FUNCTION_BLOCK FB_Gr05AutoProcedure
(*

The function block used to generate auto process..

Constructor: 		Patryk Panylo
Company:		E. Riexinger GmbH
Date:			28.04.2015
Version:			1.00

Date:			Revision:		Who:				Comment
dd.mm.yyyy		x.xx			Initials			comment

*)
VAR_INPUT
	(* Input variables / Eingang Variablen *)
	bEnable						:BOOL;						(* Enable FB signal *)
	bExecute					:BOOL;						(* Auto procedure execute *)
	bReleaseNextStep			:BOOL;						(* Auto procedure release next step *)
	bInterrupt					:BOOL;						(* Auto procedure interrupt *)
	SFCInit						:BOOL; 						(* System Flag:: INIT Flag *)
	bFirstTime					:BOOL;
END_VAR
VAR_OUTPUT
	(* Output variables / Ausgang Variablen *)
	bDone						:BOOL;						(* Program done *)
	bInterrupted					:BOOL;						(* Program interrupted *)
	bBusy						:BOOL;						(* Program busy *)
	bError						:BOOL;						(* Program error *)
	udnErrorNo					:UDINT;						(* Error number *)
	SFCError						:BOOL; 						(* System Flag: Timeout in this step *)
END_VAR
VAR_IN_OUT
	(* Input Output variables / Ausgang Variablen *)

END_VAR
VAR
	(* Enummerations *)

	(* Variables *)
	lrClamp1Pos					:LREAL;
	lrClamp1PosCache			:LREAL;
	lrClamp1PosPipeEnd			:LREAL;
	lrClamp2Pos					:LREAL;
	lrActRemoveLength			:LREAL;
	bPipeEndDetected			:BOOL;
	unProcessCounter				:UINT;
	lrActSawingLength				:LREAL;
	lrActSawingAngle				:LREAL;

	lrDistPipeBeginSawBand		:LREAL;

	bSafetyDistEnable			:BOOL; 						(* Safety distance between Clamp1 & 2 increase *)
	bErrorPipeBeginNoDetected	:BOOL;						(* Pipe begin no detected *)
	bErrorPipeEndNoDetected		:BOOL;						(* Pipe end no detected *)
	bErrorCollisionDetected		:BOOL;						(* Collision detected *)
	bWarningPipeBeginNoDetected	:BOOL;						(* Pipe begin no detected *)

	SFCCurrentStep				:STRING;					(* Name des aktiven Schritts *)

	(* References *)

	(* Interfaces *)

	(* Instances *)
	rtPipeBeginIdentify			:R_TRIG;
	rtPipeEndIdentify				:R_TRIG;
END_VAR

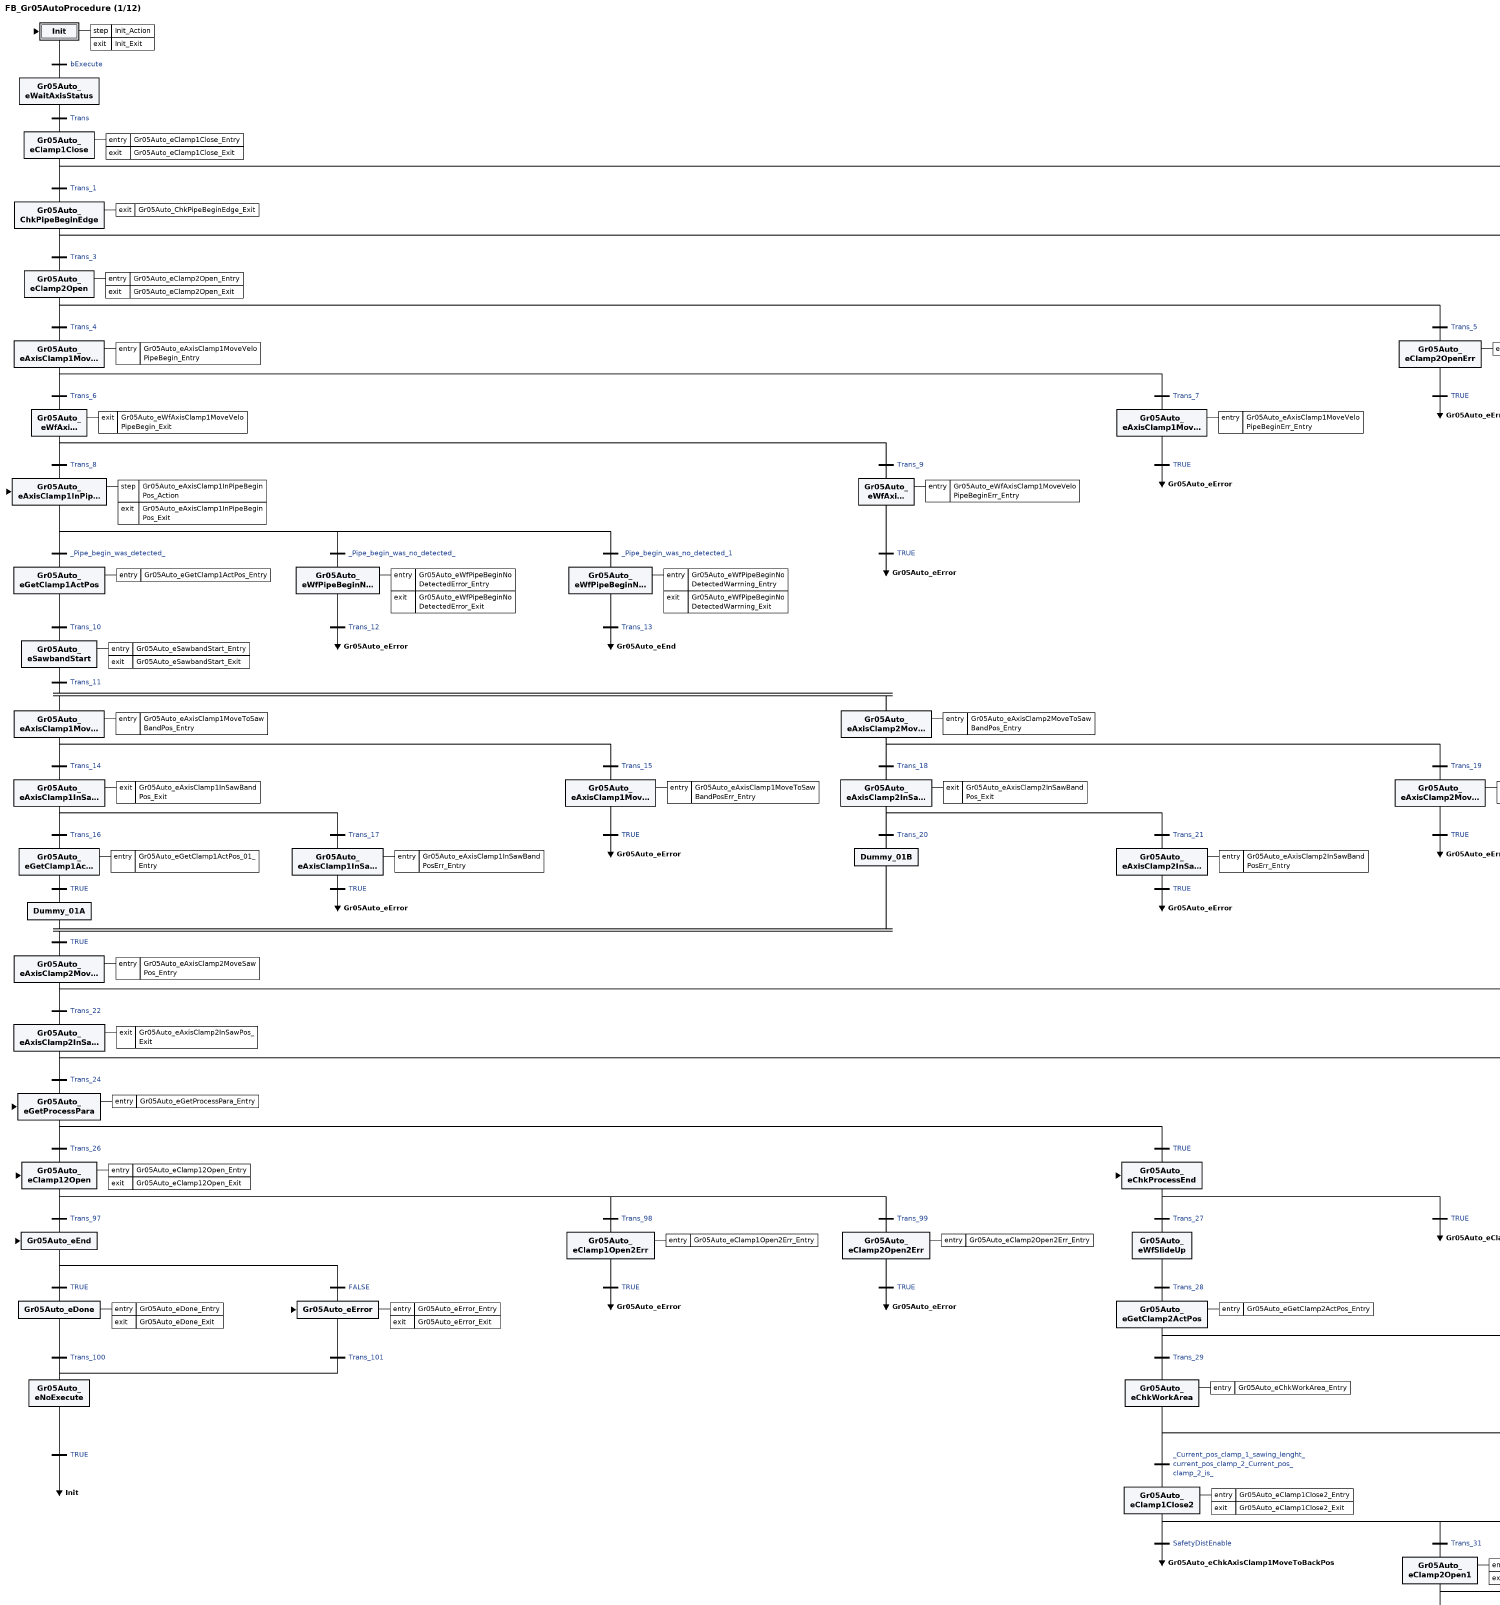
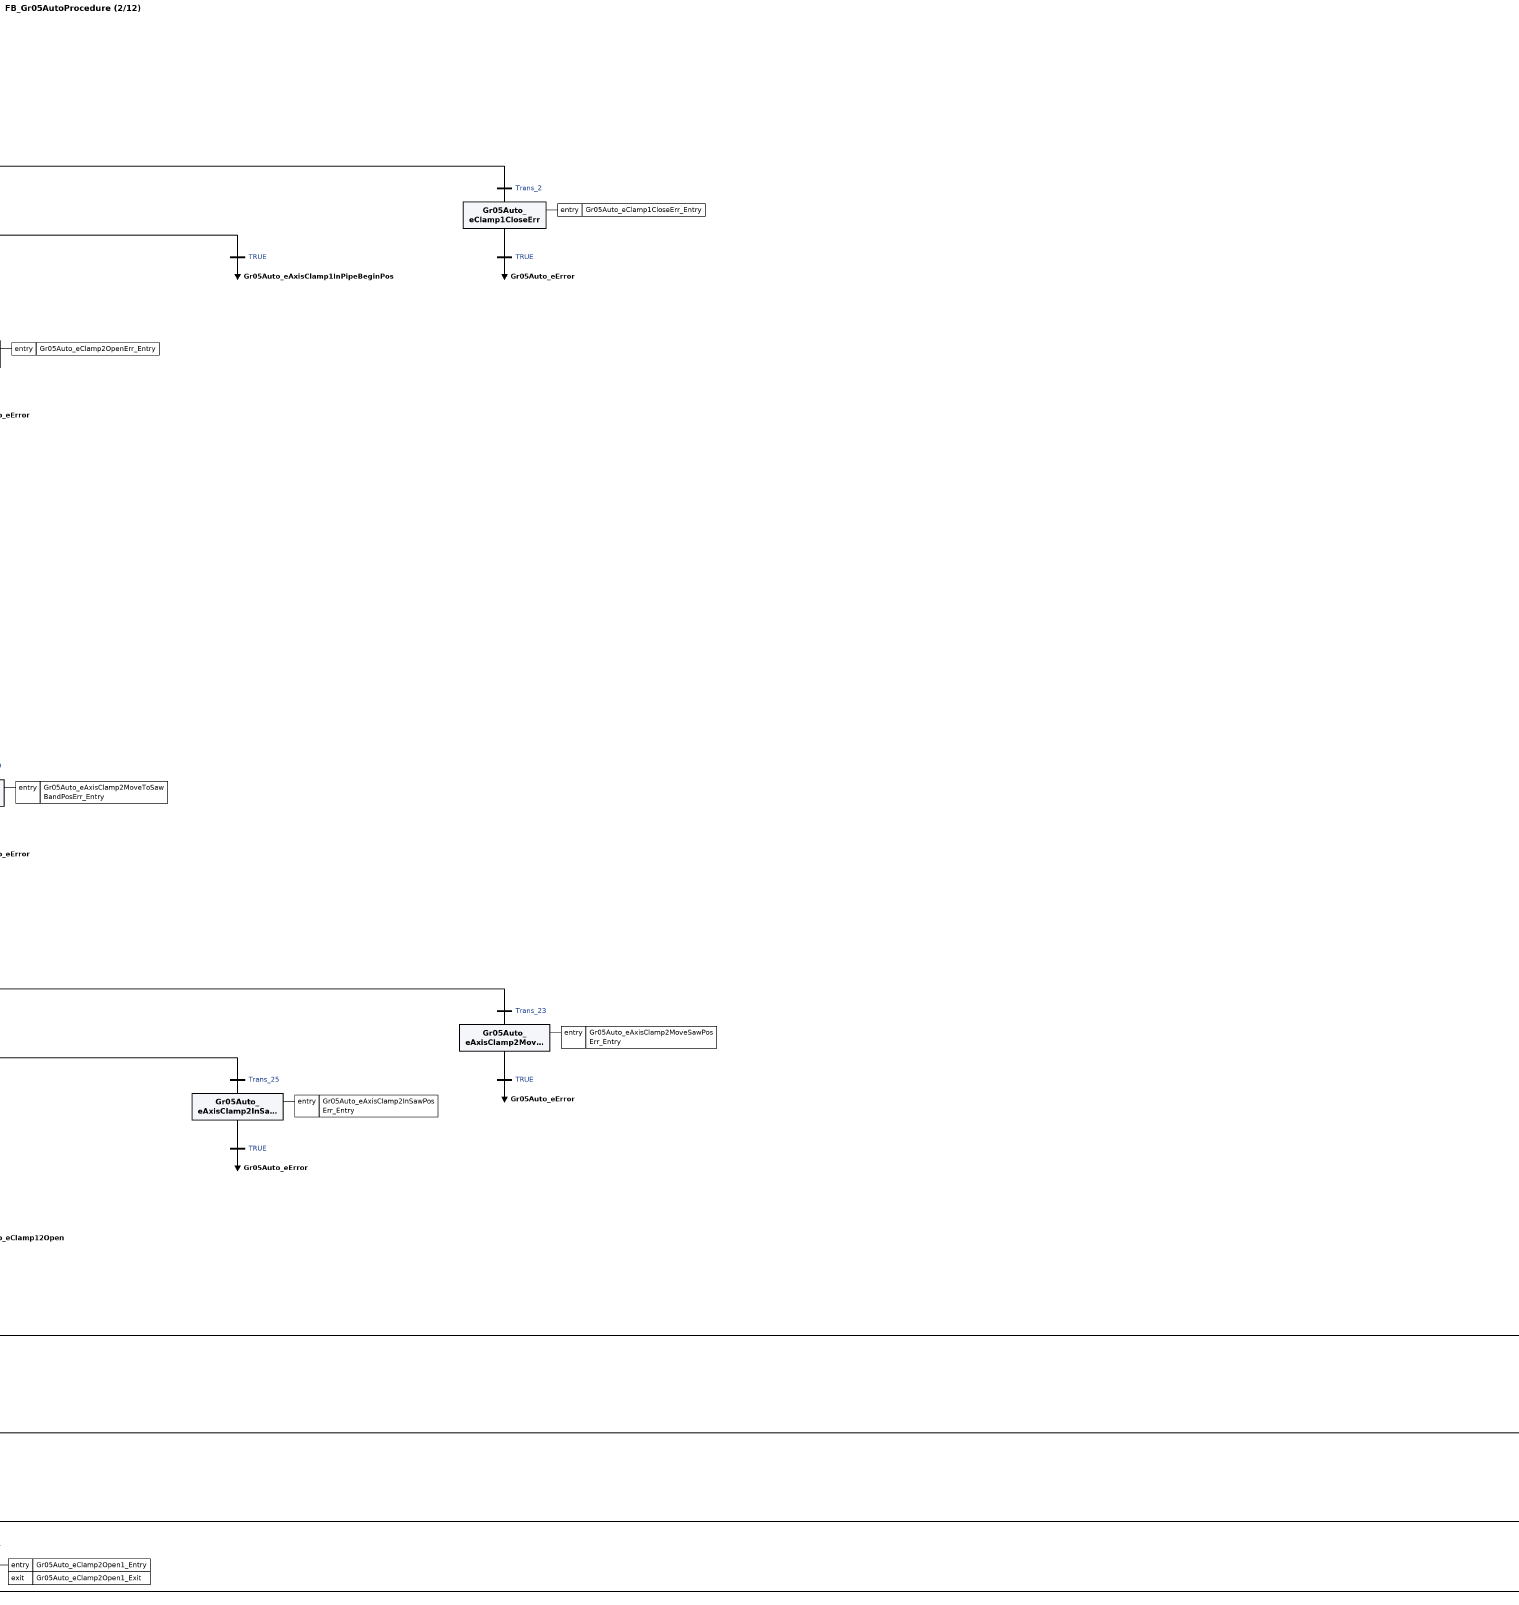
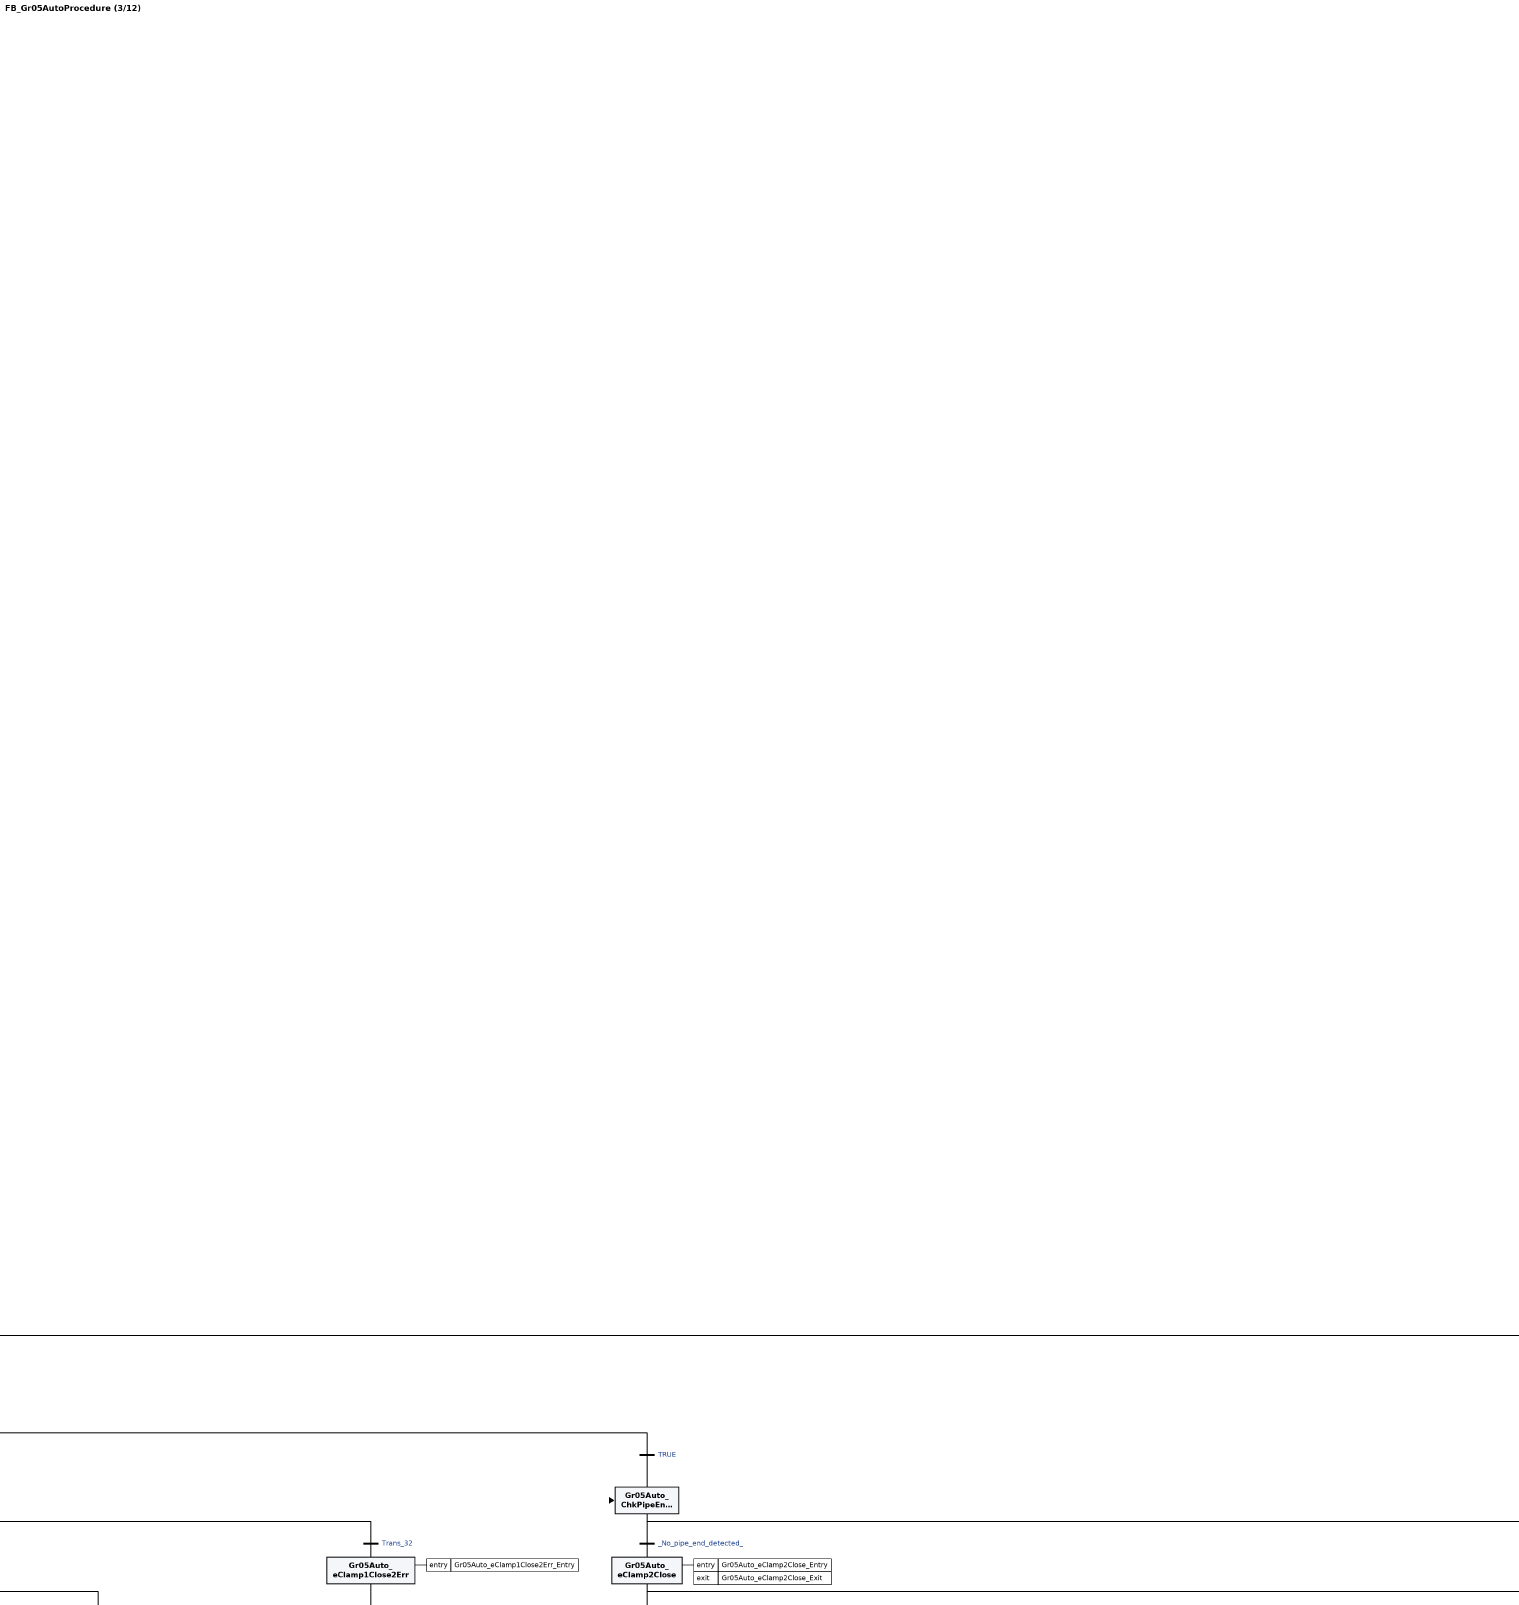
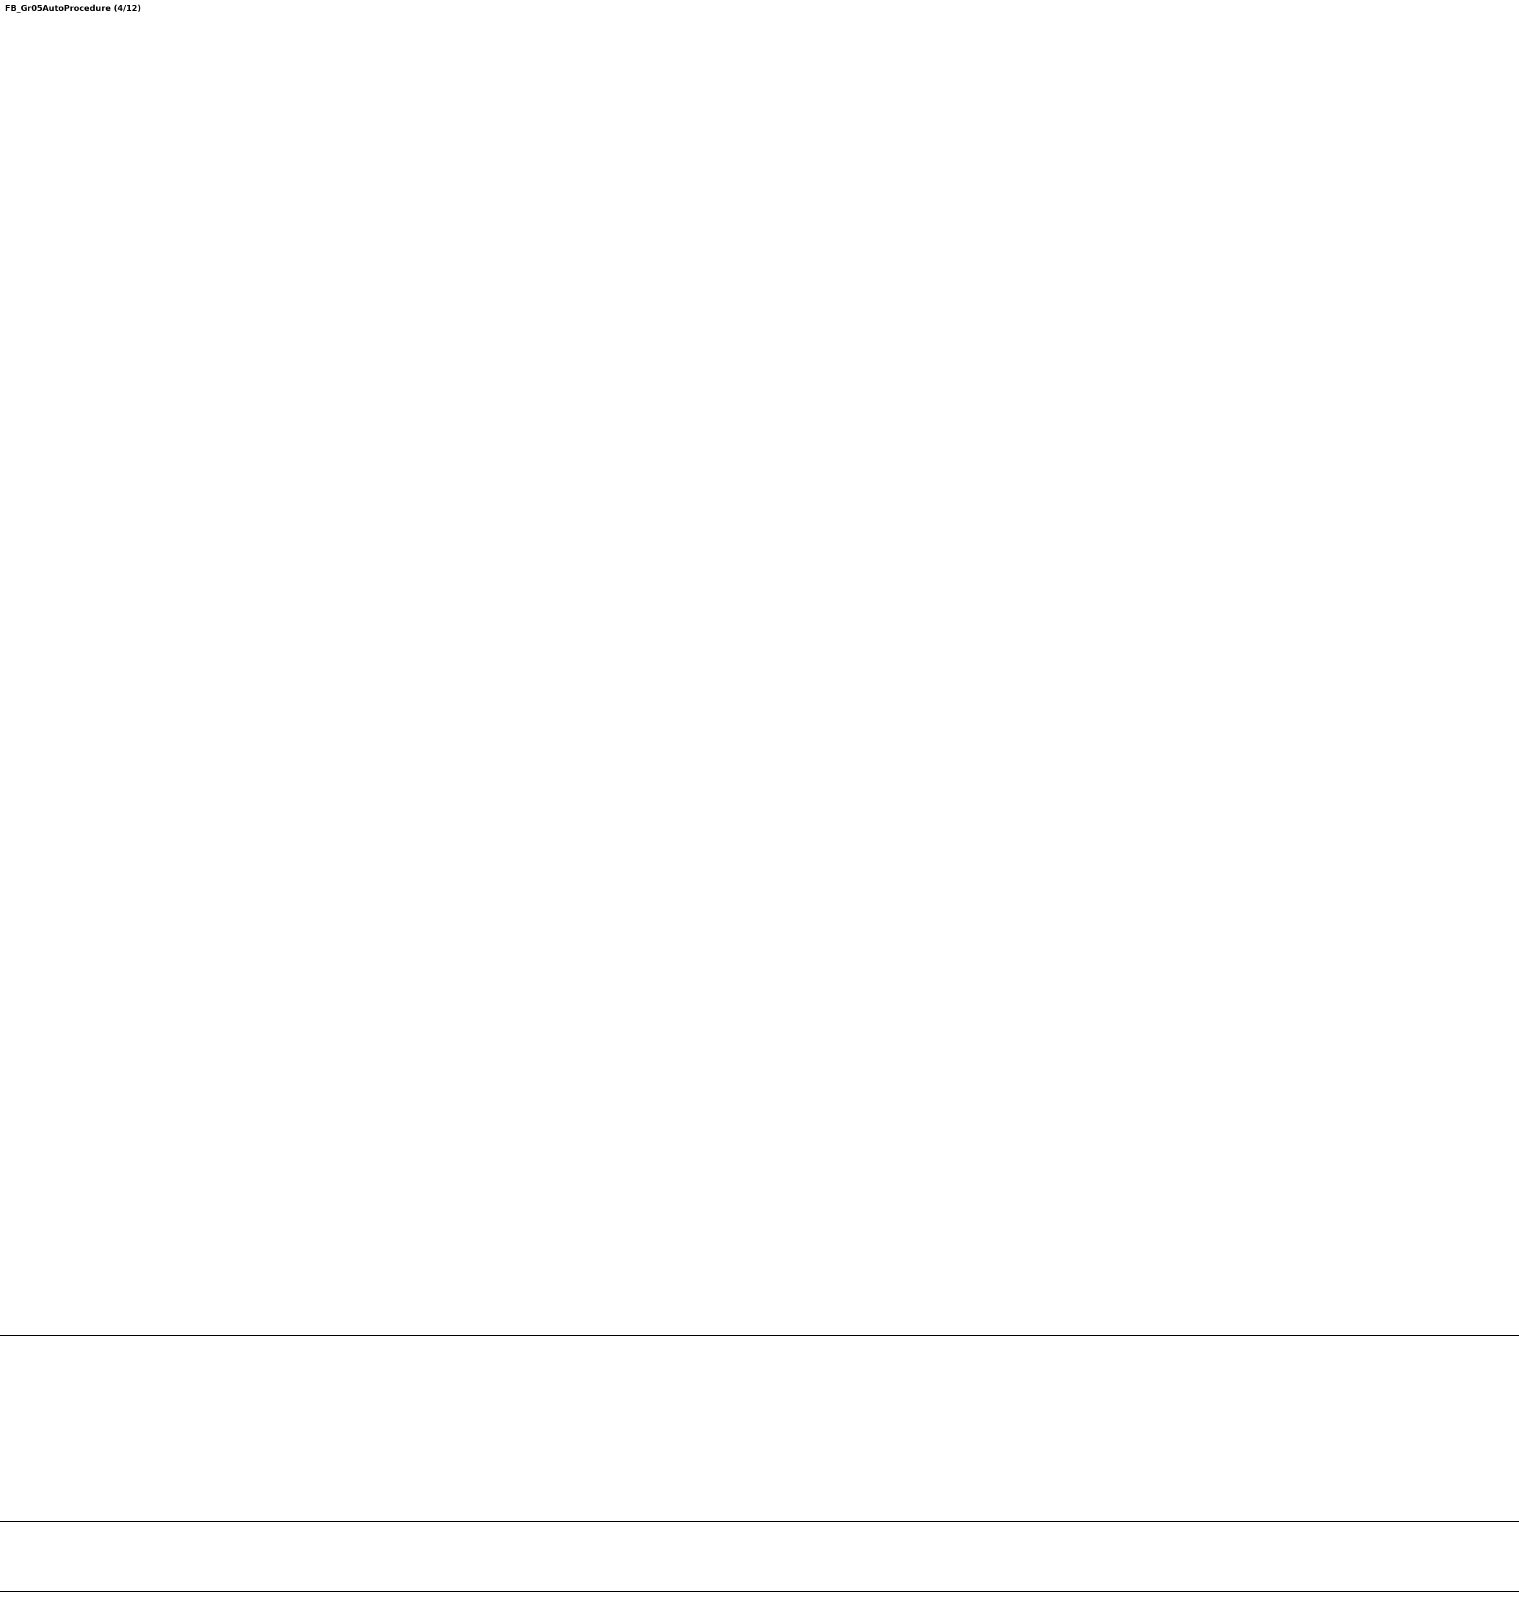
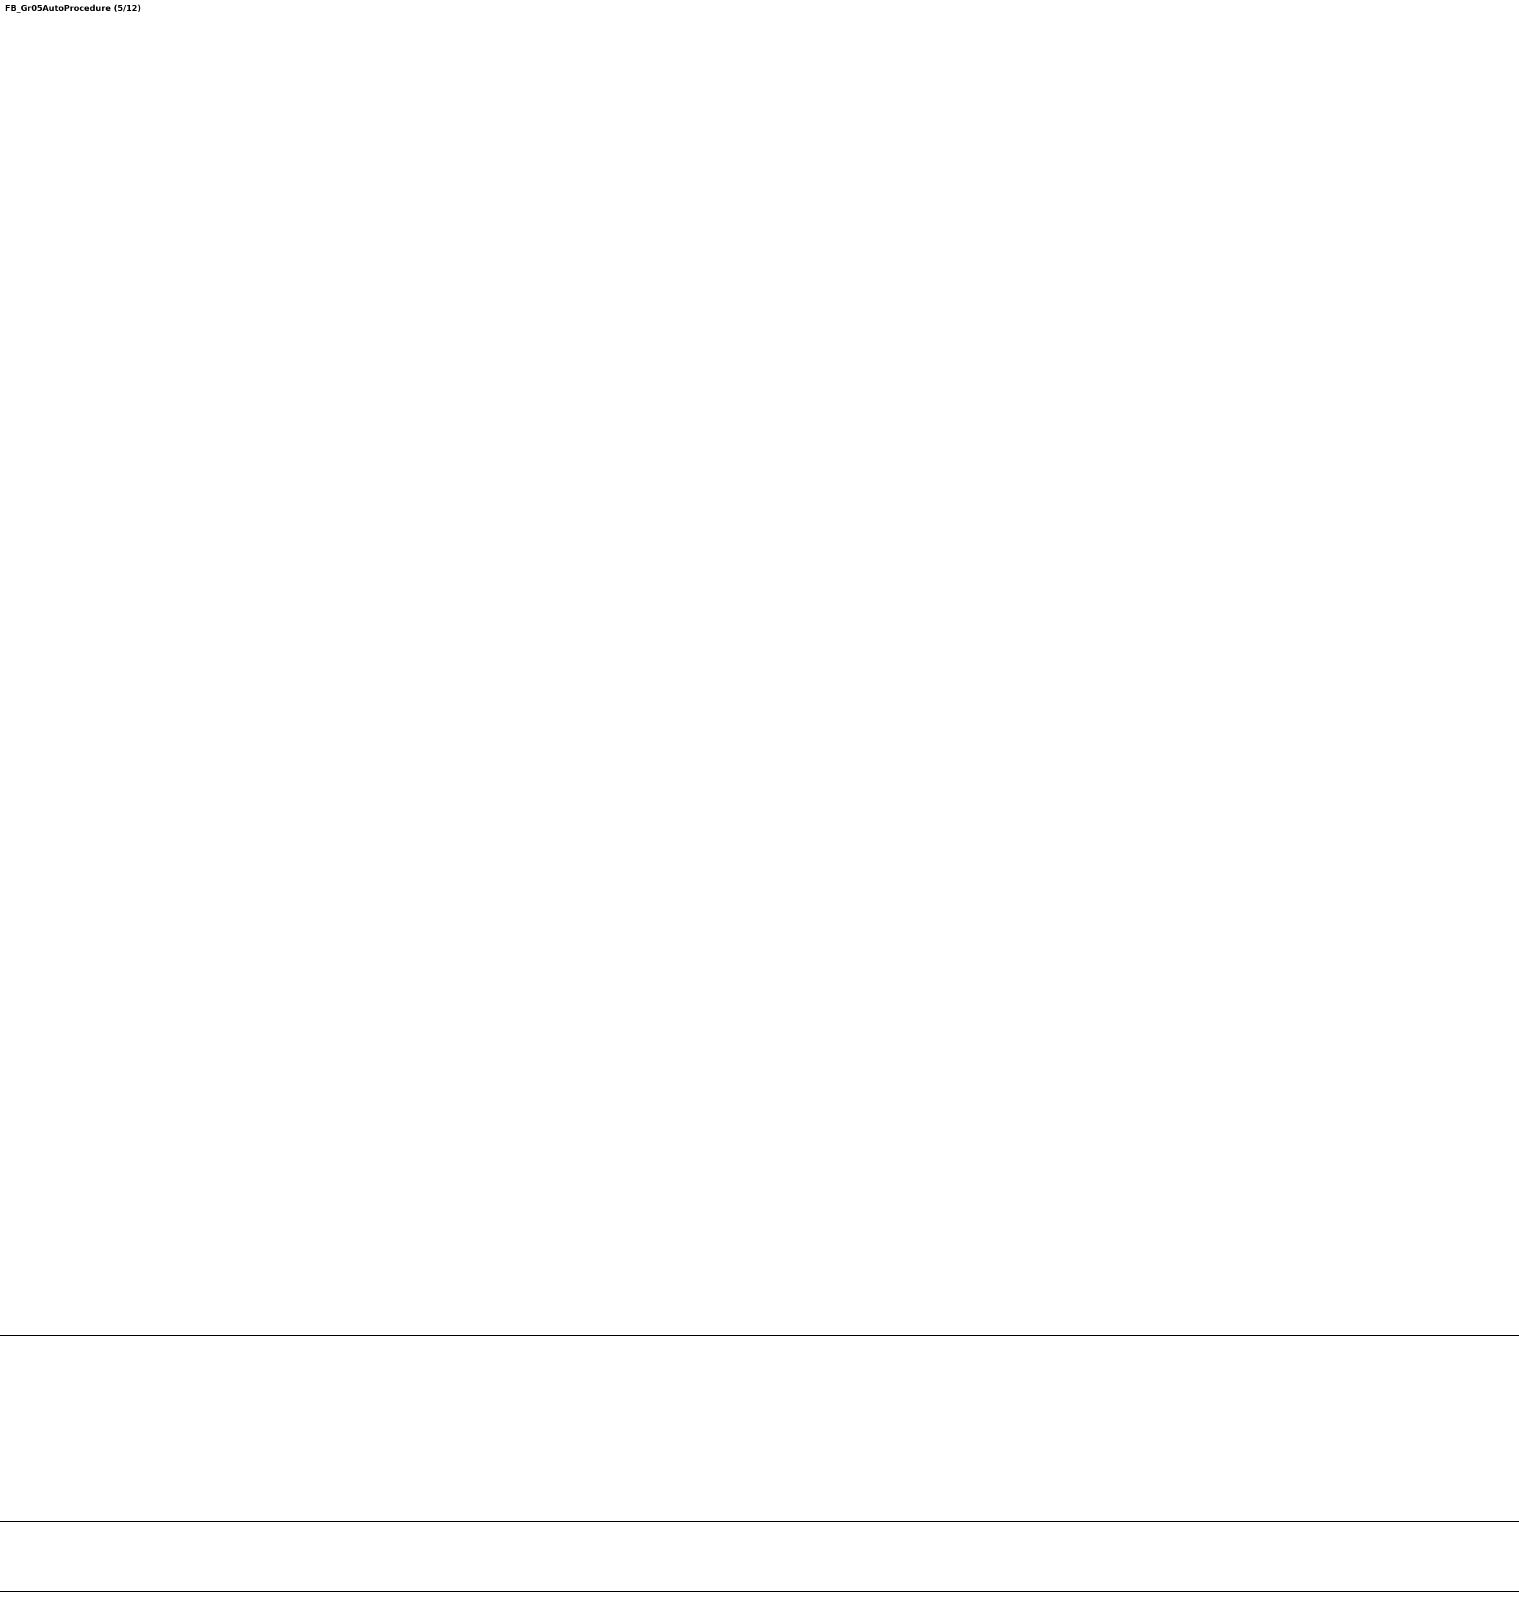
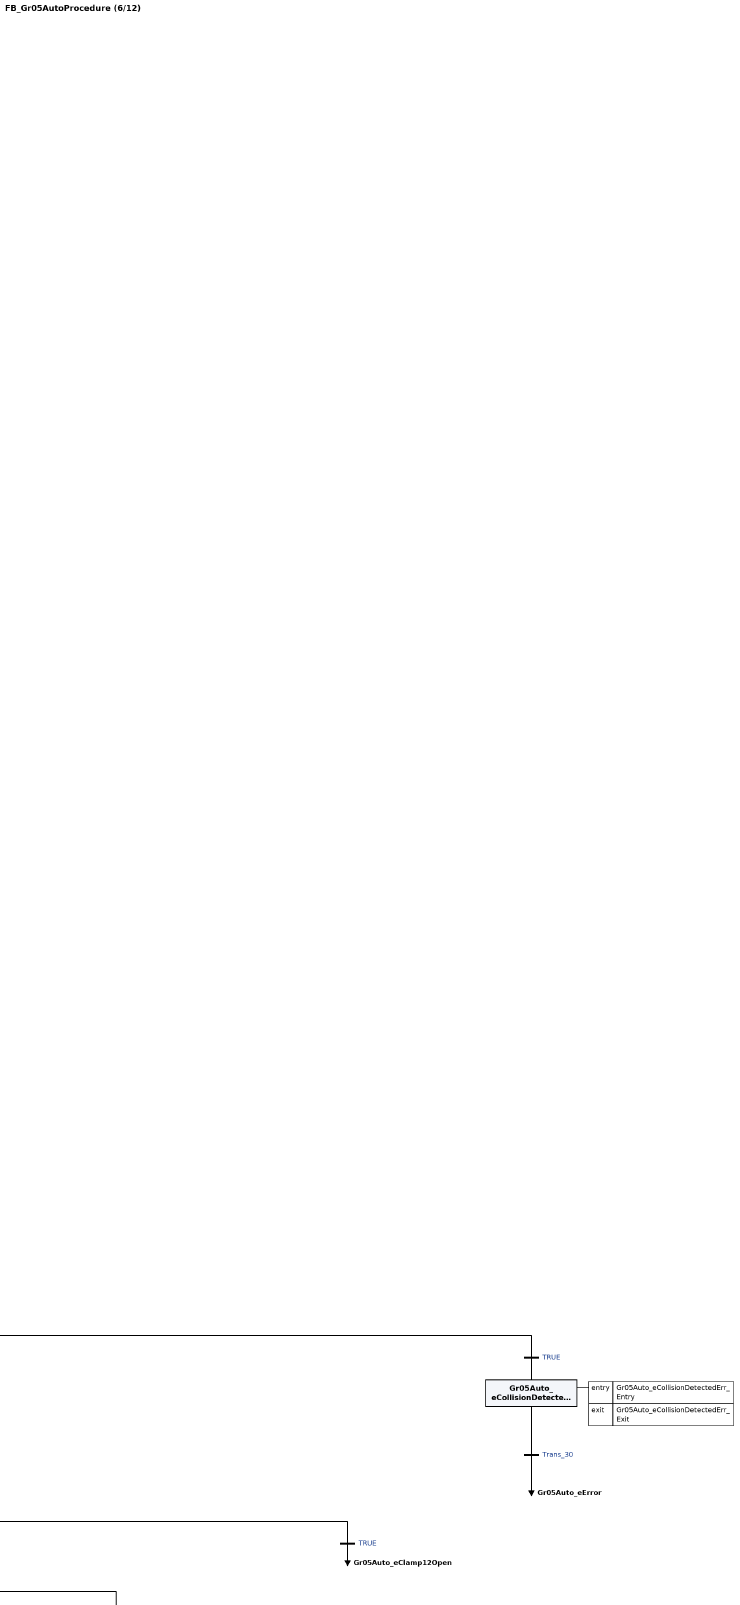
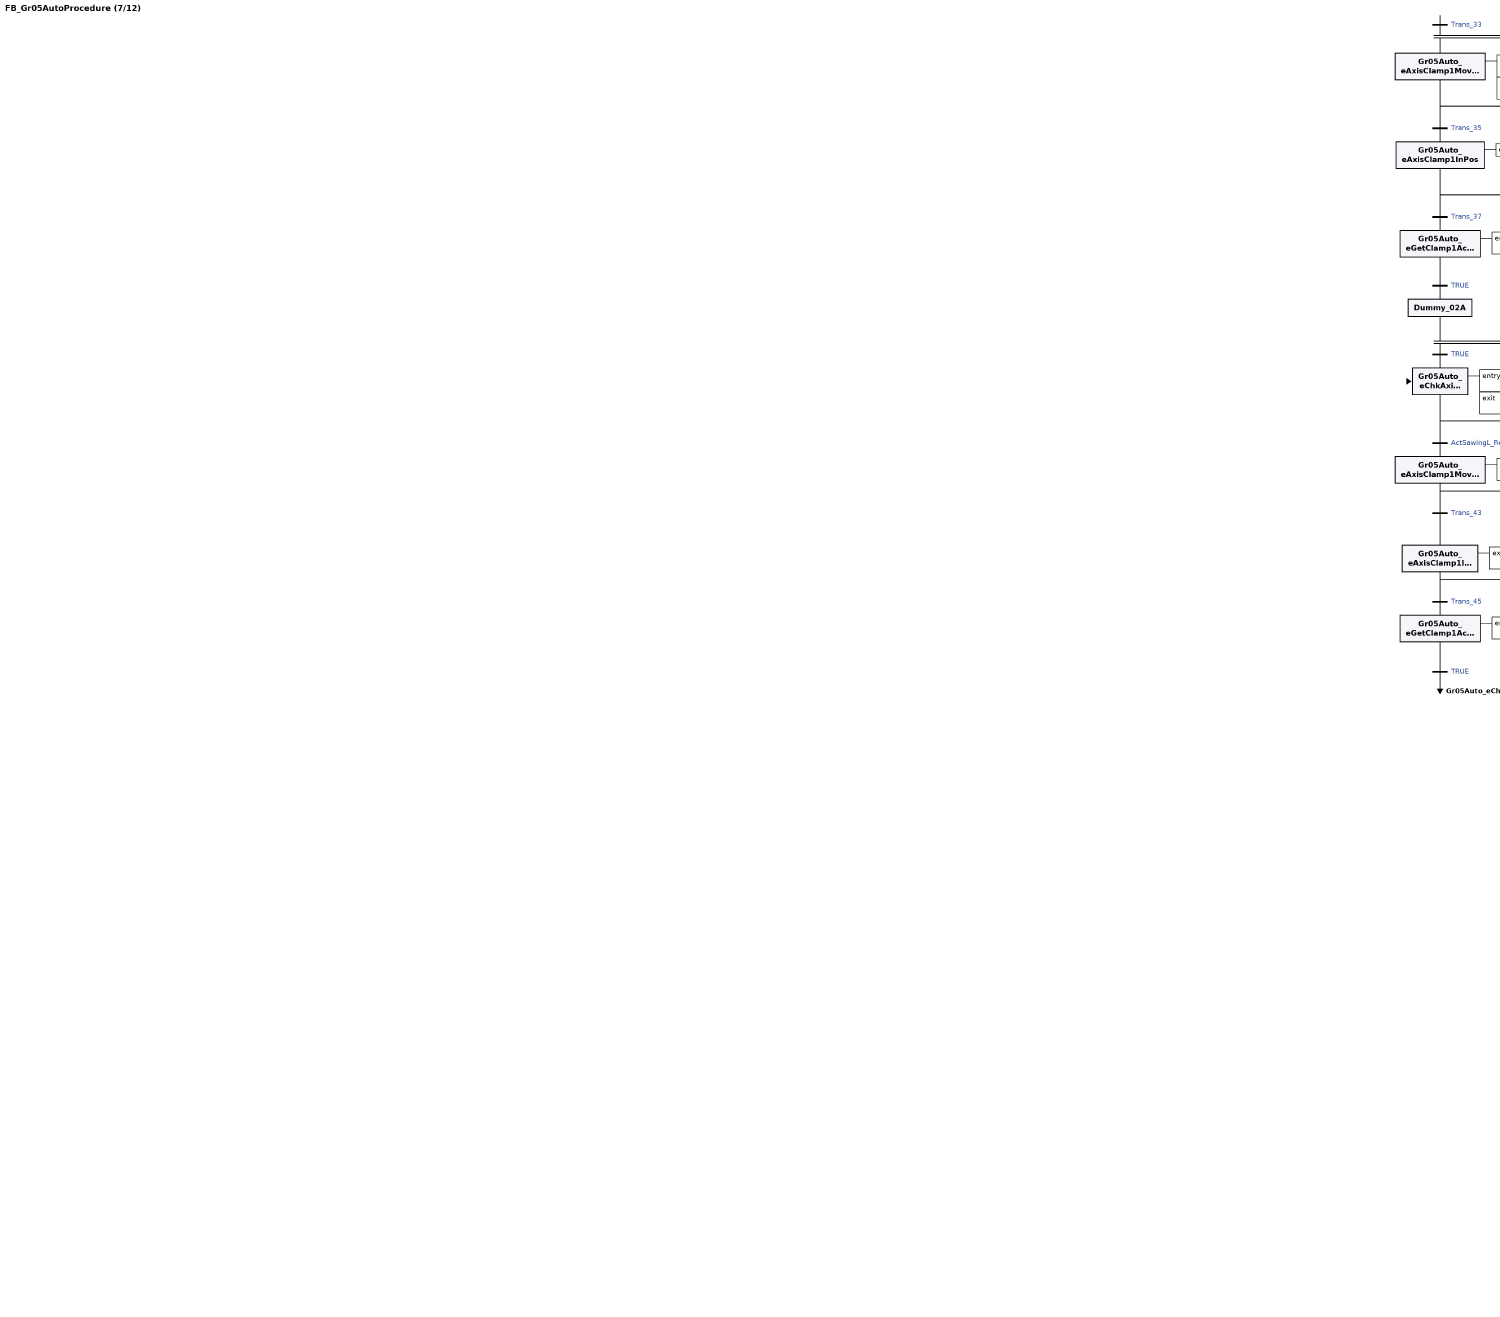
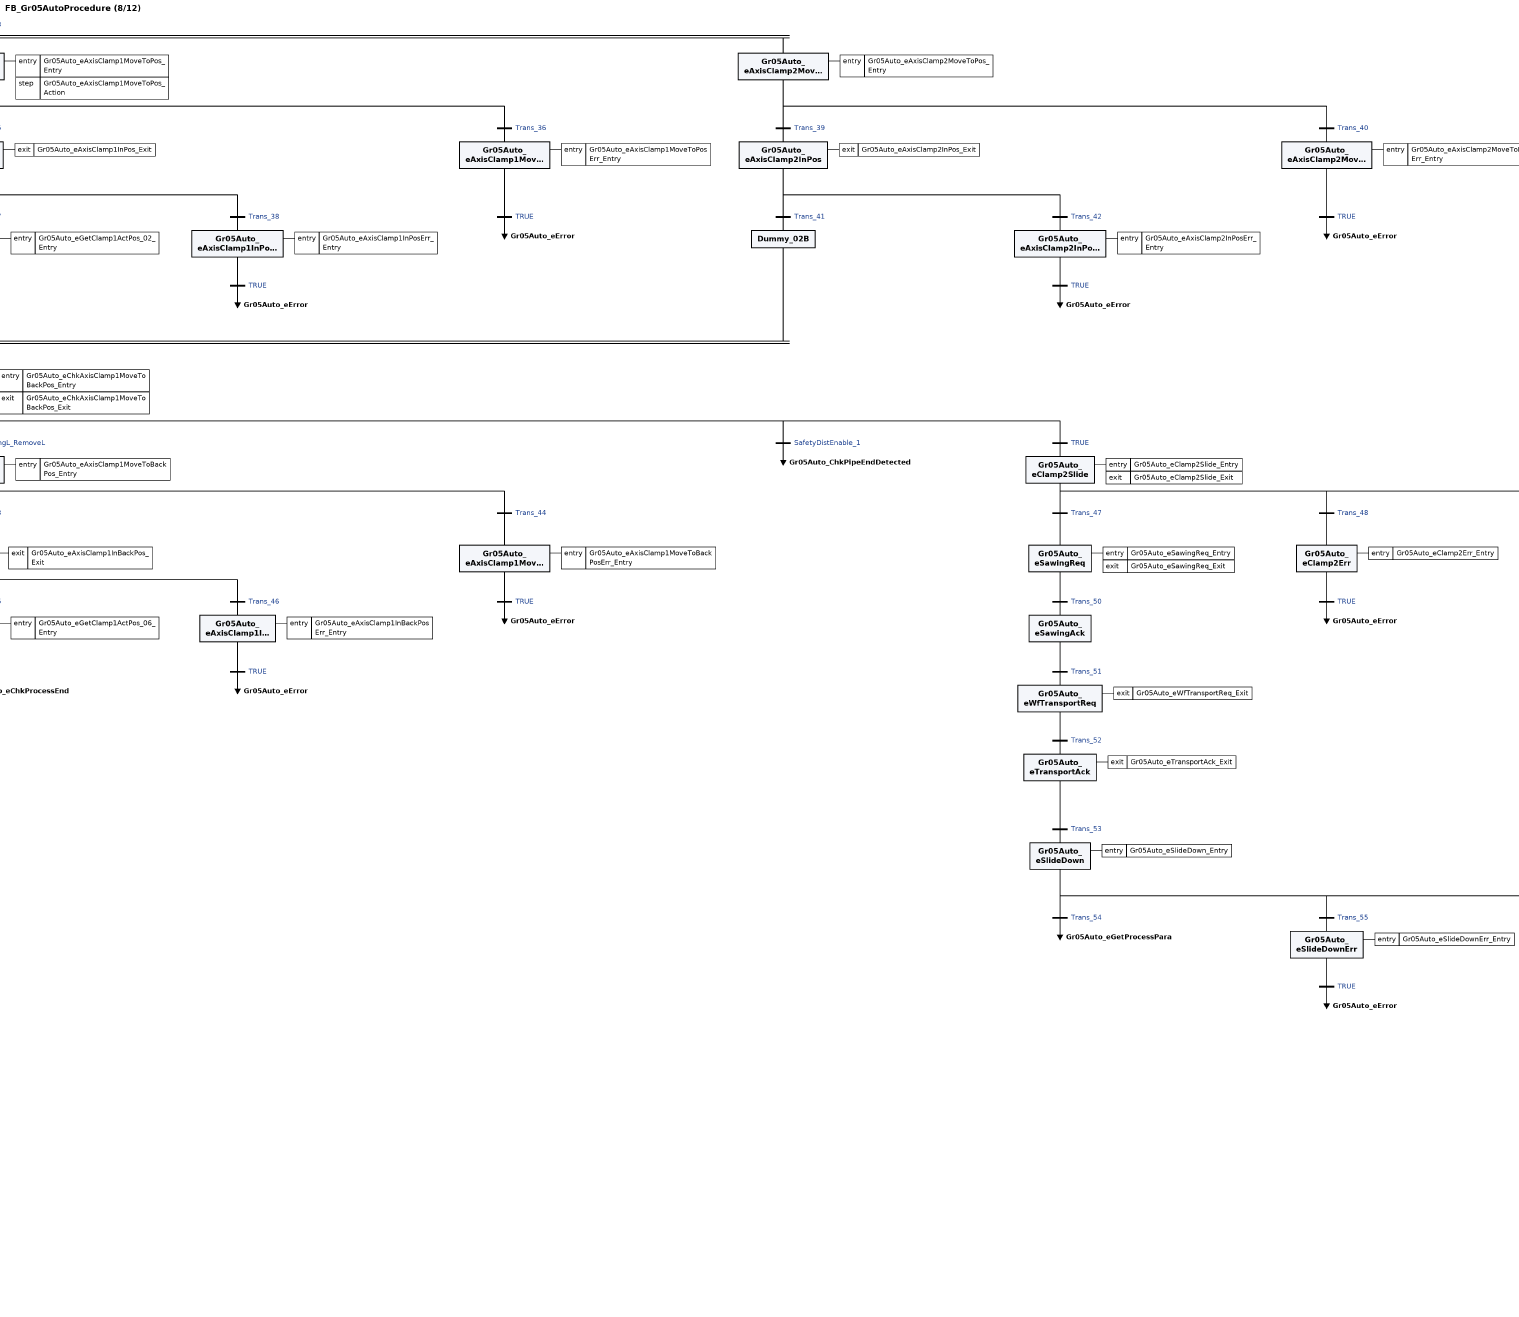
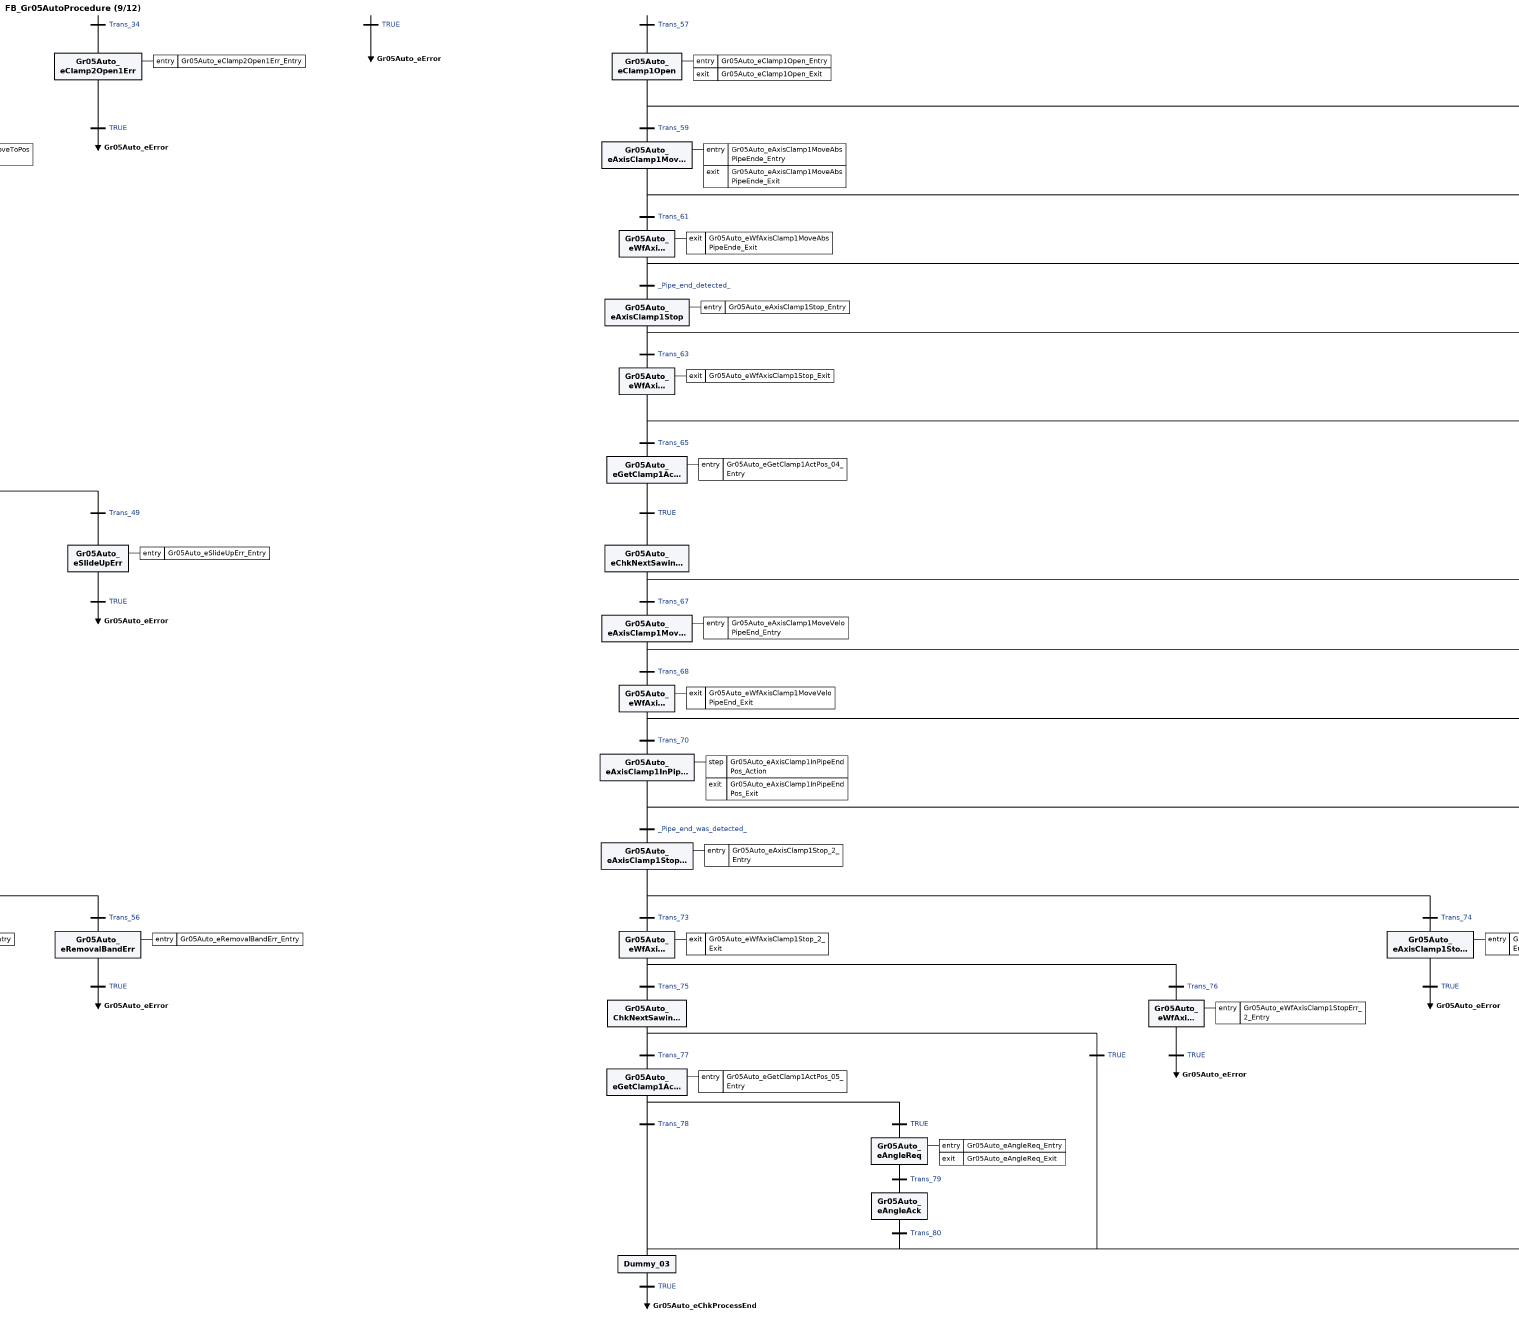
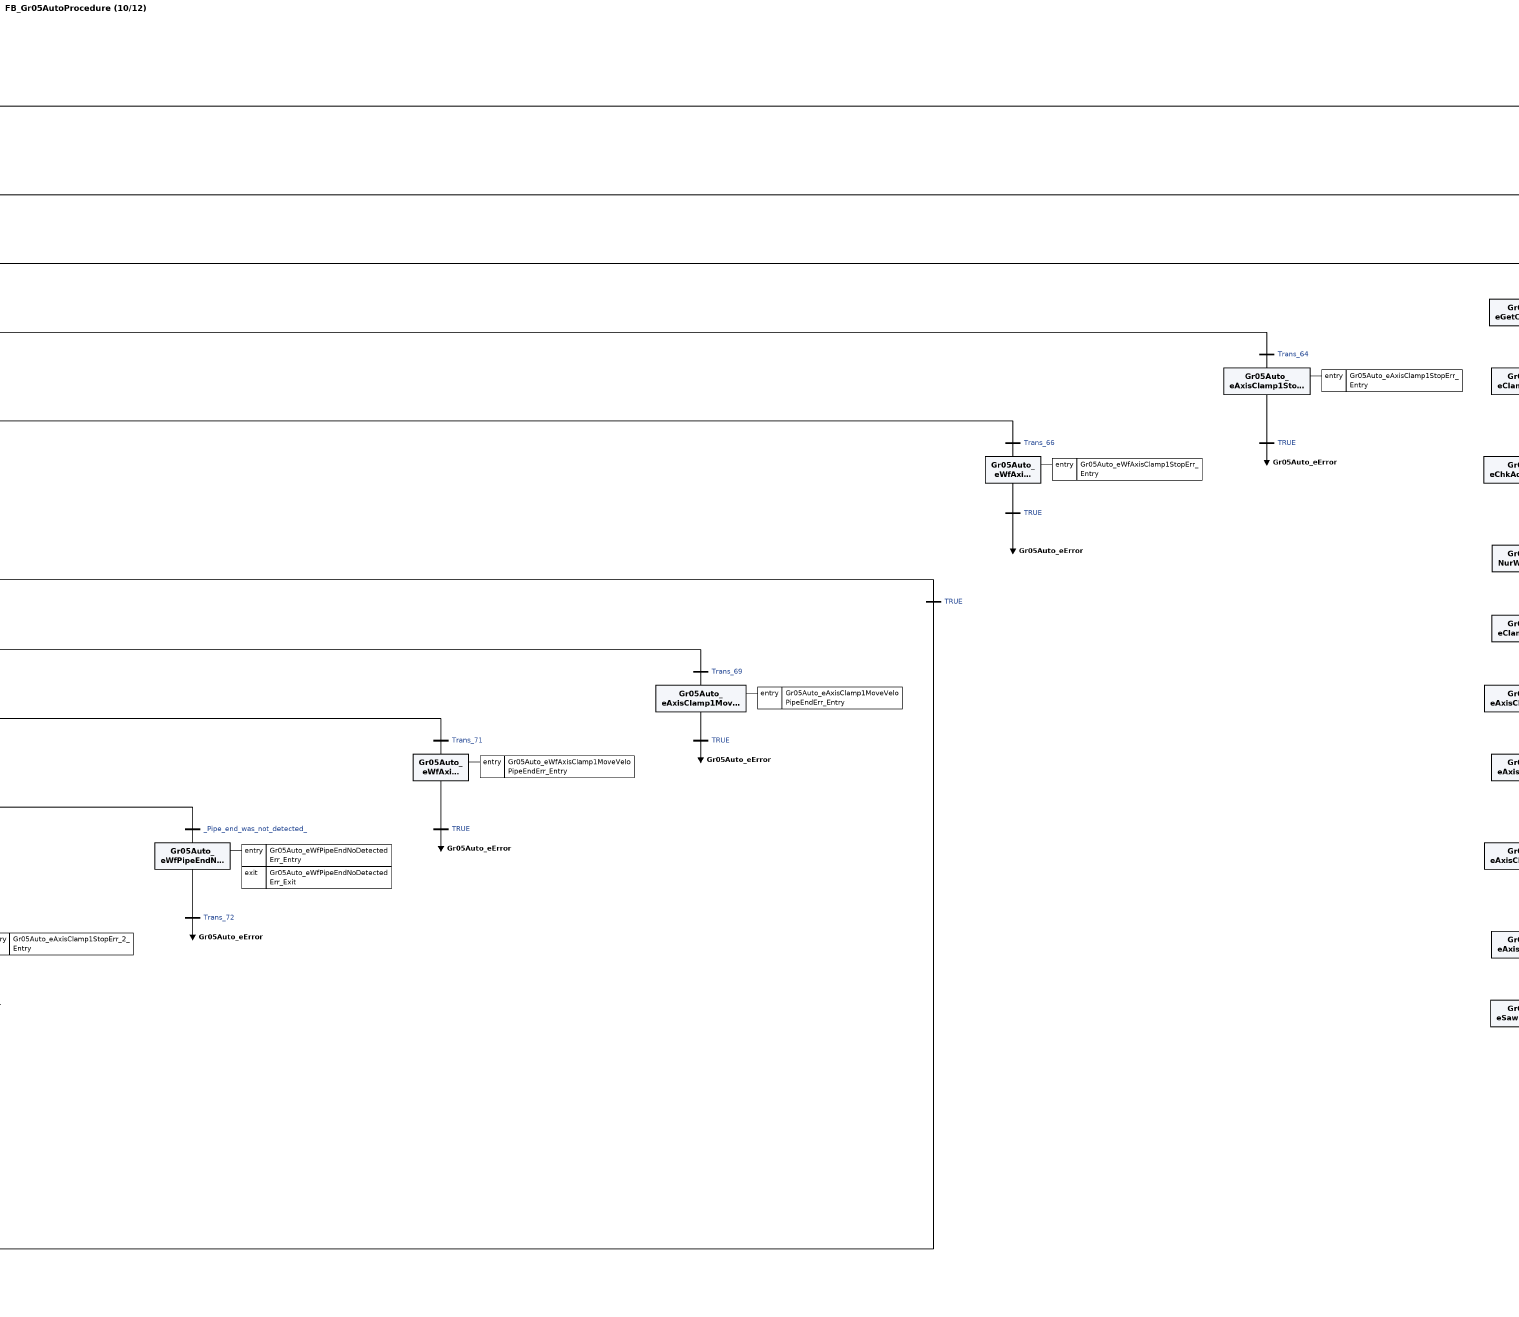
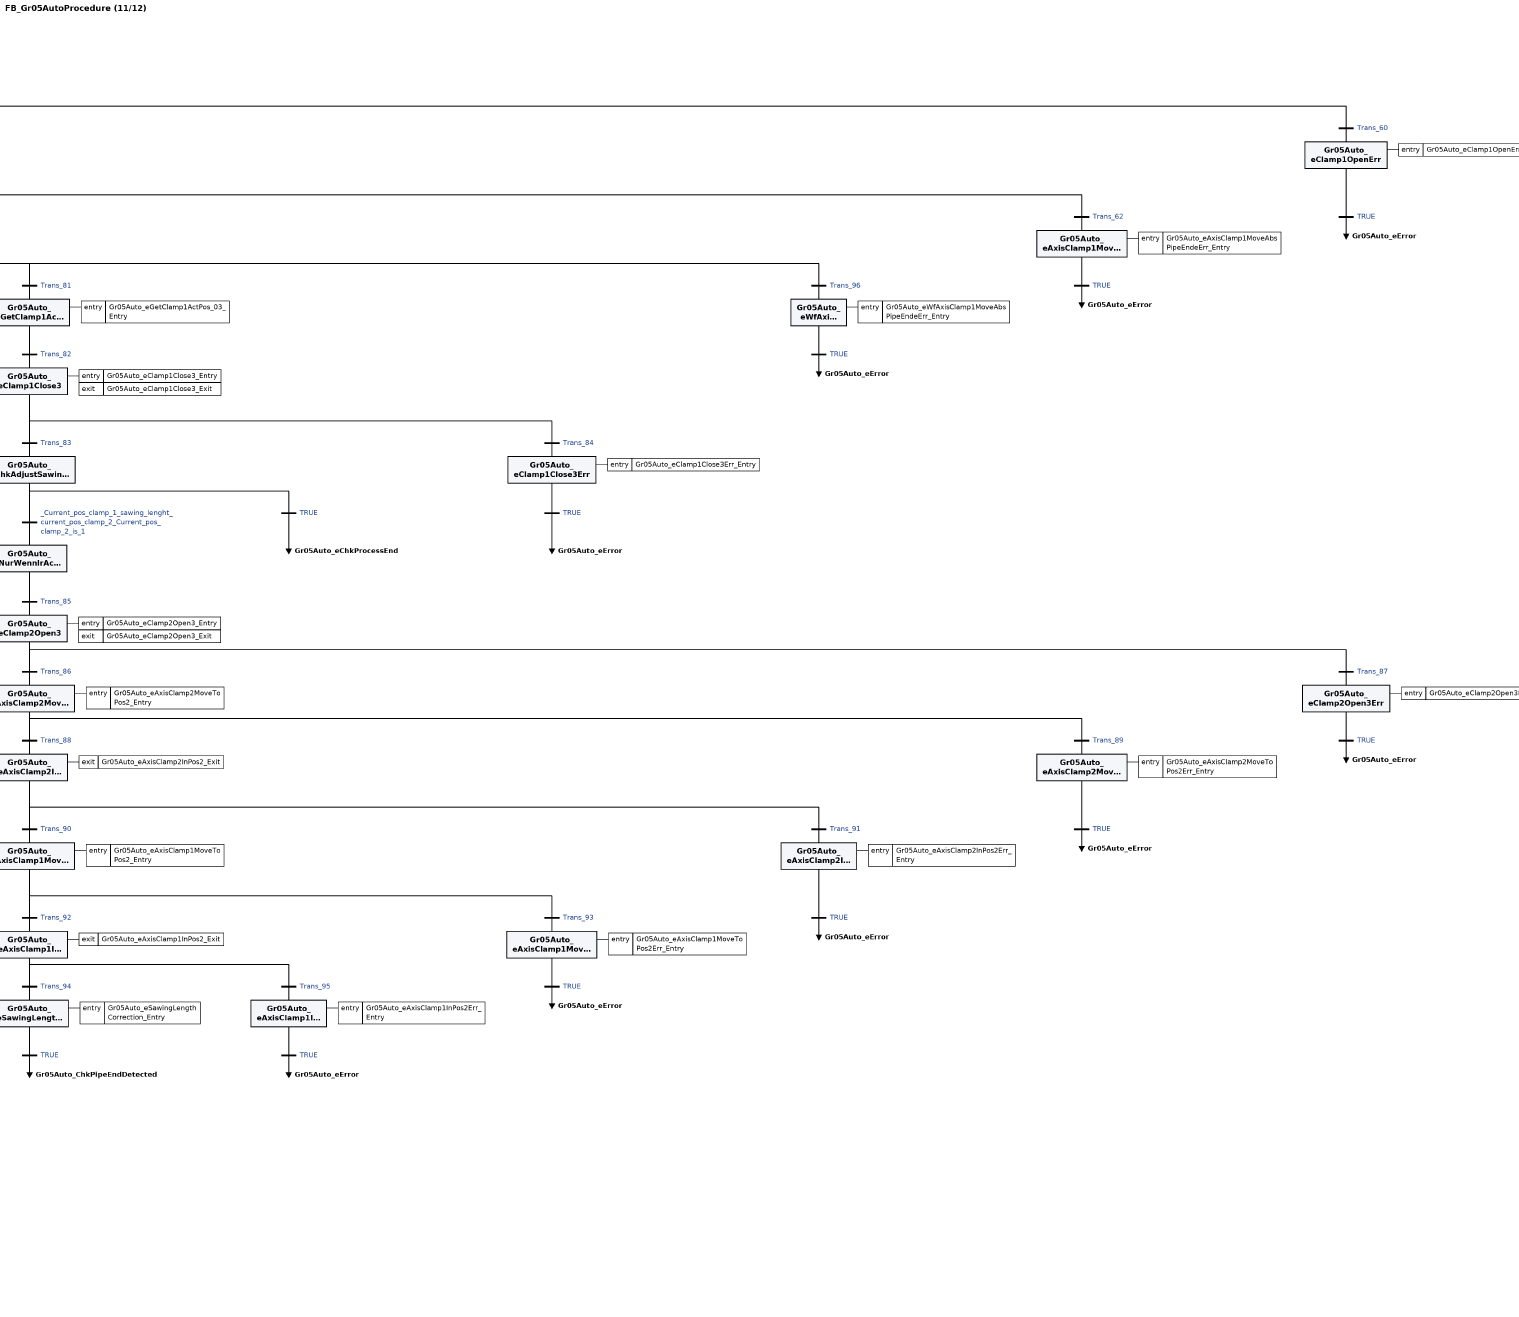
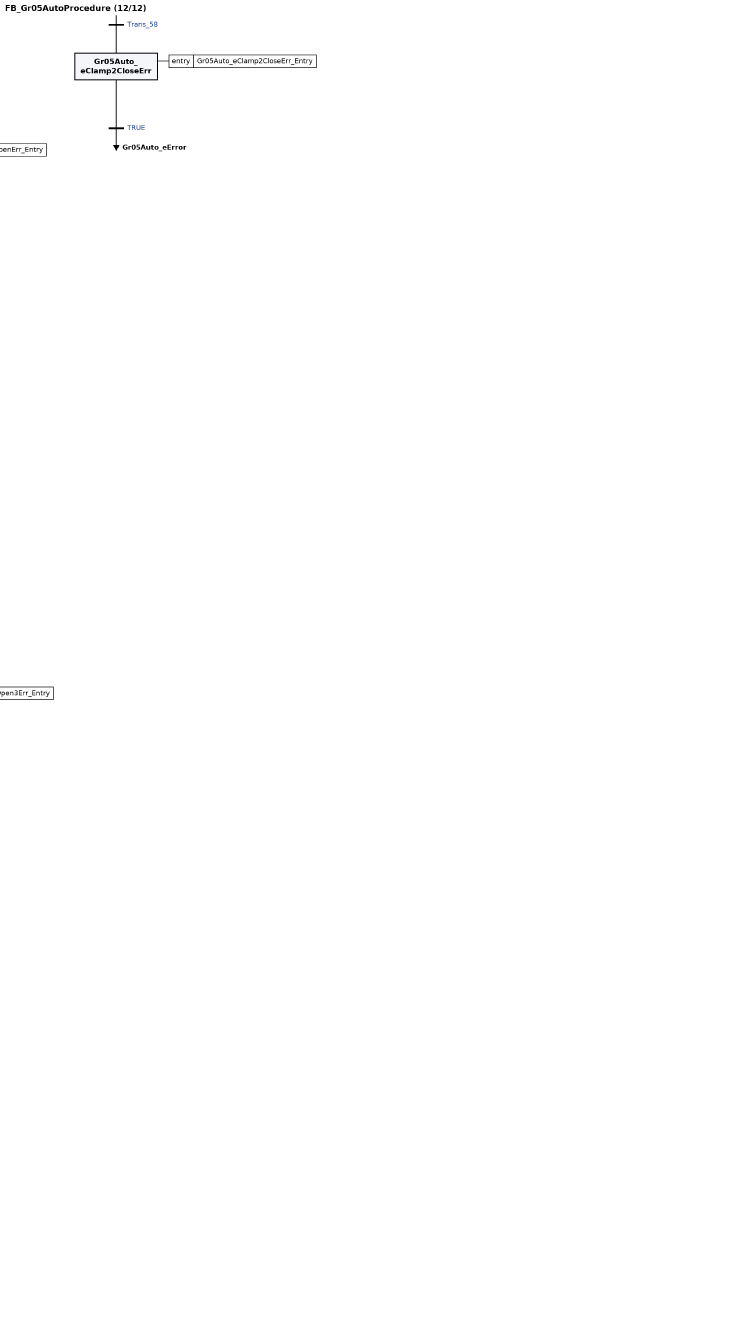
INITIAL_STEP Init:
    Init_Action(N);  // step action
    Init_Exit(P0);  // exit action
END_STEP
TRANSITION FROM Init TO Gr05Auto_eWaitAxisStatus
    := bExecute;
END_TRANSITION
STEP Gr05Auto_eWaitAxisStatus:
END_STEP
TRANSITION FROM Gr05Auto_eWaitAxisStatus TO Gr05Auto_eClamp1Close
    := Trans;
END_TRANSITION
STEP Gr05Auto_eClamp1Close:
    Gr05Auto_eClamp1Close_Entry(P1);  // entry action
    Gr05Auto_eClamp1Close_Exit(P0);  // exit action
END_STEP
TRANSITION FROM Gr05Auto_eClamp1Close TO Gr05Auto_ChkPipeBeginEdge
    := Trans_1;
END_TRANSITION
TRANSITION FROM Gr05Auto_eClamp1Close TO Gr05Auto_eClamp1CloseErr
    := Trans_2;
END_TRANSITION
STEP Gr05Auto_eClamp1CloseErr:
    Gr05Auto_eClamp1CloseErr_Entry(P1);  // entry action
END_STEP
TRANSITION FROM Gr05Auto_eClamp1CloseErr TO Gr05Auto_eError
    := TRUE;
END_TRANSITION
STEP Gr05Auto_ChkPipeBeginEdge:
    Gr05Auto_ChkPipeBeginEdge_Exit(P0);  // exit action
END_STEP
TRANSITION FROM Gr05Auto_ChkPipeBeginEdge TO Gr05Auto_eClamp2Open
    := Trans_3;
END_TRANSITION
TRANSITION FROM Gr05Auto_ChkPipeBeginEdge TO Gr05Auto_eAxisClamp1InPipeBeginPos
    := TRUE;
END_TRANSITION
STEP Gr05Auto_eClamp2Open:
    Gr05Auto_eClamp2Open_Entry(P1);  // entry action
    Gr05Auto_eClamp2Open_Exit(P0);  // exit action
END_STEP
TRANSITION FROM Gr05Auto_eClamp2Open TO Gr05Auto_eAxisClamp1MoveVeloPipeBegin
    := Trans_4;
END_TRANSITION
TRANSITION FROM Gr05Auto_eClamp2Open TO Gr05Auto_eClamp2OpenErr
    := Trans_5;
END_TRANSITION
STEP Gr05Auto_eClamp2OpenErr:
    Gr05Auto_eClamp2OpenErr_Entry(P1);  // entry action
END_STEP
TRANSITION FROM Gr05Auto_eClamp2OpenErr TO Gr05Auto_eError
    := TRUE;
END_TRANSITION
STEP Gr05Auto_eAxisClamp1MoveVeloPipeBegin:
    Gr05Auto_eAxisClamp1MoveVeloPipeBegin_Entry(P1);  // entry action
END_STEP
TRANSITION FROM Gr05Auto_eAxisClamp1MoveVeloPipeBegin TO Gr05Auto_eWfAxisClamp1MoveVeloPipeBegin
    := Trans_6;
END_TRANSITION
TRANSITION FROM Gr05Auto_eAxisClamp1MoveVeloPipeBegin TO Gr05Auto_eAxisClamp1MoveVeloPipeBeginErr
    := Trans_7;
END_TRANSITION
STEP Gr05Auto_eAxisClamp1MoveVeloPipeBeginErr:
    Gr05Auto_eAxisClamp1MoveVeloPipeBeginErr_Entry(P1);  // entry action
END_STEP
TRANSITION FROM Gr05Auto_eAxisClamp1MoveVeloPipeBeginErr TO Gr05Auto_eError
    := TRUE;
END_TRANSITION
STEP Gr05Auto_eWfAxisClamp1MoveVeloPipeBegin:
    Gr05Auto_eWfAxisClamp1MoveVeloPipeBegin_Exit(P0);  // exit action
END_STEP
TRANSITION FROM Gr05Auto_eWfAxisClamp1MoveVeloPipeBegin TO Gr05Auto_eAxisClamp1InPipeBeginPos
    := Trans_8;
END_TRANSITION
TRANSITION FROM Gr05Auto_eWfAxisClamp1MoveVeloPipeBegin TO Gr05Auto_eWfAxisClamp1MoveVeloPipeBeginErr
    := Trans_9;
END_TRANSITION
STEP Gr05Auto_eWfAxisClamp1MoveVeloPipeBeginErr:
    Gr05Auto_eWfAxisClamp1MoveVeloPipeBeginErr_Entry(P1);  // entry action
END_STEP
TRANSITION FROM Gr05Auto_eWfAxisClamp1MoveVeloPipeBeginErr TO Gr05Auto_eError
    := TRUE;
END_TRANSITION
STEP Gr05Auto_eAxisClamp1InPipeBeginPos:
    Gr05Auto_eAxisClamp1InPipeBeginPos_Action(N);  // step action
    Gr05Auto_eAxisClamp1InPipeBeginPos_Exit(P0);  // exit action
END_STEP
TRANSITION FROM Gr05Auto_eAxisClamp1InPipeBeginPos TO Gr05Auto_eGetClamp1ActPos
    := _Pipe_begin_was_detected_;
END_TRANSITION
STEP Gr05Auto_eGetClamp1ActPos:
    Gr05Auto_eGetClamp1ActPos_Entry(P1);  // entry action
END_STEP
TRANSITION FROM Gr05Auto_eGetClamp1ActPos TO Gr05Auto_eSawbandStart
    := Trans_10;
END_TRANSITION
STEP Gr05Auto_eSawbandStart:
    Gr05Auto_eSawbandStart_Entry(P1);  // entry action
    Gr05Auto_eSawbandStart_Exit(P0);  // exit action
END_STEP
TRANSITION FROM Gr05Auto_eSawbandStart TO (Gr05Auto_eAxisClamp1MoveToSawBandPos, Gr05Auto_eAxisClamp2MoveToSawBandPos)
    := Trans_11;
END_TRANSITION
TRANSITION FROM Gr05Auto_eAxisClamp1InPipeBeginPos TO Gr05Auto_eWfPipeBeginNoDetectedError
    := _Pipe_begin_was_no_detected_;
END_TRANSITION
STEP Gr05Auto_eWfPipeBeginNoDetectedError:
    Gr05Auto_eWfPipeBeginNoDetectedError_Entry(P1);  // entry action
    Gr05Auto_eWfPipeBeginNoDetectedError_Exit(P0);  // exit action
END_STEP
TRANSITION FROM Gr05Auto_eWfPipeBeginNoDetectedError TO Gr05Auto_eError
    := Trans_12;
END_TRANSITION
TRANSITION FROM Gr05Auto_eAxisClamp1InPipeBeginPos TO Gr05Auto_eWfPipeBeginNoDetectedWarrning
    := _Pipe_begin_was_no_detected_1;
END_TRANSITION
STEP Gr05Auto_eWfPipeBeginNoDetectedWarrning:
    Gr05Auto_eWfPipeBeginNoDetectedWarrning_Entry(P1);  // entry action
    Gr05Auto_eWfPipeBeginNoDetectedWarrning_Exit(P0);  // exit action
END_STEP
TRANSITION FROM Gr05Auto_eWfPipeBeginNoDetectedWarrning TO Gr05Auto_eEnd
    := Trans_13;
END_TRANSITION
STEP Gr05Auto_eAxisClamp1MoveToSawBandPos:
    Gr05Auto_eAxisClamp1MoveToSawBandPos_Entry(P1);  // entry action
END_STEP
TRANSITION FROM Gr05Auto_eAxisClamp1MoveToSawBandPos TO Gr05Auto_eAxisClamp1InSawBandPos
    := Trans_14;
END_TRANSITION
TRANSITION FROM Gr05Auto_eAxisClamp1MoveToSawBandPos TO Gr05Auto_eAxisClamp1MoveToSawBandPosErr
    := Trans_15;
END_TRANSITION
STEP Gr05Auto_eAxisClamp1MoveToSawBandPosErr:
    Gr05Auto_eAxisClamp1MoveToSawBandPosErr_Entry(P1);  // entry action
END_STEP
TRANSITION FROM Gr05Auto_eAxisClamp1MoveToSawBandPosErr TO Gr05Auto_eError
    := TRUE;
END_TRANSITION
STEP Gr05Auto_eAxisClamp1InSawBandPos:
    Gr05Auto_eAxisClamp1InSawBandPos_Exit(P0);  // exit action
END_STEP
TRANSITION FROM Gr05Auto_eAxisClamp1InSawBandPos TO Gr05Auto_eGetClamp1ActPos_01
    := Trans_16;
END_TRANSITION
STEP Gr05Auto_eGetClamp1ActPos_01:
    Gr05Auto_eGetClamp1ActPos_01_Entry(P1);  // entry action
END_STEP
TRANSITION FROM Gr05Auto_eGetClamp1ActPos_01 TO Dummy_01A
    := TRUE;
END_TRANSITION
TRANSITION FROM Gr05Auto_eAxisClamp1InSawBandPos TO Gr05Auto_eAxisClamp1InSawBandPosErr
    := Trans_17;
END_TRANSITION
STEP Gr05Auto_eAxisClamp1InSawBandPosErr:
    Gr05Auto_eAxisClamp1InSawBandPosErr_Entry(P1);  // entry action
END_STEP
TRANSITION FROM Gr05Auto_eAxisClamp1InSawBandPosErr TO Gr05Auto_eError
    := TRUE;
END_TRANSITION
STEP Dummy_01A:
END_STEP
STEP Gr05Auto_eAxisClamp2MoveToSawBandPos:
    Gr05Auto_eAxisClamp2MoveToSawBandPos_Entry(P1);  // entry action
END_STEP
TRANSITION FROM Gr05Auto_eAxisClamp2MoveToSawBandPos TO Gr05Auto_eAxisClamp2InSawBandPos
    := Trans_18;
END_TRANSITION
TRANSITION FROM Gr05Auto_eAxisClamp2MoveToSawBandPos TO Gr05Auto_eAxisClamp2MoveToSawBandPosErr
    := Trans_19;
END_TRANSITION
STEP Gr05Auto_eAxisClamp2MoveToSawBandPosErr:
    Gr05Auto_eAxisClamp2MoveToSawBandPosErr_Entry(P1);  // entry action
END_STEP
TRANSITION FROM Gr05Auto_eAxisClamp2MoveToSawBandPosErr TO Gr05Auto_eError
    := TRUE;
END_TRANSITION
STEP Gr05Auto_eAxisClamp2InSawBandPos:
    Gr05Auto_eAxisClamp2InSawBandPos_Exit(P0);  // exit action
END_STEP
TRANSITION FROM Gr05Auto_eAxisClamp2InSawBandPos TO Dummy_01B
    := Trans_20;
END_TRANSITION
TRANSITION FROM Gr05Auto_eAxisClamp2InSawBandPos TO Gr05Auto_eAxisClamp2InSawBandPosErr
    := Trans_21;
END_TRANSITION
STEP Gr05Auto_eAxisClamp2InSawBandPosErr:
    Gr05Auto_eAxisClamp2InSawBandPosErr_Entry(P1);  // entry action
END_STEP
TRANSITION FROM Gr05Auto_eAxisClamp2InSawBandPosErr TO Gr05Auto_eError
    := TRUE;
END_TRANSITION
STEP Dummy_01B:
END_STEP
TRANSITION FROM (Dummy_01A, Dummy_01B) TO Gr05Auto_eAxisClamp2MoveSawPos
    := TRUE;
END_TRANSITION
STEP Gr05Auto_eAxisClamp2MoveSawPos:
    Gr05Auto_eAxisClamp2MoveSawPos_Entry(P1);  // entry action
END_STEP
TRANSITION FROM Gr05Auto_eAxisClamp2MoveSawPos TO Gr05Auto_eAxisClamp2InSawPos
    := Trans_22;
END_TRANSITION
TRANSITION FROM Gr05Auto_eAxisClamp2MoveSawPos TO Gr05Auto_eAxisClamp2MoveSawPosErr
    := Trans_23;
END_TRANSITION
STEP Gr05Auto_eAxisClamp2MoveSawPosErr:
    Gr05Auto_eAxisClamp2MoveSawPosErr_Entry(P1);  // entry action
END_STEP
TRANSITION FROM Gr05Auto_eAxisClamp2MoveSawPosErr TO Gr05Auto_eError
    := TRUE;
END_TRANSITION
STEP Gr05Auto_eAxisClamp2InSawPos:
    Gr05Auto_eAxisClamp2InSawPos_Exit(P0);  // exit action
END_STEP
TRANSITION FROM Gr05Auto_eAxisClamp2InSawPos TO Gr05Auto_eGetProcessPara
    := Trans_24;
END_TRANSITION
TRANSITION FROM Gr05Auto_eAxisClamp2InSawPos TO Gr05Auto_eAxisClamp2InSawPosErr
    := Trans_25;
END_TRANSITION
STEP Gr05Auto_eAxisClamp2InSawPosErr:
    Gr05Auto_eAxisClamp2InSawPosErr_Entry(P1);  // entry action
END_STEP
TRANSITION FROM Gr05Auto_eAxisClamp2InSawPosErr TO Gr05Auto_eError
    := TRUE;
END_TRANSITION
STEP Gr05Auto_eGetProcessPara:
    Gr05Auto_eGetProcessPara_Entry(P1);  // entry action
END_STEP
TRANSITION FROM Gr05Auto_eGetProcessPara TO Gr05Auto_eClamp12Open
    := Trans_26;
END_TRANSITION
TRANSITION FROM Gr05Auto_eGetProcessPara TO Gr05Auto_eChkProcessEnd
    := TRUE;
END_TRANSITION
STEP Gr05Auto_eChkProcessEnd:
END_STEP
TRANSITION FROM Gr05Auto_eChkProcessEnd TO Gr05Auto_eWfSlideUp
    := Trans_27;
END_TRANSITION
TRANSITION FROM Gr05Auto_eChkProcessEnd TO Gr05Auto_eClamp12Open
    := TRUE;
END_TRANSITION
STEP Gr05Auto_eWfSlideUp:
END_STEP
TRANSITION FROM Gr05Auto_eWfSlideUp TO Gr05Auto_eGetClamp2ActPos
    := Trans_28;
END_TRANSITION
STEP Gr05Auto_eGetClamp2ActPos:
    Gr05Auto_eGetClamp2ActPos_Entry(P1);  // entry action
END_STEP
TRANSITION FROM Gr05Auto_eGetClamp2ActPos TO Gr05Auto_eChkWorkArea
    := Trans_29;
END_TRANSITION
TRANSITION FROM Gr05Auto_eGetClamp2ActPos TO Gr05Auto_eCollisionDetectedErr
    := TRUE;
END_TRANSITION
STEP Gr05Auto_eCollisionDetectedErr:
    Gr05Auto_eCollisionDetectedErr_Entry(P1);  // entry action
    Gr05Auto_eCollisionDetectedErr_Exit(P0);  // exit action
END_STEP
TRANSITION FROM Gr05Auto_eCollisionDetectedErr TO Gr05Auto_eError
    := Trans_30;
END_TRANSITION
STEP Gr05Auto_eChkWorkArea:
    Gr05Auto_eChkWorkArea_Entry(P1);  // entry action
END_STEP
TRANSITION FROM Gr05Auto_eChkWorkArea TO Gr05Auto_eClamp1Close2
    := _Current_pos_clamp_1_sawing_lenght_current_pos_clamp_2_Current_pos_clamp_2_is_;
END_TRANSITION
STEP Gr05Auto_eClamp1Close2:
    Gr05Auto_eClamp1Close2_Entry(P1);  // entry action
    Gr05Auto_eClamp1Close2_Exit(P0);  // exit action
END_STEP
TRANSITION FROM Gr05Auto_eClamp1Close2 TO Gr05Auto_eChkAxisClamp1MoveToBackPos
    := SafetyDistEnable;
END_TRANSITION
TRANSITION FROM Gr05Auto_eClamp1Close2 TO Gr05Auto_eClamp2Open1
    := Trans_31;
END_TRANSITION
TRANSITION FROM Gr05Auto_eClamp1Close2 TO Gr05Auto_eClamp1Close2Err
    := Trans_32;
END_TRANSITION
STEP Gr05Auto_eClamp1Close2Err:
    Gr05Auto_eClamp1Close2Err_Entry(P1);  // entry action
END_STEP
TRANSITION FROM Gr05Auto_eClamp1Close2Err TO Gr05Auto_eError
    := TRUE;
END_TRANSITION
STEP Gr05Auto_eClamp2Open1:
    Gr05Auto_eClamp2Open1_Entry(P1);  // entry action
    Gr05Auto_eClamp2Open1_Exit(P0);  // exit action
END_STEP
TRANSITION FROM Gr05Auto_eClamp2Open1 TO (Gr05Auto_eAxisClamp1MoveToPos, Gr05Auto_eAxisClamp2MoveToPos)
    := Trans_33;
END_TRANSITION
TRANSITION FROM Gr05Auto_eClamp2Open1 TO Gr05Auto_eClamp2Open1Err
    := Trans_34;
END_TRANSITION
STEP Gr05Auto_eClamp2Open1Err:
    Gr05Auto_eClamp2Open1Err_Entry(P1);  // entry action
END_STEP
TRANSITION FROM Gr05Auto_eClamp2Open1Err TO Gr05Auto_eError
    := TRUE;
END_TRANSITION
STEP Gr05Auto_eAxisClamp1MoveToPos:
    Gr05Auto_eAxisClamp1MoveToPos_Entry(P1);  // entry action
    Gr05Auto_eAxisClamp1MoveToPos_Action(N);  // step action
END_STEP
TRANSITION FROM Gr05Auto_eAxisClamp1MoveToPos TO Gr05Auto_eAxisClamp1InPos
    := Trans_35;
END_TRANSITION
TRANSITION FROM Gr05Auto_eAxisClamp1MoveToPos TO Gr05Auto_eAxisClamp1MoveToPosErr
    := Trans_36;
END_TRANSITION
STEP Gr05Auto_eAxisClamp1MoveToPosErr:
    Gr05Auto_eAxisClamp1MoveToPosErr_Entry(P1);  // entry action
END_STEP
TRANSITION FROM Gr05Auto_eAxisClamp1MoveToPosErr TO Gr05Auto_eError
    := TRUE;
END_TRANSITION
STEP Gr05Auto_eAxisClamp1InPos:
    Gr05Auto_eAxisClamp1InPos_Exit(P0);  // exit action
END_STEP
TRANSITION FROM Gr05Auto_eAxisClamp1InPos TO Gr05Auto_eGetClamp1ActPos_02
    := Trans_37;
END_TRANSITION
STEP Gr05Auto_eGetClamp1ActPos_02:
    Gr05Auto_eGetClamp1ActPos_02_Entry(P1);  // entry action
END_STEP
TRANSITION FROM Gr05Auto_eGetClamp1ActPos_02 TO Dummy_02A
    := TRUE;
END_TRANSITION
TRANSITION FROM Gr05Auto_eAxisClamp1InPos TO Gr05Auto_eAxisClamp1InPosErr
    := Trans_38;
END_TRANSITION
STEP Gr05Auto_eAxisClamp1InPosErr:
    Gr05Auto_eAxisClamp1InPosErr_Entry(P1);  // entry action
END_STEP
TRANSITION FROM Gr05Auto_eAxisClamp1InPosErr TO Gr05Auto_eError
    := TRUE;
END_TRANSITION
STEP Dummy_02A:
END_STEP
STEP Gr05Auto_eAxisClamp2MoveToPos:
    Gr05Auto_eAxisClamp2MoveToPos_Entry(P1);  // entry action
END_STEP
TRANSITION FROM Gr05Auto_eAxisClamp2MoveToPos TO Gr05Auto_eAxisClamp2InPos
    := Trans_39;
END_TRANSITION
TRANSITION FROM Gr05Auto_eAxisClamp2MoveToPos TO Gr05Auto_eAxisClamp2MoveToPosErr
    := Trans_40;
END_TRANSITION
STEP Gr05Auto_eAxisClamp2MoveToPosErr:
    Gr05Auto_eAxisClamp2MoveToPosErr_Entry(P1);  // entry action
END_STEP
TRANSITION FROM Gr05Auto_eAxisClamp2MoveToPosErr TO Gr05Auto_eError
    := TRUE;
END_TRANSITION
STEP Gr05Auto_eAxisClamp2InPos:
    Gr05Auto_eAxisClamp2InPos_Exit(P0);  // exit action
END_STEP
TRANSITION FROM Gr05Auto_eAxisClamp2InPos TO Dummy_02B
    := Trans_41;
END_TRANSITION
TRANSITION FROM Gr05Auto_eAxisClamp2InPos TO Gr05Auto_eAxisClamp2InPosErr
    := Trans_42;
END_TRANSITION
STEP Gr05Auto_eAxisClamp2InPosErr:
    Gr05Auto_eAxisClamp2InPosErr_Entry(P1);  // entry action
END_STEP
TRANSITION FROM Gr05Auto_eAxisClamp2InPosErr TO Gr05Auto_eError
    := TRUE;
END_TRANSITION
STEP Dummy_02B:
END_STEP
TRANSITION FROM (Dummy_02A, Dummy_02B) TO Gr05Auto_eChkAxisClamp1MoveToBackPos
    := TRUE;
END_TRANSITION
STEP Gr05Auto_eChkAxisClamp1MoveToBackPos:
    Gr05Auto_eChkAxisClamp1MoveToBackPos_Entry(P1);  // entry action
    Gr05Auto_eChkAxisClamp1MoveToBackPos_Exit(P0);  // exit action
END_STEP
TRANSITION FROM Gr05Auto_eChkAxisClamp1MoveToBackPos TO Gr05Auto_eAxisClamp1MoveToBackPos
    := ActSawingL_RemoveL;
END_TRANSITION
STEP Gr05Auto_eAxisClamp1MoveToBackPos:
    Gr05Auto_eAxisClamp1MoveToBackPos_Entry(P1);  // entry action
END_STEP
TRANSITION FROM Gr05Auto_eAxisClamp1MoveToBackPos TO Gr05Auto_eAxisClamp1InBackPos
    := Trans_43;
END_TRANSITION
TRANSITION FROM Gr05Auto_eAxisClamp1MoveToBackPos TO Gr05Auto_eAxisClamp1MoveToBackPosErr
    := Trans_44;
END_TRANSITION
STEP Gr05Auto_eAxisClamp1MoveToBackPosErr:
    Gr05Auto_eAxisClamp1MoveToBackPosErr_Entry(P1);  // entry action
END_STEP
TRANSITION FROM Gr05Auto_eAxisClamp1MoveToBackPosErr TO Gr05Auto_eError
    := TRUE;
END_TRANSITION
STEP Gr05Auto_eAxisClamp1InBackPos:
    Gr05Auto_eAxisClamp1InBackPos_Exit(P0);  // exit action
END_STEP
TRANSITION FROM Gr05Auto_eAxisClamp1InBackPos TO Gr05Auto_eGetClamp1ActPos_06
    := Trans_45;
END_TRANSITION
STEP Gr05Auto_eGetClamp1ActPos_06:
    Gr05Auto_eGetClamp1ActPos_06_Entry(P1);  // entry action
END_STEP
TRANSITION FROM Gr05Auto_eGetClamp1ActPos_06 TO Gr05Auto_eChkProcessEnd
    := TRUE;
END_TRANSITION
TRANSITION FROM Gr05Auto_eAxisClamp1InBackPos TO Gr05Auto_eAxisClamp1InBackPosErr
    := Trans_46;
END_TRANSITION
STEP Gr05Auto_eAxisClamp1InBackPosErr:
    Gr05Auto_eAxisClamp1InBackPosErr_Entry(P1);  // entry action
END_STEP
TRANSITION FROM Gr05Auto_eAxisClamp1InBackPosErr TO Gr05Auto_eError
    := TRUE;
END_TRANSITION
TRANSITION FROM Gr05Auto_eChkAxisClamp1MoveToBackPos TO Gr05Auto_ChkPipeEndDetected
    := SafetyDistEnable_1;
END_TRANSITION
TRANSITION FROM Gr05Auto_eChkAxisClamp1MoveToBackPos TO Gr05Auto_eClamp2Slide
    := TRUE;
END_TRANSITION
STEP Gr05Auto_eClamp2Slide:
    Gr05Auto_eClamp2Slide_Entry(P1);  // entry action
    Gr05Auto_eClamp2Slide_Exit(P0);  // exit action
END_STEP
TRANSITION FROM Gr05Auto_eClamp2Slide TO Gr05Auto_eSawingReq
    := Trans_47;
END_TRANSITION
TRANSITION FROM Gr05Auto_eClamp2Slide TO Gr05Auto_eClamp2Err
    := Trans_48;
END_TRANSITION
STEP Gr05Auto_eClamp2Err:
    Gr05Auto_eClamp2Err_Entry(P1);  // entry action
END_STEP
TRANSITION FROM Gr05Auto_eClamp2Err TO Gr05Auto_eError
    := TRUE;
END_TRANSITION
TRANSITION FROM Gr05Auto_eClamp2Slide TO Gr05Auto_eSlideUpErr
    := Trans_49;
END_TRANSITION
STEP Gr05Auto_eSlideUpErr:
    Gr05Auto_eSlideUpErr_Entry(P1);  // entry action
END_STEP
TRANSITION FROM Gr05Auto_eSlideUpErr TO Gr05Auto_eError
    := TRUE;
END_TRANSITION
STEP Gr05Auto_eSawingReq:
    Gr05Auto_eSawingReq_Entry(P1);  // entry action
    Gr05Auto_eSawingReq_Exit(P0);  // exit action
END_STEP
TRANSITION FROM Gr05Auto_eSawingReq TO Gr05Auto_eSawingAck
    := Trans_50;
END_TRANSITION
STEP Gr05Auto_eSawingAck:
END_STEP
TRANSITION FROM Gr05Auto_eSawingAck TO Gr05Auto_eWfTransportReq
    := Trans_51;
END_TRANSITION
STEP Gr05Auto_eWfTransportReq:
    Gr05Auto_eWfTransportReq_Exit(P0);  // exit action
END_STEP
TRANSITION FROM Gr05Auto_eWfTransportReq TO Gr05Auto_eTransportAck
    := Trans_52;
END_TRANSITION
STEP Gr05Auto_eTransportAck:
    Gr05Auto_eTransportAck_Exit(P0);  // exit action
END_STEP
TRANSITION FROM Gr05Auto_eTransportAck TO Gr05Auto_eSlideDown
    := Trans_53;
END_TRANSITION
STEP Gr05Auto_eSlideDown:
    Gr05Auto_eSlideDown_Entry(P1);  // entry action
END_STEP
TRANSITION FROM Gr05Auto_eSlideDown TO Gr05Auto_eGetProcessPara
    := Trans_54;
END_TRANSITION
TRANSITION FROM Gr05Auto_eSlideDown TO Gr05Auto_eSlideDownErr
    := Trans_55;
END_TRANSITION
STEP Gr05Auto_eSlideDownErr:
    Gr05Auto_eSlideDownErr_Entry(P1);  // entry action
END_STEP
TRANSITION FROM Gr05Auto_eSlideDownErr TO Gr05Auto_eError
    := TRUE;
END_TRANSITION
TRANSITION FROM Gr05Auto_eSlideDown TO Gr05Auto_eRemovalBandErr
    := Trans_56;
END_TRANSITION
STEP Gr05Auto_eRemovalBandErr:
    Gr05Auto_eRemovalBandErr_Entry(P1);  // entry action
END_STEP
TRANSITION FROM Gr05Auto_eRemovalBandErr TO Gr05Auto_eError
    := TRUE;
END_TRANSITION
TRANSITION FROM Gr05Auto_eChkWorkArea TO Gr05Auto_ChkPipeEndDetected
    := TRUE;
END_TRANSITION
STEP Gr05Auto_ChkPipeEndDetected:
END_STEP
TRANSITION FROM Gr05Auto_ChkPipeEndDetected TO Gr05Auto_eClamp2Close
    := _No_pipe_end_detected_;
END_TRANSITION
TRANSITION FROM Gr05Auto_ChkPipeEndDetected TO Gr05Auto_eClamp12Open
    := TRUE;
END_TRANSITION
STEP Gr05Auto_eClamp2Close:
    Gr05Auto_eClamp2Close_Entry(P1);  // entry action
    Gr05Auto_eClamp2Close_Exit(P0);  // exit action
END_STEP
TRANSITION FROM Gr05Auto_eClamp2Close TO Gr05Auto_eClamp1Open
    := Trans_57;
END_TRANSITION
TRANSITION FROM Gr05Auto_eClamp2Close TO Gr05Auto_eClamp2CloseErr
    := Trans_58;
END_TRANSITION
STEP Gr05Auto_eClamp2CloseErr:
    Gr05Auto_eClamp2CloseErr_Entry(P1);  // entry action
END_STEP
TRANSITION FROM Gr05Auto_eClamp2CloseErr TO Gr05Auto_eError
    := TRUE;
END_TRANSITION
STEP Gr05Auto_eClamp1Open:
    Gr05Auto_eClamp1Open_Entry(P1);  // entry action
    Gr05Auto_eClamp1Open_Exit(P0);  // exit action
END_STEP
TRANSITION FROM Gr05Auto_eClamp1Open TO Gr05Auto_eAxisClamp1MoveAbsPipeEnde
    := Trans_59;
END_TRANSITION
TRANSITION FROM Gr05Auto_eClamp1Open TO Gr05Auto_eClamp1OpenErr
    := Trans_60;
END_TRANSITION
STEP Gr05Auto_eClamp1OpenErr:
    Gr05Auto_eClamp1OpenErr_Entry(P1);  // entry action
END_STEP
TRANSITION FROM Gr05Auto_eClamp1OpenErr TO Gr05Auto_eError
    := TRUE;
END_TRANSITION
STEP Gr05Auto_eAxisClamp1MoveAbsPipeEnde:
    Gr05Auto_eAxisClamp1MoveAbsPipeEnde_Entry(P1);  // entry action
    Gr05Auto_eAxisClamp1MoveAbsPipeEnde_Exit(P0);  // exit action
END_STEP
TRANSITION FROM Gr05Auto_eAxisClamp1MoveAbsPipeEnde TO Gr05Auto_eWfAxisClamp1MoveAbsPipeEnde
    := Trans_61;
END_TRANSITION
TRANSITION FROM Gr05Auto_eAxisClamp1MoveAbsPipeEnde TO Gr05Auto_eAxisClamp1MoveAbsPipeEndeErr
    := Trans_62;
END_TRANSITION
STEP Gr05Auto_eAxisClamp1MoveAbsPipeEndeErr:
    Gr05Auto_eAxisClamp1MoveAbsPipeEndeErr_Entry(P1);  // entry action
END_STEP
TRANSITION FROM Gr05Auto_eAxisClamp1MoveAbsPipeEndeErr TO Gr05Auto_eError
    := TRUE;
END_TRANSITION
STEP Gr05Auto_eWfAxisClamp1MoveAbsPipeEnde:
    Gr05Auto_eWfAxisClamp1MoveAbsPipeEnde_Exit(P0);  // exit action
END_STEP
TRANSITION FROM Gr05Auto_eWfAxisClamp1MoveAbsPipeEnde TO Gr05Auto_eAxisClamp1Stop
    := _Pipe_end_detected_;
END_TRANSITION
STEP Gr05Auto_eAxisClamp1Stop:
    Gr05Auto_eAxisClamp1Stop_Entry(P1);  // entry action
END_STEP
TRANSITION FROM Gr05Auto_eAxisClamp1Stop TO Gr05Auto_eWfAxisClamp1Stop
    := Trans_63;
END_TRANSITION
TRANSITION FROM Gr05Auto_eAxisClamp1Stop TO Gr05Auto_eAxisClamp1StopErr
    := Trans_64;
END_TRANSITION
STEP Gr05Auto_eAxisClamp1StopErr:
    Gr05Auto_eAxisClamp1StopErr_Entry(P1);  // entry action
END_STEP
TRANSITION FROM Gr05Auto_eAxisClamp1StopErr TO Gr05Auto_eError
    := TRUE;
END_TRANSITION
STEP Gr05Auto_eWfAxisClamp1Stop:
    Gr05Auto_eWfAxisClamp1Stop_Exit(P0);  // exit action
END_STEP
TRANSITION FROM Gr05Auto_eWfAxisClamp1Stop TO Gr05Auto_eGetClamp1ActPos_04
    := Trans_65;
END_TRANSITION
STEP Gr05Auto_eGetClamp1ActPos_04:
    Gr05Auto_eGetClamp1ActPos_04_Entry(P1);  // entry action
END_STEP
TRANSITION FROM Gr05Auto_eGetClamp1ActPos_04 TO Gr05Auto_eChkNextSawingAngle
    := TRUE;
END_TRANSITION
TRANSITION FROM Gr05Auto_eWfAxisClamp1Stop TO Gr05Auto_eWfAxisClamp1StopErr
    := Trans_66;
END_TRANSITION
STEP Gr05Auto_eWfAxisClamp1StopErr:
    Gr05Auto_eWfAxisClamp1StopErr_Entry(P1);  // entry action
END_STEP
TRANSITION FROM Gr05Auto_eWfAxisClamp1StopErr TO Gr05Auto_eError
    := TRUE;
END_TRANSITION
STEP Gr05Auto_eChkNextSawingAngle:
END_STEP
TRANSITION FROM Gr05Auto_eChkNextSawingAngle TO Gr05Auto_eAxisClamp1MoveVeloPipeEnd
    := Trans_67;
END_TRANSITION
STEP Gr05Auto_eAxisClamp1MoveVeloPipeEnd:
    Gr05Auto_eAxisClamp1MoveVeloPipeEnd_Entry(P1);  // entry action
END_STEP
TRANSITION FROM Gr05Auto_eAxisClamp1MoveVeloPipeEnd TO Gr05Auto_eWfAxisClamp1MoveVeloPipeEnd
    := Trans_68;
END_TRANSITION
TRANSITION FROM Gr05Auto_eAxisClamp1MoveVeloPipeEnd TO Gr05Auto_eAxisClamp1MoveVeloPipeEndErr
    := Trans_69;
END_TRANSITION
STEP Gr05Auto_eAxisClamp1MoveVeloPipeEndErr:
    Gr05Auto_eAxisClamp1MoveVeloPipeEndErr_Entry(P1);  // entry action
END_STEP
TRANSITION FROM Gr05Auto_eAxisClamp1MoveVeloPipeEndErr TO Gr05Auto_eError
    := TRUE;
END_TRANSITION
STEP Gr05Auto_eWfAxisClamp1MoveVeloPipeEnd:
    Gr05Auto_eWfAxisClamp1MoveVeloPipeEnd_Exit(P0);  // exit action
END_STEP
TRANSITION FROM Gr05Auto_eWfAxisClamp1MoveVeloPipeEnd TO Gr05Auto_eAxisClamp1InPipeEndPos
    := Trans_70;
END_TRANSITION
TRANSITION FROM Gr05Auto_eWfAxisClamp1MoveVeloPipeEnd TO Gr05Auto_eWfAxisClamp1MoveVeloPipeEndErr
    := Trans_71;
END_TRANSITION
STEP Gr05Auto_eWfAxisClamp1MoveVeloPipeEndErr:
    Gr05Auto_eWfAxisClamp1MoveVeloPipeEndErr_Entry(P1);  // entry action
END_STEP
TRANSITION FROM Gr05Auto_eWfAxisClamp1MoveVeloPipeEndErr TO Gr05Auto_eError
    := TRUE;
END_TRANSITION
STEP Gr05Auto_eAxisClamp1InPipeEndPos:
    Gr05Auto_eAxisClamp1InPipeEndPos_Action(N);  // step action
    Gr05Auto_eAxisClamp1InPipeEndPos_Exit(P0);  // exit action
END_STEP
TRANSITION FROM Gr05Auto_eAxisClamp1InPipeEndPos TO Gr05Auto_eAxisClamp1Stop_2
    := _Pipe_end_was_detected_;
END_TRANSITION
TRANSITION FROM Gr05Auto_eAxisClamp1InPipeEndPos TO Gr05Auto_eWfPipeEndNoDetectedErr
    := _Pipe_end_was_not_detected_;
END_TRANSITION
STEP Gr05Auto_eWfPipeEndNoDetectedErr:
    Gr05Auto_eWfPipeEndNoDetectedErr_Entry(P1);  // entry action
    Gr05Auto_eWfPipeEndNoDetectedErr_Exit(P0);  // exit action
END_STEP
TRANSITION FROM Gr05Auto_eWfPipeEndNoDetectedErr TO Gr05Auto_eError
    := Trans_72;
END_TRANSITION
STEP Gr05Auto_eAxisClamp1Stop_2:
    Gr05Auto_eAxisClamp1Stop_2_Entry(P1);  // entry action
END_STEP
TRANSITION FROM Gr05Auto_eAxisClamp1Stop_2 TO Gr05Auto_eWfAxisClamp1Stop_2
    := Trans_73;
END_TRANSITION
TRANSITION FROM Gr05Auto_eAxisClamp1Stop_2 TO Gr05Auto_eAxisClamp1StopErr_2
    := Trans_74;
END_TRANSITION
STEP Gr05Auto_eAxisClamp1StopErr_2:
    Gr05Auto_eAxisClamp1StopErr_2_Entry(P1);  // entry action
END_STEP
TRANSITION FROM Gr05Auto_eAxisClamp1StopErr_2 TO Gr05Auto_eError
    := TRUE;
END_TRANSITION
STEP Gr05Auto_eWfAxisClamp1Stop_2:
    Gr05Auto_eWfAxisClamp1Stop_2_Exit(P0);  // exit action
END_STEP
TRANSITION FROM Gr05Auto_eWfAxisClamp1Stop_2 TO _Gr05Auto_ChkNextSawingLenght
    := Trans_75;
END_TRANSITION
TRANSITION FROM Gr05Auto_eWfAxisClamp1Stop_2 TO Gr05Auto_eWfAxisClamp1StopErr_2
    := Trans_76;
END_TRANSITION
STEP Gr05Auto_eWfAxisClamp1StopErr_2:
    Gr05Auto_eWfAxisClamp1StopErr_2_Entry(P1);  // entry action
END_STEP
TRANSITION FROM Gr05Auto_eWfAxisClamp1StopErr_2 TO Gr05Auto_eError
    := TRUE;
END_TRANSITION
STEP _Gr05Auto_ChkNextSawingLenght:  // name as stored:  Gr05Auto_ChkNextSawingLenght
END_STEP
TRANSITION FROM _Gr05Auto_ChkNextSawingLenght TO Gr05Auto_eGetClamp1ActPos_05
    := Trans_77;
END_TRANSITION
STEP Gr05Auto_eGetClamp1ActPos_05:
    Gr05Auto_eGetClamp1ActPos_05_Entry(P1);  // entry action
END_STEP
TRANSITION FROM Gr05Auto_eGetClamp1ActPos_05 TO Dummy_03
    := Trans_78;
END_TRANSITION
TRANSITION FROM Gr05Auto_eGetClamp1ActPos_05 TO Gr05Auto_eAngleReq
    := TRUE;
END_TRANSITION
STEP Gr05Auto_eAngleReq:
    Gr05Auto_eAngleReq_Entry(P1);  // entry action
    Gr05Auto_eAngleReq_Exit(P0);  // exit action
END_STEP
TRANSITION FROM Gr05Auto_eAngleReq TO Gr05Auto_eAngleAck
    := Trans_79;
END_TRANSITION
STEP Gr05Auto_eAngleAck:
END_STEP
TRANSITION FROM Gr05Auto_eAngleAck TO Dummy_03
    := Trans_80;
END_TRANSITION
TRANSITION FROM _Gr05Auto_ChkNextSawingLenght TO Dummy_03
    := TRUE;
END_TRANSITION
TRANSITION FROM Gr05Auto_eChkNextSawingAngle TO Dummy_03
    := TRUE;
END_TRANSITION
STEP Dummy_03:
END_STEP
TRANSITION FROM Dummy_03 TO Gr05Auto_eChkProcessEnd
    := TRUE;
END_TRANSITION
TRANSITION FROM Gr05Auto_eWfAxisClamp1MoveAbsPipeEnde TO Gr05Auto_eGetClamp1ActPos_03
    := Trans_81;
END_TRANSITION
STEP Gr05Auto_eGetClamp1ActPos_03:
    Gr05Auto_eGetClamp1ActPos_03_Entry(P1);  // entry action
END_STEP
TRANSITION FROM Gr05Auto_eGetClamp1ActPos_03 TO Gr05Auto_eClamp1Close3
    := Trans_82;
END_TRANSITION
STEP Gr05Auto_eClamp1Close3:
    Gr05Auto_eClamp1Close3_Entry(P1);  // entry action
    Gr05Auto_eClamp1Close3_Exit(P0);  // exit action
END_STEP
TRANSITION FROM Gr05Auto_eClamp1Close3 TO Gr05Auto_eChkAdjustSawingLength
    := Trans_83;
END_TRANSITION
TRANSITION FROM Gr05Auto_eClamp1Close3 TO Gr05Auto_eClamp1Close3Err
    := Trans_84;
END_TRANSITION
STEP Gr05Auto_eClamp1Close3Err:
    Gr05Auto_eClamp1Close3Err_Entry(P1);  // entry action
END_STEP
TRANSITION FROM Gr05Auto_eClamp1Close3Err TO Gr05Auto_eError
    := TRUE;
END_TRANSITION
STEP Gr05Auto_eChkAdjustSawingLength:
END_STEP
TRANSITION FROM Gr05Auto_eChkAdjustSawingLength TO Gr05Auto_NurWennlrActRemoveLength_0
    := _Current_pos_clamp_1_sawing_lenght_current_pos_clamp_2_Current_pos_clamp_2_is_1;
END_TRANSITION
TRANSITION FROM Gr05Auto_eChkAdjustSawingLength TO Gr05Auto_eChkProcessEnd
    := TRUE;
END_TRANSITION
STEP Gr05Auto_NurWennlrActRemoveLength_0:
END_STEP
TRANSITION FROM Gr05Auto_NurWennlrActRemoveLength_0 TO Gr05Auto_eClamp2Open3
    := Trans_85;
END_TRANSITION
STEP Gr05Auto_eClamp2Open3:
    Gr05Auto_eClamp2Open3_Entry(P1);  // entry action
    Gr05Auto_eClamp2Open3_Exit(P0);  // exit action
END_STEP
TRANSITION FROM Gr05Auto_eClamp2Open3 TO Gr05Auto_eAxisClamp2MoveToPos2
    := Trans_86;
END_TRANSITION
TRANSITION FROM Gr05Auto_eClamp2Open3 TO Gr05Auto_eClamp2Open3Err
    := Trans_87;
END_TRANSITION
STEP Gr05Auto_eClamp2Open3Err:
    Gr05Auto_eClamp2Open3Err_Entry(P1);  // entry action
END_STEP
TRANSITION FROM Gr05Auto_eClamp2Open3Err TO Gr05Auto_eError
    := TRUE;
END_TRANSITION
STEP Gr05Auto_eAxisClamp2MoveToPos2:
    Gr05Auto_eAxisClamp2MoveToPos2_Entry(P1);  // entry action
END_STEP
TRANSITION FROM Gr05Auto_eAxisClamp2MoveToPos2 TO Gr05Auto_eAxisClamp2InPos2
    := Trans_88;
END_TRANSITION
TRANSITION FROM Gr05Auto_eAxisClamp2MoveToPos2 TO Gr05Auto_eAxisClamp2MoveToPos2Err
    := Trans_89;
END_TRANSITION
STEP Gr05Auto_eAxisClamp2MoveToPos2Err:
    Gr05Auto_eAxisClamp2MoveToPos2Err_Entry(P1);  // entry action
END_STEP
TRANSITION FROM Gr05Auto_eAxisClamp2MoveToPos2Err TO Gr05Auto_eError
    := TRUE;
END_TRANSITION
STEP Gr05Auto_eAxisClamp2InPos2:
    Gr05Auto_eAxisClamp2InPos2_Exit(P0);  // exit action
END_STEP
TRANSITION FROM Gr05Auto_eAxisClamp2InPos2 TO Gr05Auto_eAxisClamp1MoveToPos2
    := Trans_90;
END_TRANSITION
TRANSITION FROM Gr05Auto_eAxisClamp2InPos2 TO Gr05Auto_eAxisClamp2InPos2Err
    := Trans_91;
END_TRANSITION
STEP Gr05Auto_eAxisClamp2InPos2Err:
    Gr05Auto_eAxisClamp2InPos2Err_Entry(P1);  // entry action
END_STEP
TRANSITION FROM Gr05Auto_eAxisClamp2InPos2Err TO Gr05Auto_eError
    := TRUE;
END_TRANSITION
STEP Gr05Auto_eAxisClamp1MoveToPos2:
    Gr05Auto_eAxisClamp1MoveToPos2_Entry(P1);  // entry action
END_STEP
TRANSITION FROM Gr05Auto_eAxisClamp1MoveToPos2 TO Gr05Auto_eAxisClamp1InPos2
    := Trans_92;
END_TRANSITION
TRANSITION FROM Gr05Auto_eAxisClamp1MoveToPos2 TO Gr05Auto_eAxisClamp1MoveToPos2Err
    := Trans_93;
END_TRANSITION
STEP Gr05Auto_eAxisClamp1MoveToPos2Err:
    Gr05Auto_eAxisClamp1MoveToPos2Err_Entry(P1);  // entry action
END_STEP
TRANSITION FROM Gr05Auto_eAxisClamp1MoveToPos2Err TO Gr05Auto_eError
    := TRUE;
END_TRANSITION
STEP Gr05Auto_eAxisClamp1InPos2:
    Gr05Auto_eAxisClamp1InPos2_Exit(P0);  // exit action
END_STEP
TRANSITION FROM Gr05Auto_eAxisClamp1InPos2 TO Gr05Auto_eSawingLengthCorrection
    := Trans_94;
END_TRANSITION
STEP Gr05Auto_eSawingLengthCorrection:
    Gr05Auto_eSawingLengthCorrection_Entry(P1);  // entry action
END_STEP
TRANSITION FROM Gr05Auto_eSawingLengthCorrection TO Gr05Auto_ChkPipeEndDetected
    := TRUE;
END_TRANSITION
TRANSITION FROM Gr05Auto_eAxisClamp1InPos2 TO Gr05Auto_eAxisClamp1InPos2Err
    := Trans_95;
END_TRANSITION
STEP Gr05Auto_eAxisClamp1InPos2Err:
    Gr05Auto_eAxisClamp1InPos2Err_Entry(P1);  // entry action
END_STEP
TRANSITION FROM Gr05Auto_eAxisClamp1InPos2Err TO Gr05Auto_eError
    := TRUE;
END_TRANSITION
TRANSITION FROM Gr05Auto_eWfAxisClamp1MoveAbsPipeEnde TO Gr05Auto_eWfAxisClamp1MoveAbsPipeEndeErr
    := Trans_96;
END_TRANSITION
STEP Gr05Auto_eWfAxisClamp1MoveAbsPipeEndeErr:
    Gr05Auto_eWfAxisClamp1MoveAbsPipeEndeErr_Entry(P1);  // entry action
END_STEP
TRANSITION FROM Gr05Auto_eWfAxisClamp1MoveAbsPipeEndeErr TO Gr05Auto_eError
    := TRUE;
END_TRANSITION
STEP Gr05Auto_eClamp12Open:
    Gr05Auto_eClamp12Open_Entry(P1);  // entry action
    Gr05Auto_eClamp12Open_Exit(P0);  // exit action
END_STEP
TRANSITION FROM Gr05Auto_eClamp12Open TO Gr05Auto_eEnd
    := Trans_97;
END_TRANSITION
TRANSITION FROM Gr05Auto_eClamp12Open TO Gr05Auto_eClamp1Open2Err
    := Trans_98;
END_TRANSITION
STEP Gr05Auto_eClamp1Open2Err:
    Gr05Auto_eClamp1Open2Err_Entry(P1);  // entry action
END_STEP
TRANSITION FROM Gr05Auto_eClamp1Open2Err TO Gr05Auto_eError
    := TRUE;
END_TRANSITION
TRANSITION FROM Gr05Auto_eClamp12Open TO Gr05Auto_eClamp2Open2Err
    := Trans_99;
END_TRANSITION
STEP Gr05Auto_eClamp2Open2Err:
    Gr05Auto_eClamp2Open2Err_Entry(P1);  // entry action
END_STEP
TRANSITION FROM Gr05Auto_eClamp2Open2Err TO Gr05Auto_eError
    := TRUE;
END_TRANSITION
STEP Gr05Auto_eEnd:
END_STEP
TRANSITION FROM Gr05Auto_eEnd TO Gr05Auto_eDone
    := TRUE;
END_TRANSITION
STEP Gr05Auto_eDone:
    Gr05Auto_eDone_Entry(P1);  // entry action
    Gr05Auto_eDone_Exit(P0);  // exit action
END_STEP
TRANSITION FROM Gr05Auto_eDone TO Gr05Auto_eNoExecute
    := Trans_100;
END_TRANSITION
TRANSITION FROM Gr05Auto_eEnd TO Gr05Auto_eError
    := FALSE;
END_TRANSITION
STEP Gr05Auto_eError:
    Gr05Auto_eError_Entry(P1);  // entry action
    Gr05Auto_eError_Exit(P0);  // exit action
END_STEP
TRANSITION FROM Gr05Auto_eError TO Gr05Auto_eNoExecute
    := Trans_101;
END_TRANSITION
STEP Gr05Auto_eNoExecute:
END_STEP
TRANSITION FROM Gr05Auto_eNoExecute TO Init
    := TRUE;
END_TRANSITION

TRANSITION _Current_pos_clamp_1_sawing_lenght_current_pos_clamp_2_Current_pos_clamp_2_is_:
(*1 Current pos clamp 1 - sawing lenght > current pos clamp 2 (Current pos clamp 2 is " + ") *)
(lrClamp1Pos - MAX(ABS(lrActSawingLength), ABS(lrActRemoveLength)) > (F_GetCylinderPos(
										F_SetCylinderPos(SEL(stgGr05HMI.stHMITOPLC.bCylinderPosActive, Gr05Control.fbCylinderPos.lrActPosition, lrClamp2Pos),
														lrgGr05CylinderPosOffset,
														lrgGr05CylinderPosOriginShiftPos,
														etgGr05CylinderPosDirection,
														usngGr05CylinderPosCodingType),
										lrgGr05CylinderPosOffset,
										lrgGr05CylinderPosOriginShiftPos,
										etgGr05CylinderPosDirection,
										usngGr05CylinderPosCodingType)
									    	+ lrgGr05Clamp2Width (*+ lrgGr05SafetyDistance*)))
AND bReleaseNextStep
END_TRANSITION

TRANSITION _Current_pos_clamp_1_sawing_lenght_current_pos_clamp_2_Current_pos_clamp_2_is_1:
(*2 Current pos clamp 1 - sawing lenght <= current pos clamp 2 (Current pos clamp 2 is " + ") *)
(lrClamp1Pos - MAX(ABS(lrActSawingLength), ABS(lrActRemoveLength)) <= (F_GetCylinderPos(
														F_SetCylinderPos(SEL(stgGr05HMI.stHMITOPLC.bCylinderPosActive, Gr05Control.fbCylinderPos.lrActPosition, lrClamp2Pos),
																		lrgGr05CylinderPosOffset,
																		lrgGr05CylinderPosOriginShiftPos,
																		etgGr05CylinderPosDirection,
																		usngGr05CylinderPosCodingType),
														lrgGr05CylinderPosOffset,
														lrgGr05CylinderPosOriginShiftPos,
														etgGr05CylinderPosDirection,
														usngGr05CylinderPosCodingType)
									   					 + lrgGr05Clamp2Width))
AND bReleaseNextStep
END_TRANSITION

TRANSITION _No_pipe_end_detected_:
NOT bPipeEndDetected
AND bReleaseNextStep
END_TRANSITION

TRANSITION _Pipe_begin_was_detected_:
(* Pipe begin was detected *)
rtPipeBeginIdentify.Q
END_TRANSITION

TRANSITION _Pipe_begin_was_no_detected_:
Gr05Control.fbAxisClamp1.lrActPosition < (lrgGr05Clamp1DistPipeBeginSawBand + 10)
OR Gr05Control.fbAxisClamp1.bHardLimitMinExceeded
OR Gr05Control.fbAxisClamp1.bSoftLimitMinExceeded
END_TRANSITION

TRANSITION _Pipe_begin_was_no_detected_1:
(Gr05Control.fbAxisClamp1.lrActPosition <= lrClamp1Pos - lrgGr05SearchDistPipeBegin
AND Gr05Control.fbAxisClamp1.lrActPosition > (lrgGr05Clamp1DistPipeBeginSawBand + 10))
OR Gr05Control.fbAxisClamp1.bHardLimitMinExceeded
OR Gr05Control.fbAxisClamp1.bSoftLimitMinExceeded
END_TRANSITION

TRANSITION _Pipe_end_detected_:
NOT binGr05PipeEndEdge
AND bReleaseNextStep
END_TRANSITION

TRANSITION _Pipe_end_was_detected_:
(* Pipe end was detected *)
rtPipeEndIdentify.Q
END_TRANSITION

TRANSITION _Pipe_end_was_not_detected_:
Gr05Control.fbAxisClamp1.lrActPosition <= lrClamp1Pos - lrgGr05SearchDistPipeEnd
OR Gr05Control.fbAxisClamp1.bHardLimitMinExceeded
OR Gr05Control.fbAxisClamp1.bSoftLimitMinExceeded
END_TRANSITION

TRANSITION ActSawingL_RemoveL:
ABS(lrActSawingLength) < ABS(lrActRemoveLength)
END_TRANSITION

ACTION Gr05Auto_ChkPipeBeginEdge_Exit:
IF NOT binGr05PipeBeginEdge
THEN
	lrDistPipeBeginSawBand := lrgGr05Clamp1DistPipeBeginSawBand;
ELSE
	lrDistPipeBeginSawBand := 0;
END_IF
END_ACTION

ACTION Gr05Auto_eAngleReq_Entry:
stgGr05HMI.stHMITOPLC.lrActSawingLength := ABS(lrClamp1PosPipeEnd - ABS(stgGr05HMI.stHMITOPLC.lrActSawingLength));
lrActSawingLength := ABS(lrClamp1PosPipeEnd - ABS(lrActSawingLength));									(* Next sawing lenght *)
lrActSawingAngle := arrGr00ProcessPara[unProcessCounter - 1, 1] / 180 * PI;
bgGr05AngleReq := TRUE;
END_ACTION

ACTION Gr05Auto_eAngleReq_Exit:
bgGr05AngleReq := FALSE;
END_ACTION

ACTION Gr05Auto_eAxisClamp1InBackPos_Exit:
Gr05Control.fbAxisClamp1.bExeMoveAbs := FALSE;
END_ACTION

ACTION Gr05Auto_eAxisClamp1InBackPosErr_Entry:
Gr05Control.fbAxisClamp1.bExeMoveAbs := FALSE;
END_ACTION

ACTION Gr05Auto_eAxisClamp1InPipeBeginPos_Action:
rtPipeBeginIdentify(CLK := binGr05PipeBeginEdge);
END_ACTION

ACTION Gr05Auto_eAxisClamp1InPipeBeginPos_Exit:
rtPipeBeginIdentify(CLK := FALSE);
END_ACTION

ACTION Gr05Auto_eAxisClamp1InPipeEndPos_Action:
rtPipeEndIdentify(CLK := binGr05PipeEndEdge );
END_ACTION

ACTION Gr05Auto_eAxisClamp1InPipeEndPos_Exit:
rtPipeEndIdentify(CLK := FALSE);
END_ACTION

ACTION Gr05Auto_eAxisClamp1InPos_Exit:
Gr05Control.fbAxisClamp1.bExeMoveAbs := FALSE;
END_ACTION

ACTION Gr05Auto_eAxisClamp1InPos2_Exit:
Gr05Control.fbAxisClamp1.bExeMoveAbs := FALSE;
END_ACTION

ACTION Gr05Auto_eAxisClamp1InPos2Err_Entry:
Gr05Control.fbAxisClamp1.bExeMoveAbs := FALSE;
END_ACTION

ACTION Gr05Auto_eAxisClamp1InPosErr_Entry:
Gr05Control.fbAxisClamp1.bExeMoveAbs := FALSE;
END_ACTION

ACTION Gr05Auto_eAxisClamp1InSawBandPos_Exit:
Gr05Control.fbAxisClamp1.bExeMoveAbs := FALSE;
END_ACTION

ACTION Gr05Auto_eAxisClamp1InSawBandPosErr_Entry:
Gr05Control.fbAxisClamp1.bExeMoveAbs := FALSE;
END_ACTION

ACTION Gr05Auto_eAxisClamp1MoveAbsPipeEnde_Entry:
Gr05Control.fbAxisClamp1.bExeMoveAbs := binGr05PipeEndEdge;
Gr05Control.fbAxisClamp1.lrTargetPosition := stgGr05HMI.stHMITOPLC.arlrAxisClampSoftLimitMax[1];
Gr05Control.fbAxisClamp1.lrAutoVelocity := stgGr05HMI.stHMITOPLC.arlrAxisClampAutoVelo[1];
END_ACTION

ACTION Gr05Auto_eAxisClamp1MoveAbsPipeEnde_Exit:
IF NOT Gr05Control.fbUtility.bPipeEndPresent
THEN
	Gr05Control.fbAxisClamp1.bExeMoveAbs := FALSE;
END_IF
END_ACTION

ACTION Gr05Auto_eAxisClamp1MoveAbsPipeEndeErr_Entry:
Gr05Control.fbAxisClamp1.bExeMoveAbs := FALSE;
END_ACTION

ACTION Gr05Auto_eAxisClamp1MoveToBackPos_Entry:
Gr05Control.fbAxisClamp1.bExeMoveAbs := TRUE;
Gr05Control.fbAxisClamp1.lrTargetPosition := lrClamp1Pos + ABS(lrActRemoveLength - lrActSawingLength);
Gr05Control.fbAxisClamp1.lrAutoVelocity := stgGr05HMI.stHMITOPLC.arlrAxisClampAutoVelo[1];
lrActSawingLength := 0.0;
END_ACTION

ACTION Gr05Auto_eAxisClamp1MoveToBackPosErr_Entry:
Gr05Control.fbAxisClamp1.bExeMoveAbs := FALSE;
END_ACTION

ACTION Gr05Auto_eAxisClamp1MoveToPos_Action:

Gr05Control.fbAxisClamp1.bExeMoveAbs := lrClamp1Pos - MAX(ABS(lrActSawingLength), ABS(lrActRemoveLength)) > (stgGr05HMI.stPLCTOHMI.arlrAxisClampActPos[2] + lrgGr05Clamp2Width (*+lrgGr05SafetyDistance   	(*ESKG 12032026*)*) );
END_ACTION

ACTION Gr05Auto_eAxisClamp1MoveToPos_Entry:
(*IF lrClamp1Pos + ABS(lrActSawingLength) > stgGr05HMI.stPLCTOHMI.lrAxisClamp1ActPos
THEN
	Gr05Control.fbAxisClamp1.bExeMoveAbs := lrClamp1Pos + ABS(lrActSawingLength) < (stgGr05HMI.stPLCTOHMI.lrAxisClamp2ActPos - lrgGr05Clamp2Width);
ELSE
	Gr05Control.fbAxisClamp1.bExeMoveAbs := TRUE;
END_IF*)
Gr05Control.fbAxisClamp1.lrTargetPosition := lrClamp1Pos - MAX(ABS(lrActSawingLength), ABS(lrActRemoveLength));
Gr05Control.fbAxisClamp1.lrAutoVelocity := stgGr05HMI.stHMITOPLC.arlrAxisClampAutoVelo[1];
END_ACTION

ACTION Gr05Auto_eAxisClamp1MoveToPos2_Entry:
Gr05Control.fbAxisClamp1.bExeMoveAbs := TRUE;
Gr05Control.fbAxisClamp1.lrTargetPosition := lrClamp1Pos -MIN(lrActSawingLength , ABS(Gr05Control.fbAxisClamp1.lrActPosition - Gr05Control.fbCylinderPos.lrActPosition - lrgGr05Clamp2Width)); 	(*ESKG 12032026*)
Gr05Control.fbAxisClamp1.lrAutoVelocity := stgGr05HMI.stHMITOPLC.arlrAxisClampAutoVelo[1];
END_ACTION

ACTION Gr05Auto_eAxisClamp1MoveToPos2Err_Entry:
Gr05Control.fbAxisClamp1.bExeMoveAbs := FALSE;
END_ACTION

ACTION Gr05Auto_eAxisClamp1MoveToPosErr_Entry:
Gr05Control.fbAxisClamp1.bExeMoveAbs := FALSE;
END_ACTION

ACTION Gr05Auto_eAxisClamp1MoveToSawBandPos_Entry:
Gr05Control.fbAxisClamp1.bExeMoveAbs := TRUE;
Gr05Control.fbAxisClamp1.lrTargetPosition := lrClamp1Pos - lrDistPipeBeginSawBand;
Gr05Control.fbAxisClamp1.lrAutoVelocity := stgGr05HMI.stHMITOPLC.arlrAxisClampAutoVelo[1];
END_ACTION

ACTION Gr05Auto_eAxisClamp1MoveToSawBandPosErr_Entry:
Gr05Control.fbAxisClamp1.bExeMoveAbs := FALSE;
END_ACTION

ACTION Gr05Auto_eAxisClamp1MoveVeloPipeBegin_Entry:
Gr05Control.fbAxisClamp1.bExeMoveVelo := TRUE;
Gr05Control.fbAxisClamp1.lrAutoVelocity := -stgGr05HMI.stHMITOPLC.arlrAxisClampAutoVelo[1] / 10;
lrClamp1Pos := Gr05Control.fbAxisClamp1.lrActPosition;
END_ACTION

ACTION Gr05Auto_eAxisClamp1MoveVeloPipeBeginErr_Entry:
Gr05Control.fbAxisClamp1.bExeMoveVelo := FALSE;
END_ACTION

ACTION Gr05Auto_eAxisClamp1MoveVeloPipeEnd_Entry:
Gr05Control.fbAxisClamp1.bExeMoveVelo := TRUE;
Gr05Control.fbAxisClamp1.lrAutoVelocity := -stgGr05HMI.stHMITOPLC.arlrAxisClampAutoVelo[1] / 10;
END_ACTION

ACTION Gr05Auto_eAxisClamp1MoveVeloPipeEndErr_Entry:
Gr05Control.fbAxisClamp1.bExeMoveVelo := FALSE;
END_ACTION

ACTION Gr05Auto_eAxisClamp1Stop_2_Entry:
Gr05Control.fbAxisClamp1.bExeStop := TRUE;
Gr05Control.fbAxisClamp1.lrAutoVelocity := 0.0;
lrClamp1PosPipeEnd := Gr05Control.fbAxisClamp1.lrActPosition + lrgGr05Clamp1PipeSensorOffset;
END_ACTION

ACTION Gr05Auto_eAxisClamp1Stop_Entry:
Gr05Control.fbAxisClamp1.bExeStop := TRUE;
Gr05Control.fbAxisClamp1.lrAutoVelocity := 0.0;
bPipeEndDetected := TRUE;
END_ACTION

ACTION Gr05Auto_eAxisClamp1StopErr_2_Entry:
Gr05Control.fbAxisClamp1.bExeStop := FALSE;
END_ACTION

ACTION Gr05Auto_eAxisClamp1StopErr_Entry:
Gr05Control.fbAxisClamp1.bExeStop := FALSE;
END_ACTION

ACTION Gr05Auto_eAxisClamp2InPos_Exit:
Gr05Control.fbCylinderPos.bExeMoveAbs := FALSE;
END_ACTION

ACTION Gr05Auto_eAxisClamp2InPos2_Exit:
Gr05Control.fbCylinderPos.bExeMoveAbs := FALSE;
END_ACTION

ACTION Gr05Auto_eAxisClamp2InPos2Err_Entry:
Gr05Control.fbCylinderPos.bExeMoveAbs := FALSE;
END_ACTION

ACTION Gr05Auto_eAxisClamp2InPosErr_Entry:
Gr05Control.fbCylinderPos.bExeMoveAbs := FALSE;
END_ACTION

ACTION Gr05Auto_eAxisClamp2InSawBandPos_Exit:
Gr05Control.fbCylinderPos.bExeMoveAbs := FALSE;
END_ACTION

ACTION Gr05Auto_eAxisClamp2InSawBandPosErr_Entry:
Gr05Control.fbCylinderPos.bExeMoveAbs := FALSE;
END_ACTION

ACTION Gr05Auto_eAxisClamp2InSawPos_Exit:
Gr05Control.fbCylinderPos.bExeMoveAbs := FALSE;
END_ACTION

ACTION Gr05Auto_eAxisClamp2InSawPosErr_Entry:
Gr05Control.fbCylinderPos.bExeMoveAbs := FALSE;
END_ACTION

ACTION Gr05Auto_eAxisClamp2MoveSawPos_Entry:
Gr05Control.fbCylinderPos.bExeMoveAbs := TRUE;
Gr05Control.fbCylinderPos.lrTargetPosition := lrgGr05Clamp2SawPos; (* 0.0 *)
END_ACTION

ACTION Gr05Auto_eAxisClamp2MoveSawPosErr_Entry:
Gr05Control.fbCylinderPos.bExeMoveAbs := FALSE;
END_ACTION

ACTION Gr05Auto_eAxisClamp2MoveToPos_Entry:
(*IF (lrClamp2Pos - lrgGr05Clamp2Width) > stgGr05HMI.stPLCTOHMI.lrAxisClamp2ActPos
THEN*)
	Gr05Control.fbCylinderPos.bExeMoveAbs := TRUE;
(*ELSE
	Gr05Control.fbCylinderPos.bExeMoveAbs := stgGr05HMI.stPLCTOHMI.lrAxisClamp1ActPos < (lrClamp2Pos - lrgGr05Clamp2Width);
END_IF*)

Gr05Control.fbCylinderPos.lrTargetPosition := lrClamp2Pos;
END_ACTION

ACTION Gr05Auto_eAxisClamp2MoveToPos2_Entry:
Gr05Control.fbCylinderPos.bExeMoveAbs := TRUE;
IF ABS(lrActSawingLength) < ABS(lrClamp1Pos - lrgGr05Clamp2Width)
THEN
	IF Gr05Control.fbCylinderPos.lrActPosition < (lrClamp1Pos - ABS(lrActSawingLength) - lrgGr05Clamp2Width)
	THEN
		Gr05Control.fbCylinderPos.lrTargetPosition := Gr05Control.fbCylinderPos.lrActPosition;
	ELSE
		Gr05Control.fbCylinderPos.lrTargetPosition := lrClamp1Pos - ABS(lrActSawingLength) - lrgGr05Clamp2Width;
	END_IF
ELSE
	Gr05Control.fbCylinderPos.lrTargetPosition := 0.0;
END_IF
END_ACTION

ACTION Gr05Auto_eAxisClamp2MoveToPos2Err_Entry:
Gr05Control.fbCylinderPos.bExeMoveAbs := FALSE;
END_ACTION

ACTION Gr05Auto_eAxisClamp2MoveToPosErr_Entry:
Gr05Control.fbCylinderPos.bExeMoveAbs := FALSE;
END_ACTION

ACTION Gr05Auto_eAxisClamp2MoveToSawBandPos_Entry:
Gr05Control.fbCylinderPos.bExeMoveAbs := TRUE;
Gr05Control.fbCylinderPos.lrTargetPosition := lrgGr05Clamp2PipeBeginPos;  (*0*)
END_ACTION

ACTION Gr05Auto_eAxisClamp2MoveToSawBandPosErr_Entry:
Gr05Control.fbCylinderPos.bExeMoveAbs := FALSE;
END_ACTION

ACTION Gr05Auto_eChkAxisClamp1MoveToBackPos_Entry:
(*ESKG 12032026*)

IF ABS(lrActSawingLength) >= ABS(lrActRemoveLength)
THEN
	bSafetyDistEnable := ((Gr05Control.fbAxisClamp1.lrActPosition - Gr05Control.fbCylinderPos.lrActPosition - lrgGr05Clamp2Width ) <  lrgGr05SafetyDistance)
						AND Gr05Control.fbUtility.bPipeEndPresent;

	IF bSafetyDistEnable
	THEN
		lrActSawingLength := 0;
		lrActRemoveLength := 0;
	END_IF
END_IF
END_ACTION

ACTION Gr05Auto_eChkAxisClamp1MoveToBackPos_Exit:
Gr05Control.fbAxisClamp1.bExeMoveAbs := FALSE;
END_ACTION

ACTION Gr05Auto_eChkWorkArea_Entry:
lrClamp1PosCache := lrClamp1Pos;
END_ACTION

ACTION Gr05Auto_eClamp12Open_Entry:
Gr05Control.arfbCylinderClamp[1].bAutoOpen := TRUE;					(* Auto open *)
Gr05Control.arfbCylinderClamp[1].bAutoClose := FALSE;					(* Auto close *)
(*Gr05Control.arfbCylinderClamp[2].bAutoOpen := TRUE;				(* Auto open *)
Gr05Control.arfbCylinderClamp[2].bAutoClose := FALSE;					(* Auto close *)*)
END_ACTION

ACTION Gr05Auto_eClamp12Open_Exit:
Gr05Control.arfbCylinderClamp[1].bAutoOpen := FALSE;					(* Auto open *)
Gr05Control.arfbCylinderClamp[1].bAutoClose := FALSE;					(* Auto close *)
Gr05Control.arfbCylinderClamp[2].bAutoOpen := FALSE;					(* Auto open *)
Gr05Control.arfbCylinderClamp[2].bAutoClose := FALSE;					(* Auto close *)
END_ACTION

ACTION Gr05Auto_eClamp1Close_Entry:

Gr05Control.arfbCylinderClamp[1].bAutoOpen := FALSE;										(* Auto open *)
Gr05Control.arfbCylinderClamp[1].bAutoClose := NOT binGr05PipeBeginEdge;					(*ESKG 12032026*)			(* Auto close *)
END_ACTION

ACTION Gr05Auto_eClamp1Close_Exit:
Gr05Control.arfbCylinderClamp[1].bAutoOpen := FALSE;					(* Auto open *)
Gr05Control.arfbCylinderClamp[1].bAutoClose := FALSE;					(* Auto close *)
END_ACTION

ACTION Gr05Auto_eClamp1Close2_Entry:

Gr05Control.arfbCylinderClamp[1].bAutoOpen := FALSE;					(* Auto open *)
Gr05Control.arfbCylinderClamp[1].bAutoClose := TRUE;					(* Auto close *)
END_ACTION

ACTION Gr05Auto_eClamp1Close2_Exit:
Gr05Control.arfbCylinderClamp[1].bAutoOpen := FALSE;					(* Auto open *)
Gr05Control.arfbCylinderClamp[1].bAutoClose := FALSE;					(* Auto close *)
END_ACTION

ACTION Gr05Auto_eClamp1Close2Err_Entry:
Gr05Control.arfbCylinderClamp[1].bAutoOpen := FALSE;					(* Auto open *)
Gr05Control.arfbCylinderClamp[1].bAutoClose := FALSE;					(* Auto close *)
END_ACTION

ACTION Gr05Auto_eClamp1Close3_Entry:
Gr05Control.arfbCylinderClamp[1].bAutoOpen := FALSE;					(* Auto open *)
Gr05Control.arfbCylinderClamp[1].bAutoClose := TRUE;					(* Auto close *)
END_ACTION

ACTION Gr05Auto_eClamp1Close3_Exit:
Gr05Control.arfbCylinderClamp[1].bAutoOpen := FALSE;					(* Auto open *)
Gr05Control.arfbCylinderClamp[1].bAutoClose := FALSE;					(* Auto close *)
END_ACTION

ACTION Gr05Auto_eClamp1Close3Err_Entry:
Gr05Control.arfbCylinderClamp[1].bAutoOpen:= FALSE;					(* Auto open *)
Gr05Control.arfbCylinderClamp[1].bAutoClose := FALSE;					(* Auto close *)
END_ACTION

ACTION Gr05Auto_eClamp1CloseErr_Entry:
Gr05Control.arfbCylinderClamp[1].bAutoOpen := FALSE;					(* Auto open *)
Gr05Control.arfbCylinderClamp[1].bAutoClose := FALSE;					(* Auto close *)
END_ACTION

ACTION Gr05Auto_eClamp1Open_Entry:
Gr05Control.arfbCylinderClamp[1].bAutoOpen := TRUE;					(* Auto open *)
Gr05Control.arfbCylinderClamp[1].bAutoClose := FALSE;					(* Auto close *)
END_ACTION

ACTION Gr05Auto_eClamp1Open_Exit:
Gr05Control.arfbCylinderClamp[1].bAutoOpen := FALSE;					(* Auto open *)
Gr05Control.arfbCylinderClamp[1].bAutoClose := FALSE;					(* Auto close *)
END_ACTION

ACTION Gr05Auto_eClamp1Open2Err_Entry:
Gr05Control.arfbCylinderClamp[1].bAutoOpen := FALSE;					(* Auto open *)
Gr05Control.arfbCylinderClamp[1].bAutoClose := FALSE;					(* Auto close *)
END_ACTION

ACTION Gr05Auto_eClamp1OpenErr_Entry:
Gr05Control.arfbCylinderClamp[1].bAutoOpen := FALSE;					(* Auto open *)
Gr05Control.arfbCylinderClamp[1].bAutoClose := FALSE;					(* Auto close *)
END_ACTION

ACTION Gr05Auto_eClamp2Close_Entry:
Gr05Control.arfbCylinderClamp[2].bAutoOpen := FALSE;					(* Auto open *)
Gr05Control.arfbCylinderClamp[2].bAutoClose := TRUE;					(* Auto close *)
END_ACTION

ACTION Gr05Auto_eClamp2Close_Exit:
Gr05Control.arfbCylinderClamp[2].bAutoOpen := FALSE;					(* Auto open *)
Gr05Control.arfbCylinderClamp[2].bAutoClose := FALSE;					(* Auto close *)
END_ACTION

ACTION Gr05Auto_eClamp2CloseErr_Entry:
Gr05Control.arfbCylinderClamp[2].bAutoOpen := FALSE;					(* Auto open *)
Gr05Control.arfbCylinderClamp[2].bAutoClose := FALSE;					(* Auto close *)
END_ACTION

ACTION Gr05Auto_eClamp2Err_Entry:
Gr05Control.arfbCylinderClamp[2].bAutoOpen := FALSE;					(* Auto open *)
Gr05Control.arfbCylinderClamp[2].bAutoClose := FALSE;					(* Auto close *)
END_ACTION

ACTION Gr05Auto_eClamp2Open_Entry:
Gr05Control.arfbCylinderClamp[2].bAutoOpen := TRUE;					(* Auto open *)
Gr05Control.arfbCylinderClamp[2].bAutoClose := FALSE;					(* Auto close *)
END_ACTION

ACTION Gr05Auto_eClamp2Open_Exit:
Gr05Control.arfbCylinderClamp[2].bAutoOpen := FALSE;					(* Auto open *)
Gr05Control.arfbCylinderClamp[2].bAutoClose := FALSE;					(* Auto close *)
END_ACTION

ACTION Gr05Auto_eClamp2Open1_Entry:
Gr05Control.arfbCylinderClamp[2].bAutoOpen :=	(Gr05Control.fbCylinderPos.lrActPosition <> lrClamp2Pos )   	(*ESKG 12032026*)
											OR	lrClamp1PosCache <> (lrClamp1Pos - MAX(ABS(lrActSawingLength), ABS(lrActRemoveLength)));					(* Auto open *)
Gr05Control.arfbCylinderClamp[2].bAutoClose := FALSE;					(* Auto close *)
END_ACTION

ACTION Gr05Auto_eClamp2Open1_Exit:
Gr05Control.arfbCylinderClamp[2].bAutoOpen := FALSE;					(* Auto open *)
Gr05Control.arfbCylinderClamp[2].bAutoClose := FALSE;					(* Auto close *)
END_ACTION

ACTION Gr05Auto_eClamp2Open1Err_Entry:
Gr05Control.arfbCylinderClamp[2].bAutoOpen := FALSE;					(* Auto open *)
Gr05Control.arfbCylinderClamp[2].bAutoClose := FALSE;					(* Auto close *)
END_ACTION

ACTION Gr05Auto_eClamp2Open2Err_Entry:
Gr05Control.arfbCylinderClamp[2].bAutoOpen := FALSE;					(* Auto open *)
Gr05Control.arfbCylinderClamp[2].bAutoClose := FALSE;					(* Auto close *)
END_ACTION

ACTION Gr05Auto_eClamp2Open3_Entry:
Gr05Control.arfbCylinderClamp[2].bAutoOpen := TRUE;					(* Auto open *)
Gr05Control.arfbCylinderClamp[2].bAutoClose := FALSE;					(* Auto close *)
END_ACTION

ACTION Gr05Auto_eClamp2Open3_Exit:
Gr05Control.arfbCylinderClamp[2].bAutoOpen := FALSE;					(* Auto open *)
Gr05Control.arfbCylinderClamp[2].bAutoClose := FALSE;					(* Auto close *)
END_ACTION

ACTION Gr05Auto_eClamp2Open3Err_Entry:
Gr05Control.arfbCylinderClamp[2].bAutoOpen := FALSE;					(* Auto open *)
Gr05Control.arfbCylinderClamp[2].bAutoClose := FALSE;					(* Auto close *)
END_ACTION

ACTION Gr05Auto_eClamp2OpenErr_Entry:
Gr05Control.arfbCylinderClamp[2].bAutoOpen := FALSE;					(* Auto open *)
Gr05Control.arfbCylinderClamp[2].bAutoClose := FALSE;					(* Auto close *)
END_ACTION

ACTION Gr05Auto_eClamp2Slide_Entry:
Gr05Control.arfbCylinderClamp[2].bAutoOpen := FALSE;					(* Auto open *)
Gr05Control.arfbCylinderClamp[2].bAutoClose := TRUE;					(* Auto close *)
Gr05Control.fbSlide.bAutoMoveToBase := TRUE;						(* Auto move to base *)
Gr05Control.fbSlide.bAutoMoveToWork := FALSE;						(* Auto move to work *)

Gr05Control.fbRemovalBand.arbAutoMoveToMinus[2] := FALSE;			(* Auto move to minus *)

(*ESKG 12032026*)
bSafetyDistEnable:= FALSE;
END_ACTION

ACTION Gr05Auto_eClamp2Slide_Exit:
Gr05Control.arfbCylinderClamp[2].bAutoOpen := FALSE;					(* Auto open *)
Gr05Control.arfbCylinderClamp[2].bAutoClose := FALSE;					(* Auto close *)
Gr05Control.fbSlide.bAutoMoveToBase := FALSE;				(* Auto move to base *)
Gr05Control.fbSlide.bAutoMoveToWork := FALSE;				(* Auto move to work *)
END_ACTION

ACTION Gr05Auto_eCollisionDetectedErr_Entry:
bErrorCollisionDetected := TRUE;
END_ACTION

ACTION Gr05Auto_eCollisionDetectedErr_Exit:
bErrorCollisionDetected := FALSE;
udnErrorNo := 3;
END_ACTION

ACTION Gr05Auto_eDone_Entry:
bDone := TRUE;                                      		(* Program done, in position *)
bBusy := FALSE;                                     		(* Program not busy *)
END_ACTION

ACTION Gr05Auto_eDone_Exit:
bDone := FALSE;                                 	(* Program done *)
bBusy := FALSE;                                 	(* Program not busy *)
bError := FALSE;                                		(* Program not error *)
END_ACTION

ACTION Gr05Auto_eError_Entry:
bDone := FALSE;                                    	 	(* Program done, in position *)
bError := TRUE;                                     		(* Program error *)
bBusy := FALSE;                                     		(* Program not busy *)
END_ACTION

ACTION Gr05Auto_eError_Exit:
bDone := FALSE;                                 	(* Program done *)
bBusy := FALSE;                                 	(* Program not busy *)
bError := FALSE;                                		(* Program not error *)
END_ACTION

ACTION Gr05Auto_eGetClamp1ActPos_01_Entry:
lrClamp1Pos := Gr05Control.fbAxisClamp1.lrActPosition;
END_ACTION

ACTION Gr05Auto_eGetClamp1ActPos_02_Entry:
lrClamp1Pos := Gr05Control.fbAxisClamp1.lrActPosition;
END_ACTION

ACTION Gr05Auto_eGetClamp1ActPos_03_Entry:
lrClamp1Pos := Gr05Control.fbAxisClamp1.lrActPosition;
END_ACTION

ACTION Gr05Auto_eGetClamp1ActPos_04_Entry:
lrClamp1Pos := Gr05Control.fbAxisClamp1.lrActPosition;
END_ACTION

ACTION Gr05Auto_eGetClamp1ActPos_05_Entry:
lrClamp1Pos := Gr05Control.fbAxisClamp1.lrActPosition;
END_ACTION

ACTION Gr05Auto_eGetClamp1ActPos_06_Entry:
lrActRemoveLength := 0.0;
lrClamp1Pos := Gr05Control.fbAxisClamp1.lrActPosition;
END_ACTION

ACTION Gr05Auto_eGetClamp1ActPos_Entry:
lrClamp1Pos := Gr05Control.fbAxisClamp1.lrActPosition;
END_ACTION

ACTION Gr05Auto_eGetClamp2ActPos_Entry:

lrClamp2Pos := F_AxisClamp2Pos(
					bEnable := TRUE,
					lrActClamp2Pos := Gr05Control.fbCylinderPos.lrActPosition,
					lrAngle := lrActSawingAngle,
					lrRadius := stgGr01HMI.stHMITOPLC.rPipeDiameter / 2.0,
					lrPipeClampWidth := lrgGr05PipeClampWidth,
					lrSawbandGuideWidth := lrgGr05SawbandGuideWidth
				);
END_ACTION

ACTION Gr05Auto_eGetProcessPara_Entry:
IF unProcessCounter <= usnFileArrayMaxDimR
THEN
	unProcessCounter := unProcessCounter + 1;

	IF unProcessCounter > 1
	THEN
		lrActRemoveLength := lrgGr05RemovalBandSawBand;
	ELSE
		lrActRemoveLength := 0.0;
	END_IF

	stgGr05HMI.stHMITOPLC.lrActSawingLength := REAL_TO_LREAL(ABS(arrGr00ProcessPara[unProcessCounter,0]));
	lrActSawingLength := SEL(
							stgGr05HMI.stHMITOPLC.lrActSawingLength > 0,
						    	0.0,
						    	REAL_TO_LREAL(ABS(arrGr00ProcessPara[unProcessCounter,0]) +
							(stgGr01HMI.stHMITOPLC.lrSawBandThickness * (1/COS(ABS(arrGr00ProcessPara[unProcessCounter, 1] / 180 * PI)))))
						     );
	(*lrActSawingLength := ABS(arrGr00ProcessPara[unProcessCounter,0]) + (stgGr01HMI.stHMITOPLC.lrSawBandThickness * 1);*)
	lrActSawingAngle := REAL_TO_LREAL(arrGr00ProcessPara[unProcessCounter, 1] / 180 * PI);

	(*ESKG 12032026*)
	IF lrActSawingLength>=lrActRemoveLength
	THEN
		lrActRemoveLength := 0.0;
	END_IF

END_IF
END_ACTION

ACTION Gr05Auto_eRemovalBandErr_Entry:
Gr05Control.fbRemovalBand.arbAutoMoveToMinus[2] := FALSE;				(* Auto move to minus *)
END_ACTION

ACTION Gr05Auto_eSawbandStart_Entry:
Gr01Control.fbSawband.bExeMoveVelo:= TRUE;
Gr01Control.fbSawband.lrAutoVelocity := stgGr01HMI.stHMITOPLC.rSawbandAutoSpeed / 3.28084;
END_ACTION

ACTION Gr05Auto_eSawbandStart_Exit:
Gr01Control.fbSawband.bExeMoveVelo:= FALSE;
END_ACTION

ACTION Gr05Auto_eSawingLengthCorrection_Entry:
stgGr05HMI.stHMITOPLC.lrActSawingLength := MAX(0, ABS(stgGr05HMI.stHMITOPLC.lrActSawingLength) - ABS(lrClamp1Pos - Gr05Control.fbAxisClamp1.lrActPosition));
lrActSawingLength := MAX(0, ABS(lrActSawingLength) - ABS(lrClamp1Pos - Gr05Control.fbAxisClamp1.lrActPosition));
END_ACTION

ACTION Gr05Auto_eSawingReq_Entry:
bgGr05SawingReq := TRUE;
END_ACTION

ACTION Gr05Auto_eSawingReq_Exit:
bgGr05SawingReq := FALSE;
END_ACTION

ACTION Gr05Auto_eSlideDown_Entry:
Gr05Control.fbSlide.bAutoMoveToBase := FALSE;					(* Auto move to base *)
Gr05Control.fbSlide.bAutoMoveToWork := stgGr05HMI.stHMITOPLC.bSlideActive;					(* Auto move to work *)

Gr05Control.fbRemovalBand.arbAutoMoveToMinus[2] := TRUE;				(* Auto move to minus *)
END_ACTION

ACTION Gr05Auto_eSlideDownErr_Entry:
Gr05Control.fbSlide.bAutoMoveToBase := FALSE;				(* Auto move to base *)
Gr05Control.fbSlide.bAutoMoveToWork := FALSE;				(* Auto move to work *)
END_ACTION

ACTION Gr05Auto_eSlideUpErr_Entry:
Gr05Control.fbSlide.bAutoMoveToBase := FALSE;				(* Auto move to base *)
Gr05Control.fbSlide.bAutoMoveToWork := FALSE;				(* Auto move to work *)
END_ACTION

ACTION Gr05Auto_eTransportAck_Exit:
bgGr05TransportAck := FALSE;
END_ACTION

ACTION Gr05Auto_eWfAxisClamp1MoveAbsPipeEnde_Exit:
Gr05Control.fbAxisClamp1.bExeMoveAbs := FALSE;
END_ACTION

ACTION Gr05Auto_eWfAxisClamp1MoveAbsPipeEndeErr_Entry:
Gr05Control.fbAxisClamp1.bExeMoveAbs := FALSE;
END_ACTION

ACTION Gr05Auto_eWfAxisClamp1MoveVeloPipeBegin_Exit:
Gr05Control.fbAxisClamp1.bExeMoveVelo := FALSE;
END_ACTION

ACTION Gr05Auto_eWfAxisClamp1MoveVeloPipeBeginErr_Entry:
Gr05Control.fbAxisClamp1.bExeMoveVelo := FALSE;
END_ACTION

ACTION Gr05Auto_eWfAxisClamp1MoveVeloPipeEnd_Exit:
Gr05Control.fbAxisClamp1.bExeMoveVelo := FALSE;
END_ACTION

ACTION Gr05Auto_eWfAxisClamp1MoveVeloPipeEndErr_Entry:
Gr05Control.fbAxisClamp1.bExeMoveVelo := FALSE;
END_ACTION

ACTION Gr05Auto_eWfAxisClamp1Stop_2_Exit:
Gr05Control.fbAxisClamp1.bExeStop := FALSE;
END_ACTION

ACTION Gr05Auto_eWfAxisClamp1Stop_Exit:
Gr05Control.fbAxisClamp1.bExeStop := FALSE;
END_ACTION

ACTION Gr05Auto_eWfAxisClamp1StopErr_2_Entry:
Gr05Control.fbAxisClamp1.bExeStop := FALSE;
END_ACTION

ACTION Gr05Auto_eWfAxisClamp1StopErr_Entry:
Gr05Control.fbAxisClamp1.bExeStop := FALSE;
END_ACTION

ACTION Gr05Auto_eWfPipeBeginNoDetectedError_Entry:
bErrorPipeBeginNoDetected := TRUE;
END_ACTION

ACTION Gr05Auto_eWfPipeBeginNoDetectedError_Exit:
bErrorPipeBeginNoDetected := FALSE;
END_ACTION

ACTION Gr05Auto_eWfPipeBeginNoDetectedWarrning_Entry:
bWarningPipeBeginNoDetected := TRUE;
END_ACTION

ACTION Gr05Auto_eWfPipeBeginNoDetectedWarrning_Exit:
bWarningPipeBeginNoDetected := FALSE;
END_ACTION

ACTION Gr05Auto_eWfPipeEndNoDetectedErr_Entry:
bErrorPipeEndNoDetected := TRUE;
END_ACTION

ACTION Gr05Auto_eWfPipeEndNoDetectedErr_Exit:
bErrorPipeEndNoDetected := FALSE;
udnErrorNo := 2;
END_ACTION

ACTION Gr05Auto_eWfTransportReq_Exit:
bgGr05TransportAck := TRUE;
END_ACTION

ACTION Init_Action:
IF NOT bFirstTime
THEN
	SFCCurrentStep:= 'Init';

	bDone := FALSE;                                 	(* Program done *)
	bBusy := FALSE;                                  	(* Program not busy *)
	bError := FALSE;                                 	(* Program not error *)
	udnErrorNo := 0;                                		(* Error number *)
	
	(* Internal flags *)
	bgGr05SawingReq := FALSE;
	bgGr05AngleReq := FALSE;
	bgGr05TransportAck := FALSE;
	unProcessCounter	 := 0;

	bErrorPipeBeginNoDetected := FALSE;
	bErrorPipeEndNoDetected := FALSE;
	bWarningPipeBeginNoDetected := FALSE;
	(*ESKG 12032026*)
	bSafetyDistEnable := FALSE;

	bFirstTime := TRUE;
END_IF
END_ACTION

ACTION Init_Exit:
(* Set status *)
bDone := FALSE;                                 	(* Program done *)
bBusy := FALSE;                                  	(* Program not busy *)
bError := FALSE;                                 	(* Program not error *)
udnErrorNo := 0;                                		(* Error number *)

(* Internal flags *)
bgGr05SawingReq := FALSE;
bgGr05AngleReq := FALSE;
bgGr05TransportAck := FALSE;
unProcessCounter	 := 0;
bPipeEndDetected := FALSE;
rtPipeBeginIdentify(CLK := FALSE);
rtPipeEndIdentify(CLK := FALSE);

bErrorPipeBeginNoDetected := FALSE;
bErrorPipeEndNoDetected := FALSE;
bWarningPipeBeginNoDetected := FALSE;

(*ESKG 12032026*)
bSafetyDistEnable:= FALSE;
END_ACTION

TRANSITION SafetyDistEnable:
bSafetyDistEnable  	(*ESKG 12032026*)
AND Gr05Control.arfbCylinderClamp[1].fbCylinder.bEndWork
AND bReleaseNextStep
END_TRANSITION

TRANSITION SafetyDistEnable_1:
	(*ESKG 12032026*)
(*(Gr05Control.fbAxisClamp1.lrActPosition - Gr05Control.fbCylinderPos.lrActPosition - lrgGr05Clamp2Width ) <  lrgGr05SafetyDistance*)
bSafetyDistEnable
END_TRANSITION

TRANSITION Trans:
Gr05Control.bAllAxisCtrlEnabled
END_TRANSITION

TRANSITION Trans_1:
(Gr05Control.arfbCylinderClamp[1].fbCylinder.bEndWork OR  binGr05PipeBeginEdge)
AND bReleaseNextStep
END_TRANSITION

TRANSITION Trans_10:
bReleaseNextStep
END_TRANSITION

TRANSITION Trans_100:
NOT bExecute
END_TRANSITION

TRANSITION Trans_101:
NOT bExecute
END_TRANSITION

TRANSITION Trans_11:
Gr01Control.fbSawband.fbMoveAuto.fbMCMoveVelo.Busy
END_TRANSITION

TRANSITION Trans_12:
stgGr05Alarm.stAuto.arbError[0].bActive
END_TRANSITION

TRANSITION Trans_13:
stgGr05Alarm.stAuto.arbWarning[0].bActive
END_TRANSITION

TRANSITION Trans_14:
Gr05Control.fbAxisClamp1.fbMoveAuto.fbMCMoveAbs.Busy
END_TRANSITION

TRANSITION Trans_15:
Gr05Control.fbAxisClamp1.fbMoveAuto.fbMCMoveAbs.Error
END_TRANSITION

TRANSITION Trans_16:
Gr05Control.fbAxisClamp1.fbMoveAuto.bInPosition
AND bReleaseNextStep
END_TRANSITION

TRANSITION Trans_17:
Gr05Control.fbAxisClamp1.fbMoveAuto.fbMCMoveAbs.Error
END_TRANSITION

TRANSITION Trans_18:
Gr05Control.fbCylinderPos.fbMoveAbs.bBusy
END_TRANSITION

TRANSITION Trans_19:
Gr05Control.fbCylinderPos.fbMoveAbs.bError
END_TRANSITION

TRANSITION Trans_2:
Gr05Control.arfbCylinderClamp[1].bErrorClose
END_TRANSITION

TRANSITION Trans_20:
Gr05Control.fbCylinderPos.fbMoveAbs.bDone
AND bReleaseNextStep
END_TRANSITION

TRANSITION Trans_21:
Gr05Control.fbCylinderPos.fbMoveAbs.bError
END_TRANSITION

TRANSITION Trans_22:
Gr05Control.fbCylinderPos.fbMoveAbs.bBusy
END_TRANSITION

TRANSITION Trans_23:
Gr05Control.fbCylinderPos.fbMoveAbs.bError
END_TRANSITION

TRANSITION Trans_24:
Gr05Control.fbCylinderPos.fbMoveAbs.bDone
AND bReleaseNextStep
END_TRANSITION

TRANSITION Trans_25:
Gr05Control.fbCylinderPos.fbMoveAbs.bError
END_TRANSITION

TRANSITION Trans_26:
unProcessCounter >= usnFileArrayMaxDimR
AND bReleaseNextStep
END_TRANSITION

TRANSITION Trans_27:
arrGr00ProcessPara[unProcessCounter, 0] > 0.0
OR arrGr00ProcessPara[unProcessCounter, 1] <> 0.0
END_TRANSITION

TRANSITION Trans_28:
(Gr05Control.fbSlide.fbCylinder.bEndBase
OR NOT Gr05Control.fbSlide.bEnable)
AND bReleaseNextStep
END_TRANSITION

TRANSITION Trans_29:
(stgGr05HMI.stHMITOPLC.bCylinderPosActive
OR lrClamp2Pos <= Gr05Control.fbCylinderPos.lrActPosition)
AND bReleaseNextStep
END_TRANSITION

TRANSITION Trans_3:
NOT binGr05PipeBeginEdge
AND bReleaseNextStep
END_TRANSITION

TRANSITION Trans_30:
stgGr05Alarm.stAuto.arbError[2].bActive
END_TRANSITION

TRANSITION Trans_31:
Gr05Control.arfbCylinderClamp[1].fbCylinder.bEndWork
AND bReleaseNextStep
END_TRANSITION

TRANSITION Trans_32:
Gr05Control.arfbCylinderClamp[1].bErrorClose
END_TRANSITION

TRANSITION Trans_33:
((Gr05Control.arfbCylinderClamp[2].fbCylinder.bEndBase OR NOT Gr05Control.arfbCylinderClamp[2].bAutoOpen )
OR ( lrClamp1PosCache = (lrClamp1Pos - MAX(ABS(lrActSawingLength), ABS(lrActRemoveLength))+0.2)
))

AND bReleaseNextStep

(* +0.2 this is just an offset works in this case as a delay until the EndBase comes *)
END_TRANSITION

TRANSITION Trans_34:
Gr05Control.arfbCylinderClamp[2].bErrorOpen
END_TRANSITION

TRANSITION Trans_35:
Gr05Control.fbAxisClamp1.fbMoveAuto.fbMCMoveAbs.Busy
END_TRANSITION

TRANSITION Trans_36:
Gr05Control.fbAxisClamp1.fbMoveAuto.fbMCMoveAbs.Error
END_TRANSITION

TRANSITION Trans_37:
Gr05Control.fbAxisClamp1.fbMoveAuto.bInPosition
AND bReleaseNextStep
END_TRANSITION

TRANSITION Trans_38:
Gr05Control.fbAxisClamp1.fbMoveAuto.fbMCMoveAbs.Error
END_TRANSITION

TRANSITION Trans_39:
Gr05Control.fbCylinderPos.fbMoveAbs.bBusy
END_TRANSITION

TRANSITION Trans_4:
Gr05Control.arfbCylinderClamp[2].fbCylinder.bEndBase
AND bReleaseNextStep
END_TRANSITION

TRANSITION Trans_40:
Gr05Control.fbCylinderPos.fbMoveAbs.bError
END_TRANSITION

TRANSITION Trans_41:
Gr05Control.fbCylinderPos.fbMoveAbs.bDone
AND bReleaseNextStep
END_TRANSITION

TRANSITION Trans_42:
Gr05Control.fbCylinderPos.fbMoveAbs.bError
END_TRANSITION

TRANSITION Trans_43:
Gr05Control.fbAxisClamp1.fbMoveAuto.fbMCMoveAbs.Busy
END_TRANSITION

TRANSITION Trans_44:
Gr05Control.fbAxisClamp1.fbMoveAuto.fbMCMoveAbs.Error
END_TRANSITION

TRANSITION Trans_45:
Gr05Control.fbAxisClamp1.fbMoveAuto.bInPosition
AND bReleaseNextStep
END_TRANSITION

TRANSITION Trans_46:
Gr05Control.fbAxisClamp1.fbMoveAuto.fbMCMoveAbs.Error
END_TRANSITION

TRANSITION Trans_47:
Gr05Control.arfbCylinderClamp[2].fbCylinder.bEndWork
AND (Gr05Control.fbSlide.fbCylinder.bEndBase OR NOT Gr05Control.fbSlide.bEnable)
AND bReleaseNextStep
END_TRANSITION

TRANSITION Trans_48:
Gr05Control.arfbCylinderClamp[2].bErrorOpen
END_TRANSITION

TRANSITION Trans_49:
Gr05Control.fbSlide.bErrorMoveToBase
END_TRANSITION

TRANSITION Trans_5:
Gr05Control.arfbCylinderClamp[2].bErrorOpen
END_TRANSITION

TRANSITION Trans_50:
bgGr01SawingAck
AND bReleaseNextStep
END_TRANSITION

TRANSITION Trans_51:
NOT bgGr01SawingAck
AND bReleaseNextStep
END_TRANSITION

TRANSITION Trans_52:
bgGr01TransportReq
AND bReleaseNextStep
END_TRANSITION

TRANSITION Trans_53:
NOT bgGr01TransportReq
AND bReleaseNextStep
END_TRANSITION

TRANSITION Trans_54:
(NOT Gr05Control.fbSlide.fbCylinder.bEndBase
OR NOT Gr05Control.fbSlide.bEnable)
AND bReleaseNextStep
END_TRANSITION

TRANSITION Trans_55:
Gr05Control.fbSlide.bErrorMoveToWork
END_TRANSITION

TRANSITION Trans_56:
Gr05Control.fbRemovalBand.bErrorMoveToMinus
OR Gr05Control.fbRemovalBand.bErrorMoveToPlus
END_TRANSITION

TRANSITION Trans_57:
Gr05Control.arfbCylinderClamp[2].fbCylinder.bEndWork
AND bReleaseNextStep
END_TRANSITION

TRANSITION Trans_58:
Gr05Control.arfbCylinderClamp[2].bErrorClose
END_TRANSITION

TRANSITION Trans_59:
Gr05Control.arfbCylinderClamp[1].fbCylinder.bEndBase
AND bReleaseNextStep
END_TRANSITION

TRANSITION Trans_6:
Gr05Control.fbAxisClamp1.fbMoveAuto.fbMCMoveVelo.Busy
END_TRANSITION

TRANSITION Trans_60:
Gr05Control.arfbCylinderClamp[1].bErrorOpen
END_TRANSITION

TRANSITION Trans_61:
NOT binGr05PipeEndEdge
OR Gr05Control.fbAxisClamp1.fbMoveAuto.fbMCMoveAbs.Busy
END_TRANSITION

TRANSITION Trans_62:
Gr05Control.fbAxisClamp1.fbMoveAuto.fbMCMoveAbs.Error
END_TRANSITION

TRANSITION Trans_63:
Gr05Control.fbAxisClamp1.fbMoveAuto.fbMCStop.Busy
END_TRANSITION

TRANSITION Trans_64:
Gr05Control.fbAxisClamp1.fbMoveAuto.fbMCStop.Error
END_TRANSITION

TRANSITION Trans_65:
Gr05Control.fbAxisClamp1.fbMoveAuto.bStopped
AND Gr05Control.fbAxisClamp1.lrActVelocity = 0.0
AND bReleaseNextStep
END_TRANSITION

TRANSITION Trans_66:
Gr05Control.fbAxisClamp1.fbMoveAuto.fbMCStop.Error
END_TRANSITION

TRANSITION Trans_67:
unProcessCounter > 1
AND arrGr00ProcessPara[unProcessCounter, 1] / 180 * PI = 0.0								(* Check next sawing angle *)
AND bReleaseNextStep
END_TRANSITION

TRANSITION Trans_68:
Gr05Control.fbAxisClamp1.fbMoveAuto.fbMCMoveVelo.Busy
END_TRANSITION

TRANSITION Trans_69:
Gr05Control.fbAxisClamp1.fbMoveAuto.fbMCMoveVelo.Error
END_TRANSITION

TRANSITION Trans_7:
Gr05Control.fbAxisClamp1.fbMoveAuto.fbMCMoveVelo.Error
END_TRANSITION

TRANSITION Trans_70:
Gr05Control.fbAxisClamp1.fbMoveAuto.bInVelocity
AND bReleaseNextStep
END_TRANSITION

TRANSITION Trans_71:
Gr05Control.fbAxisClamp1.fbMoveAuto.fbMCMoveVelo.Error
END_TRANSITION

TRANSITION Trans_72:
stgGr05Alarm.stAuto.arbError[1].bActive
END_TRANSITION

TRANSITION Trans_73:
Gr05Control.fbAxisClamp1.fbMoveAuto.fbMCStop.Busy
END_TRANSITION

TRANSITION Trans_74:
Gr05Control.fbAxisClamp1.fbMoveAuto.fbMCStop.Error
END_TRANSITION

TRANSITION Trans_75:
Gr05Control.fbAxisClamp1.fbMoveAuto.bStopped
AND Gr05Control.fbAxisClamp1.lrActVelocity = 0.0
AND bReleaseNextStep
END_TRANSITION

TRANSITION Trans_76:
Gr05Control.fbAxisClamp1.fbMoveAuto.fbMCStop.Error
END_TRANSITION

TRANSITION Trans_77:
(*lrClamp1PosPipeEnd > ABS(arrGr00ProcessPara[unProcessCounter, 0])					(* Check next sawing lenght *)*)
lrClamp1PosPipeEnd > MAX(ABS(lrActSawingLength), ABS(lrActRemoveLength))				(* Check next sawing lenght *)
END_TRANSITION

TRANSITION Trans_78:
(* Current pos clamp 1 - sawing lenght > current pos clamp 2 (Current pos clamp 2 is " + ") *)
(lrClamp1Pos - MAX(ABS(lrActSawingLength), ABS(lrActRemoveLength)) > (F_GetCylinderPos(
														F_SetCylinderPos(SEL(stgGr05HMI.stHMITOPLC.bCylinderPosActive, Gr05Control.fbCylinderPos.lrActPosition, lrClamp2Pos),
																		lrgGr05CylinderPosOffset,
																		lrgGr05CylinderPosOriginShiftPos,
																		etgGr05CylinderPosDirection,
																		usngGr05CylinderPosCodingType),
														lrgGr05CylinderPosOffset,
														lrgGr05CylinderPosOriginShiftPos,
														etgGr05CylinderPosDirection,
														usngGr05CylinderPosCodingType)
									    + lrgGr05Clamp2Width))
AND bReleaseNextStep
END_TRANSITION

TRANSITION Trans_79:
bgGr01AngleAck
AND bReleaseNextStep
END_TRANSITION

TRANSITION Trans_8:
Gr05Control.fbAxisClamp1.fbMoveAuto.bInVelocity
AND bReleaseNextStep
END_TRANSITION

TRANSITION Trans_80:
NOT bgGr01AngleAck
AND bReleaseNextStep
END_TRANSITION

TRANSITION Trans_81:
Gr05Control.fbAxisClamp1.fbMoveAuto.bInPosition
END_TRANSITION

TRANSITION Trans_82:
bReleaseNextStep
END_TRANSITION

TRANSITION Trans_83:
Gr05Control.arfbCylinderClamp[1].fbCylinder.bEndWork
AND bReleaseNextStep
END_TRANSITION

TRANSITION Trans_84:
Gr05Control.arfbCylinderClamp[1].bErrorClose
END_TRANSITION

TRANSITION Trans_85:
lrActRemoveLength = 0.0
END_TRANSITION

TRANSITION Trans_86:
Gr05Control.arfbCylinderClamp[2].fbCylinder.bEndBase
AND bReleaseNextStep
END_TRANSITION

TRANSITION Trans_87:
Gr05Control.arfbCylinderClamp[2].bErrorOpen
END_TRANSITION

TRANSITION Trans_88:
Gr05Control.fbCylinderPos.fbMoveAbs.bBusy
END_TRANSITION

TRANSITION Trans_89:
Gr05Control.fbCylinderPos.fbMoveAbs.bError
END_TRANSITION

TRANSITION Trans_9:
Gr05Control.fbAxisClamp1.fbMoveAuto.fbMCMoveVelo.Error
END_TRANSITION

TRANSITION Trans_90:
Gr05Control.fbCylinderPos.fbMoveAbs.bDone
AND bReleaseNextStep
END_TRANSITION

TRANSITION Trans_91:
Gr05Control.fbCylinderPos.fbMoveAbs.bError
END_TRANSITION

TRANSITION Trans_92:
Gr05Control.fbAxisClamp1.fbMoveAuto.fbMCMoveAbs.Busy
END_TRANSITION

TRANSITION Trans_93:
Gr05Control.fbAxisClamp1.fbMoveAuto.fbMCMoveAbs.Error
END_TRANSITION

TRANSITION Trans_94:
Gr05Control.fbAxisClamp1.fbMoveAuto.bInPosition
AND bReleaseNextStep
END_TRANSITION

TRANSITION Trans_95:
Gr05Control.fbAxisClamp1.fbMoveAuto.fbMCMoveAbs.Error
END_TRANSITION

TRANSITION Trans_96:
Gr05Control.fbAxisClamp1.fbMoveAuto.fbMCMoveAbs.Error
END_TRANSITION

TRANSITION Trans_97:
Gr05Control.arfbCylinderClamp[1].fbCylinder.bEndBase
(*AND Gr05Control.arfbCylinderClamp[2].fbCylinder.bEndBase*)
AND bReleaseNextStep
END_TRANSITION

TRANSITION Trans_98:
Gr05Control.arfbCylinderClamp[1].bErrorOpen
END_TRANSITION

TRANSITION Trans_99:
Gr05Control.arfbCylinderClamp[2].bErrorOpen
END_TRANSITION

END_FUNCTION_BLOCK

(* stored: Version 1.1.0.1, ProductVersion 3.1.4024.15
   POU FB_Gr05AutoProcedure: Id {c006d6a3-c91a-4fe7-8398-424f5924b193}, SpecialFunc None
   Transition _Current_pos_clamp_1_sawing_lenght_current_pos_clamp_2_Current_pos_clamp_2_is_: Id {6481c542-76c8-4b43-9684-46d763f37665}
   Transition _Current_pos_clamp_1_sawing_lenght_current_pos_clamp_2_Current_pos_clamp_2_is_1: Id {c65fc21f-bb3b-4cd4-9e8a-6c45a80448ee}
   Transition _No_pipe_end_detected_: Id {91338bbf-53d1-4184-bed6-d73023aafab0}
   Transition _Pipe_begin_was_detected_: Id {f2b07088-bb37-471a-801e-c6ecbaf7a004}
   Transition _Pipe_begin_was_no_detected_: Id {8db41f5e-4a0f-443a-a780-380d1f41a938}
   Transition _Pipe_begin_was_no_detected_1: Id {1e069f00-c6b8-490d-a87a-b080814a921c}
   Transition _Pipe_end_detected_: Id {9e7cd500-a92b-4ee3-a79b-95b5c25ca170}
   Transition _Pipe_end_was_detected_: Id {c5fd9dc7-71cd-428d-bfbf-95b4b388e900}
   Transition _Pipe_end_was_not_detected_: Id {2c869067-fd6f-4c9e-9e22-8aadf3bbb1e4}
   Transition ActSawingL_RemoveL: Id {fe49722e-35f7-4a17-a97f-217c16edbb81}
   Action Gr05Auto_ChkPipeBeginEdge_Exit: Id {7d1101a2-06f3-4b58-bdba-abb1531224e7}
   Action Gr05Auto_eAngleReq_Entry: Id {1d389b3c-9699-4362-b889-d016f35d9696}
   Action Gr05Auto_eAngleReq_Exit: Id {534527a1-8315-4c66-9664-36794cbaf616}
   Action Gr05Auto_eAxisClamp1InBackPos_Exit: Id {82f27437-61a9-45f9-8bc8-d1d22b9b4029}
   Action Gr05Auto_eAxisClamp1InBackPosErr_Entry: Id {c587c135-40d7-4d96-97bc-9cad6350b39d}
   Action Gr05Auto_eAxisClamp1InPipeBeginPos_Action: Id {818575f0-a336-4413-9f5c-e9f2037814b7}
   Action Gr05Auto_eAxisClamp1InPipeBeginPos_Exit: Id {d8b00fc7-8f08-47d7-89cb-baa3f7a1f272}
   Action Gr05Auto_eAxisClamp1InPipeEndPos_Action: Id {02437d06-368c-46ab-b97e-751dd7ee46d1}
   Action Gr05Auto_eAxisClamp1InPipeEndPos_Exit: Id {010e0099-2b89-4bbf-a561-caf5a0e95b21}
   Action Gr05Auto_eAxisClamp1InPos_Exit: Id {d5857da8-10ea-4615-acb6-caa53af139cc}
   Action Gr05Auto_eAxisClamp1InPos2_Exit: Id {447f4946-7b9d-47b6-8988-b094f8f70f11}
   Action Gr05Auto_eAxisClamp1InPos2Err_Entry: Id {67a7eb8f-cc21-4a2a-958e-094230f470c6}
   Action Gr05Auto_eAxisClamp1InPosErr_Entry: Id {1f8f0153-e9b0-480c-a34d-00c2505183a0}
   Action Gr05Auto_eAxisClamp1InSawBandPos_Exit: Id {a1ce9bc2-95ab-4922-9439-6b141e3588f7}
   Action Gr05Auto_eAxisClamp1InSawBandPosErr_Entry: Id {21f85646-0df1-460d-be10-4ec4635e9559}
   Action Gr05Auto_eAxisClamp1MoveAbsPipeEnde_Entry: Id {a0101a6c-31a1-43c3-a722-76f0baeda599}
   Action Gr05Auto_eAxisClamp1MoveAbsPipeEnde_Exit: Id {ec425a8e-f2a1-44e3-8922-f107615160fb}
   Action Gr05Auto_eAxisClamp1MoveAbsPipeEndeErr_Entry: Id {21853957-6bde-4e98-b330-6d97e5247b95}
   Action Gr05Auto_eAxisClamp1MoveToBackPos_Entry: Id {e265f354-3adf-4b1b-a593-e700b87d49f9}
   Action Gr05Auto_eAxisClamp1MoveToBackPosErr_Entry: Id {676edf1c-3706-4631-914d-22510e6f13d7}
   Action Gr05Auto_eAxisClamp1MoveToPos_Action: Id {a26a0dce-c76a-4711-be64-a08c8aa22c56}
   Action Gr05Auto_eAxisClamp1MoveToPos_Entry: Id {ecc447ef-c0f8-470d-ac82-be64f50fa825}
   Action Gr05Auto_eAxisClamp1MoveToPos2_Entry: Id {a86c68ce-4588-492a-b688-fd2f40e0f9a9}
   Action Gr05Auto_eAxisClamp1MoveToPos2Err_Entry: Id {e9c77a3a-e884-499f-8e39-ffaab5eeaccf}
   Action Gr05Auto_eAxisClamp1MoveToPosErr_Entry: Id {ca8224d6-1b22-4e4c-8c8e-2294d0d8c087}
   Action Gr05Auto_eAxisClamp1MoveToSawBandPos_Entry: Id {2eef4d10-19d2-42cf-93b6-58293ec388af}
   Action Gr05Auto_eAxisClamp1MoveToSawBandPosErr_Entry: Id {ba50b007-a133-476c-b3ab-5fc9f431f3ca}
   Action Gr05Auto_eAxisClamp1MoveVeloPipeBegin_Entry: Id {e699aee6-0300-4c07-a2a6-49007f5a09ad}
   Action Gr05Auto_eAxisClamp1MoveVeloPipeBeginErr_Entry: Id {78790b27-2540-4b02-964c-8637b813a519}
   Action Gr05Auto_eAxisClamp1MoveVeloPipeEnd_Entry: Id {32c1370d-4185-4d69-b7cf-d77dcbdff087}
   Action Gr05Auto_eAxisClamp1MoveVeloPipeEndErr_Entry: Id {ab0564e6-3d4a-42bf-aef7-cdf399171da7}
   Action Gr05Auto_eAxisClamp1Stop_2_Entry: Id {4788458a-91dc-49dd-85e9-1a28e841f245}
   Action Gr05Auto_eAxisClamp1Stop_Entry: Id {2c316997-9a2d-47bc-a0cb-e4d4dc5c0044}
   Action Gr05Auto_eAxisClamp1StopErr_2_Entry: Id {03905c0e-891e-4242-bf65-f20e95932e92}
   Action Gr05Auto_eAxisClamp1StopErr_Entry: Id {07788e5a-f1c9-405c-8725-191e9ad33104}
   Action Gr05Auto_eAxisClamp2InPos_Exit: Id {d585134b-7419-4d8f-8668-f5c98c079cc5}
   Action Gr05Auto_eAxisClamp2InPos2_Exit: Id {8d051bda-26ed-4bef-93ed-dd5497a7903f}
   Action Gr05Auto_eAxisClamp2InPos2Err_Entry: Id {a16c5bc0-785f-43cd-891a-6f89e3d9952d}
   Action Gr05Auto_eAxisClamp2InPosErr_Entry: Id {df1ecd55-6106-4267-ad38-f95bb237d40b}
   Action Gr05Auto_eAxisClamp2InSawBandPos_Exit: Id {d4345afb-4634-4cfb-903b-c43df2f9863b}
   Action Gr05Auto_eAxisClamp2InSawBandPosErr_Entry: Id {c7991712-0773-4cf5-8758-d968077fc7d5}
   Action Gr05Auto_eAxisClamp2InSawPos_Exit: Id {3698282c-eb3b-4737-a95a-d25262388aa3}
   Action Gr05Auto_eAxisClamp2InSawPosErr_Entry: Id {91e6d10d-d2b2-445c-8a56-efc64929a08b}
   Action Gr05Auto_eAxisClamp2MoveSawPos_Entry: Id {2f51a821-8757-48c8-befb-2e15b0a9c27e}
   Action Gr05Auto_eAxisClamp2MoveSawPosErr_Entry: Id {d01e3b9b-39fb-4019-bfa7-8b24ed2512ac}
   Action Gr05Auto_eAxisClamp2MoveToPos_Entry: Id {564b843a-143b-4f2c-b16d-cf8e822d734b}
   Action Gr05Auto_eAxisClamp2MoveToPos2_Entry: Id {dee9280e-ac7e-48cd-a916-68ade5b1e999}
   Action Gr05Auto_eAxisClamp2MoveToPos2Err_Entry: Id {6595b859-6d9e-4a6d-9a76-9ea032ca9493}
   Action Gr05Auto_eAxisClamp2MoveToPosErr_Entry: Id {d3bf44ef-5107-4021-b4c3-6a2ddbc1c78f}
   Action Gr05Auto_eAxisClamp2MoveToSawBandPos_Entry: Id {e8610859-81ea-414b-b5c1-121b70fe0966}
   Action Gr05Auto_eAxisClamp2MoveToSawBandPosErr_Entry: Id {74b45e41-57db-4495-a1b9-1e7285bc0811}
   Action Gr05Auto_eChkAxisClamp1MoveToBackPos_Entry: Id {c15f677a-24fd-4755-8ab3-a5e3d41c95d0}
   Action Gr05Auto_eChkAxisClamp1MoveToBackPos_Exit: Id {e48deca1-f7b0-41b7-a2f3-60835af9fee8}
   Action Gr05Auto_eChkWorkArea_Entry: Id {33352e18-62da-49c8-8740-f93b31518d88}
   Action Gr05Auto_eClamp12Open_Entry: Id {25d99cf5-deef-4ef3-9012-b97b1be136f2}
   Action Gr05Auto_eClamp12Open_Exit: Id {bd9f8848-ce7f-4722-9a4c-b0b4d9ee2d4d}
   Action Gr05Auto_eClamp1Close_Entry: Id {72183c9e-dc9e-49b7-a69a-54fe28f1f6ec}
   Action Gr05Auto_eClamp1Close_Exit: Id {4b28f930-a1bb-42e8-913e-508ce8030708}
   Action Gr05Auto_eClamp1Close2_Entry: Id {528de016-69e2-426f-9bc1-8460d76e5a4c}
   Action Gr05Auto_eClamp1Close2_Exit: Id {ea079475-ff0a-4b2c-9f0a-7abc9d24e173}
   Action Gr05Auto_eClamp1Close2Err_Entry: Id {243046a1-4045-43c9-a4e2-ae5d218699c3}
   Action Gr05Auto_eClamp1Close3_Entry: Id {6729ea2c-9bf8-4346-a6b8-d8a99a5f6745}
   Action Gr05Auto_eClamp1Close3_Exit: Id {32a706df-f003-4226-a5c6-ad22f46eba73}
   Action Gr05Auto_eClamp1Close3Err_Entry: Id {ed0eb64f-b294-4bb5-8737-5fff4ee47b35}
   Action Gr05Auto_eClamp1CloseErr_Entry: Id {c4adbdf8-0350-421a-bf0a-8f022d3d4796}
   Action Gr05Auto_eClamp1Open_Entry: Id {89beb1bd-91ad-426b-884e-c750ed7ec7d3}
   Action Gr05Auto_eClamp1Open_Exit: Id {47f7eb34-7693-4b6a-bbd2-0aee97a8cde2}
   Action Gr05Auto_eClamp1Open2Err_Entry: Id {62a50412-8b9e-4667-b82c-d270259cbb16}
   Action Gr05Auto_eClamp1OpenErr_Entry: Id {9a731d93-6a99-4964-a7d3-3a93b297f220}
   Action Gr05Auto_eClamp2Close_Entry: Id {aadb4727-179a-47ae-a454-f444ca84ff5b}
   Action Gr05Auto_eClamp2Close_Exit: Id {7f93481f-14ba-4f9f-b8bd-34ce4266271e}
   Action Gr05Auto_eClamp2CloseErr_Entry: Id {97146f8b-2272-4f68-9758-bf4784ee4e72}
   Action Gr05Auto_eClamp2Err_Entry: Id {6a952772-b017-4ee7-bc33-1da17f483437}
   Action Gr05Auto_eClamp2Open_Entry: Id {e69eb5ea-9054-4a61-afc6-2e880d34a3b8}
   Action Gr05Auto_eClamp2Open_Exit: Id {6a61fe58-b92f-4428-b287-0dfa6509d2aa}
   Action Gr05Auto_eClamp2Open1_Entry: Id {d329d572-6934-4333-9c51-90f499b42085}
   Action Gr05Auto_eClamp2Open1_Exit: Id {35cf07fb-2f81-4b27-9f0e-edc0603fe2b7}
   Action Gr05Auto_eClamp2Open1Err_Entry: Id {d1e99eda-1446-4ef3-8560-d0d529c24baf}
   Action Gr05Auto_eClamp2Open2Err_Entry: Id {a8fc3ca8-a504-4154-bb40-5e4c23464b4e}
   Action Gr05Auto_eClamp2Open3_Entry: Id {e0cd2334-91c9-4838-b0d5-84d8dca1c8d2}
   Action Gr05Auto_eClamp2Open3_Exit: Id {a8ebbeb3-57d6-4f2f-8f8f-c0c53991025e}
   Action Gr05Auto_eClamp2Open3Err_Entry: Id {7fd9181b-424e-47ff-9b7a-f19a378090c1}
   Action Gr05Auto_eClamp2OpenErr_Entry: Id {91e23f9e-13d2-4baa-8f47-37da7eb28d04}
   Action Gr05Auto_eClamp2Slide_Entry: Id {1b509614-5c8f-4072-92f1-f9c1f7248f9e}
   Action Gr05Auto_eClamp2Slide_Exit: Id {4c541fdc-aaa8-4bf3-8748-213803fbb427}
   Action Gr05Auto_eCollisionDetectedErr_Entry: Id {4d44d703-5490-422c-8fa4-937cd67571c1}
   Action Gr05Auto_eCollisionDetectedErr_Exit: Id {968e4e1a-0728-4257-8ad5-ca47403f9ccf}
   Action Gr05Auto_eDone_Entry: Id {1c745913-da3c-4f44-829a-3cf26310d759}
   Action Gr05Auto_eDone_Exit: Id {7ab109ae-4201-4fc3-b6f9-c5034bbf4897}
   Action Gr05Auto_eError_Entry: Id {8ff6a727-cb1f-40d8-9399-c0a1f0edc994}
   Action Gr05Auto_eError_Exit: Id {d5f44c68-5af0-41b9-824d-baf54a1fb0b2}
   Action Gr05Auto_eGetClamp1ActPos_01_Entry: Id {94c0fcbb-e02d-4852-9da7-5ea490b3f11d}
   Action Gr05Auto_eGetClamp1ActPos_02_Entry: Id {def876cc-eecb-4aa5-9dc6-ca3227bcfc02}
   Action Gr05Auto_eGetClamp1ActPos_03_Entry: Id {64795166-20bb-4a1c-9c63-6cd05bae47ae}
   Action Gr05Auto_eGetClamp1ActPos_04_Entry: Id {f500f5c2-f162-4e2c-a6f2-ac3316910f9a}
   Action Gr05Auto_eGetClamp1ActPos_05_Entry: Id {6ac5818d-c157-4f43-adb0-ca0be23cb02b}
   Action Gr05Auto_eGetClamp1ActPos_06_Entry: Id {10e52d9c-0a10-4f33-852d-f75074e4270b}
   Action Gr05Auto_eGetClamp1ActPos_Entry: Id {3729689b-c43c-49cb-823e-b8a98e2f0273}
   Action Gr05Auto_eGetClamp2ActPos_Entry: Id {8f51bb36-e3aa-4108-b809-c75d7ad21bb0}
   Action Gr05Auto_eGetProcessPara_Entry: Id {22f4a980-7d39-48f7-b450-d1793048e058}
   Action Gr05Auto_eRemovalBandErr_Entry: Id {cbb27a62-3f2f-4868-991f-db92473c6f01}
   Action Gr05Auto_eSawbandStart_Entry: Id {020eb7db-6d27-4c83-9b2b-f5583953e4b6}
   Action Gr05Auto_eSawbandStart_Exit: Id {57ff5e58-fe83-4b98-95e5-a6936022fb58}
   Action Gr05Auto_eSawingLengthCorrection_Entry: Id {9c418063-f092-4e75-95d0-e602933e46bc}
   Action Gr05Auto_eSawingReq_Entry: Id {c426ed76-57e2-452f-9d36-e766017cfdd0}
   Action Gr05Auto_eSawingReq_Exit: Id {76d1889a-60fc-4fd2-b5ea-13bf0109cf3c}
   Action Gr05Auto_eSlideDown_Entry: Id {a44d763e-9492-4915-b7f5-140352186076}
   Action Gr05Auto_eSlideDownErr_Entry: Id {475aa099-df50-4844-8f0f-e6e5ee771ed8}
   Action Gr05Auto_eSlideUpErr_Entry: Id {82559d77-26fa-4ea5-a94e-2275adaf32e9}
   Action Gr05Auto_eTransportAck_Exit: Id {78aeef6f-07e6-4252-bcb1-58d6013bc1e7}
   Action Gr05Auto_eWfAxisClamp1MoveAbsPipeEnde_Exit: Id {4dab6c74-788e-403c-b963-cf04d4fbec81}
   Action Gr05Auto_eWfAxisClamp1MoveAbsPipeEndeErr_Entry: Id {f4fc9039-2dad-4ea1-945e-a28a4c7d83c3}
   Action Gr05Auto_eWfAxisClamp1MoveVeloPipeBegin_Exit: Id {170e38a7-3c2d-44a5-bbcb-696debfd69af}
   Action Gr05Auto_eWfAxisClamp1MoveVeloPipeBeginErr_Entry: Id {cd8cf5d5-7040-4bce-8fce-f1e806a9d4f6}
   Action Gr05Auto_eWfAxisClamp1MoveVeloPipeEnd_Exit: Id {d7b933c6-c2c7-4454-a675-bd10502400ab}
   Action Gr05Auto_eWfAxisClamp1MoveVeloPipeEndErr_Entry: Id {7f8750b2-eb21-4071-95e5-afae5d1c54c2}
   Action Gr05Auto_eWfAxisClamp1Stop_2_Exit: Id {37bedc03-1a5d-47d6-acdd-9d4526947790}
   Action Gr05Auto_eWfAxisClamp1Stop_Exit: Id {edaeb31f-2806-4e16-b9d3-0173a80d8f61}
   Action Gr05Auto_eWfAxisClamp1StopErr_2_Entry: Id {6f857205-34a8-4dfc-b879-93376445566c}
   Action Gr05Auto_eWfAxisClamp1StopErr_Entry: Id {8c9784ac-8c69-47be-9db5-f9ce3998c119}
   Action Gr05Auto_eWfPipeBeginNoDetectedError_Entry: Id {59aa8b79-44d2-4253-97ff-cec75c460835}
   Action Gr05Auto_eWfPipeBeginNoDetectedError_Exit: Id {60842bba-c9e9-40b8-af45-960cd0009ccc}
   Action Gr05Auto_eWfPipeBeginNoDetectedWarrning_Entry: Id {3b44d596-f122-4735-8f47-e49b74d78f45}
   Action Gr05Auto_eWfPipeBeginNoDetectedWarrning_Exit: Id {a66a2d82-b8b4-4733-8b01-d00f61bda4bc}
   Action Gr05Auto_eWfPipeEndNoDetectedErr_Entry: Id {8011e142-bd4c-41e8-a55c-7e877bdf0b9f}
   Action Gr05Auto_eWfPipeEndNoDetectedErr_Exit: Id {46b0ed65-6d3a-4b14-9012-9ca07481e536}
   Action Gr05Auto_eWfTransportReq_Exit: Id {07162ad3-42cb-4c70-8ff4-8a4787adb266}
   Action Init_Action: Id {73020b56-24e3-4ee9-bad5-4ae590e36ed2}
   Action Init_Exit: Id {85d4513c-b205-4f2e-89c9-544ae04dd426}
   Transition SafetyDistEnable: Id {d0ec5b99-d67e-4fe1-8932-a0722f74e568}
   Transition SafetyDistEnable_1: Id {b1fda3e7-c5fa-48d9-8a77-5c2022df07d4}
   Transition Trans: Id {3ddce4b7-11c1-4ed2-80c1-5f760c49db1d}
   Transition Trans_1: Id {05cc9c8b-bd71-4e38-b12e-5fde4340a0b8}
   Transition Trans_10: Id {17f506b3-00a9-476b-8d71-4695e39f48d7}
   Transition Trans_100: Id {dac33c7f-d08f-42ba-96d3-17a32f722bfb}
   Transition Trans_101: Id {3644a6e6-a052-4fdc-821d-4fb05e9e1b2f}
   Transition Trans_11: Id {9acd7d56-70f4-41e3-8fac-4f2fa8f8fd83}
   Transition Trans_12: Id {b29ccfdc-a253-4455-b478-8a89802d1ed4}
   Transition Trans_13: Id {4ef7619e-fc0d-46d1-9f72-6ba00625f868}
   Transition Trans_14: Id {6b3b904d-609e-4f74-887e-c4a332baa76c}
   Transition Trans_15: Id {aa107144-0995-48c2-b1be-5f0931f705ba}
   Transition Trans_16: Id {8a47e3a0-2dcc-4eaf-96ec-06ec88024399}
   Transition Trans_17: Id {23d1c92a-a5fb-41d3-a543-090ffeaf9f25}
   Transition Trans_18: Id {d2263dee-a359-4264-a422-9a229513cfbb}
   Transition Trans_19: Id {fee0b0bd-475f-496b-885b-7880f3b10418}
   Transition Trans_2: Id {51af1fe4-769d-4e24-8970-e888a7f42fee}
   Transition Trans_20: Id {9c2d4755-9e3d-4562-91e0-fafa709f22f6}
   Transition Trans_21: Id {2f365ad8-931c-4a9d-b293-e29bb5bec034}
   Transition Trans_22: Id {9d0dfb6f-c662-436b-b601-c07d13765bd8}
   Transition Trans_23: Id {14a4469b-942c-419f-a123-cfc462a58e06}
   Transition Trans_24: Id {f534d3b3-f15c-436b-8ba5-1dd49a3a8adf}
   Transition Trans_25: Id {29fd3c2b-3925-412d-91e0-c147f8661701}
   Transition Trans_26: Id {300aff37-1920-46e8-bfc4-a457e570384e}
   Transition Trans_27: Id {954dae76-5937-4d76-8740-8643c3f66dc7}
   Transition Trans_28: Id {75213184-ede9-427f-ba25-c168bd6f0566}
   Transition Trans_29: Id {d6bee61e-8eda-4ffe-83a7-860a90cb9ab6}
   Transition Trans_3: Id {f2832df7-ceb3-4aee-b1db-bd2e990a9715}
   Transition Trans_30: Id {dae48976-0e1f-4321-a07a-745529641746}
   Transition Trans_31: Id {6a1fa657-8587-40fa-8370-d6eeb93975ed}
   Transition Trans_32: Id {362dd6ce-6a41-47cf-8073-0062f6f7fc4c}
   Transition Trans_33: Id {80223384-cc75-4628-a1ca-27aa74a27ceb}
   Transition Trans_34: Id {1bb3413f-3a0f-4a58-a7aa-cbcb580e8c73}
   Transition Trans_35: Id {15510543-586d-461b-88e1-866a042414c6}
   Transition Trans_36: Id {78b535a0-759b-43d3-b1b9-94b532d28884}
   Transition Trans_37: Id {8cc0a4fa-9ee1-45c5-8585-0612d52508a5}
   Transition Trans_38: Id {b53eee66-2713-4295-ae54-c97af9237b0a}
   Transition Trans_39: Id {e9c255fb-5086-4480-bdac-63238da542d3}
   Transition Trans_4: Id {e99af99f-1de7-4a99-b049-2549e48732a4}
   Transition Trans_40: Id {afbf47f0-b10b-472c-bddd-a3fd6463fc71}
   Transition Trans_41: Id {864bfcfa-a754-46a1-b9fb-3b50f74807cc}
   Transition Trans_42: Id {8ceb7b10-6f0c-472e-83f2-fbe351a9cd01}
   Transition Trans_43: Id {37644647-fb0b-4d46-a4c2-5d95b541800d}
   Transition Trans_44: Id {bf6b613f-7154-4b3f-bf51-324b4f1f262c}
   Transition Trans_45: Id {0ab1eddb-7c04-4f68-a470-72fcef43ae7c}
   Transition Trans_46: Id {e1e3b099-39ab-48eb-ae4b-1ad5759431d9}
   Transition Trans_47: Id {9476b89a-8f35-4799-83d4-03e82138e902}
   Transition Trans_48: Id {d89d8a4e-c6c4-4409-ba7b-7e5c9429613e}
   Transition Trans_49: Id {6dbbcb69-cb96-4fc1-98a6-2bb80ae8d84c}
   Transition Trans_5: Id {e47b9578-df07-4e12-8306-26aaa0a6ecf0}
   Transition Trans_50: Id {76ceeb70-4452-4a40-9c42-b601ef241637}
   Transition Trans_51: Id {f35dacd5-e0d1-4451-bfd5-086652e73351}
   Transition Trans_52: Id {6e75a62e-8497-4508-8ef5-08e25c99fe6b}
   Transition Trans_53: Id {869e56c1-6eb5-4878-9e66-7cb560c5fcb3}
   Transition Trans_54: Id {cae10fe3-e081-4350-b242-745fd4227805}
   Transition Trans_55: Id {08ac33b2-5e1f-4639-a09a-883298509093}
   Transition Trans_56: Id {71ca1fcf-2265-417d-aa2a-27d911069c78}
   Transition Trans_57: Id {b06078fa-6b6f-48c2-bd1c-8a764f46e477}
   Transition Trans_58: Id {c1bdcb17-a11e-4f98-9e5b-c240bf65e069}
   Transition Trans_59: Id {011ce394-7eda-4a73-9816-2ca7149ee80a}
   Transition Trans_6: Id {8e5b9af4-6320-4af4-967d-8615b8e6dabc}
   Transition Trans_60: Id {971986f1-afa8-4631-a150-12b43643526c}
   Transition Trans_61: Id {049c2c78-8b06-48b1-86b1-659bce566ca4}
   Transition Trans_62: Id {ab1c7d03-d8ce-4c4f-bc2a-2f89b17fe068}
   Transition Trans_63: Id {e4cef4bf-9afd-4fe2-a6b4-5e76e2d98e3b}
   Transition Trans_64: Id {2cc9c9e4-4837-49d4-b31d-2f987d2761b6}
   Transition Trans_65: Id {1fd3af44-cc34-4fe9-a3fe-0651e24799b9}
   Transition Trans_66: Id {dd2ddf4b-0db4-4fb6-88ac-aa712741aa0d}
   Transition Trans_67: Id {0b733374-9c56-4a18-9450-8350918fb205}
   Transition Trans_68: Id {c95cf03b-e98e-4821-828f-a4723c836fda}
   Transition Trans_69: Id {02611326-3bf6-4659-a5f1-06d69a7f86ca}
   Transition Trans_7: Id {d2cc99d2-2baa-4c66-8c61-1574092b01d9}
   Transition Trans_70: Id {147e7842-75d8-4982-99be-4acd026e049c}
   Transition Trans_71: Id {b5494e10-3c0d-4c65-8350-5ad04d31aa3c}
   Transition Trans_72: Id {b01024d1-36ef-4dfc-a55e-ff07b835c43c}
   Transition Trans_73: Id {24f62e30-d7db-4e81-9a6a-702321be4f16}
   Transition Trans_74: Id {007a540b-c73f-4993-9237-b79ca7773d1e}
   Transition Trans_75: Id {87cd0eb4-ee69-4d2f-b286-111fa5b31793}
   Transition Trans_76: Id {00915d48-24a0-46d3-ab6a-a85c3ee66421}
   Transition Trans_77: Id {966a3c91-99ab-4190-b151-9b0d5b19940d}
   Transition Trans_78: Id {ac882a59-53a7-426b-92b0-75861867283b}
   Transition Trans_79: Id {190c7633-18eb-4ce8-8931-f7432173c920}
   Transition Trans_8: Id {26204b5a-f781-4ed1-8b43-32f9c984f456}
   Transition Trans_80: Id {d07f8a6a-e3fa-4af0-88fb-f69c7c03dbeb}
   Transition Trans_81: Id {bf437b9f-c399-42bf-bf49-0a40301a341c}
   Transition Trans_82: Id {2ff399e3-f641-4568-97c7-4dcc8d85be82}
   Transition Trans_83: Id {b018ba08-9f31-4896-bda9-9a71d18f25a2}
   Transition Trans_84: Id {dbfce89f-bdb4-4dcc-804c-74e75a2eab1a}
   Transition Trans_85: Id {11025e17-f8e6-4f8e-9b2f-4ea1b24bf397}
   Transition Trans_86: Id {62981d2b-bc79-4b59-a3c5-a49a8831a407}
   Transition Trans_87: Id {f750845b-a2db-4101-b0a6-8d4f4e052dc6}
   Transition Trans_88: Id {1f525d0d-441f-4bd4-ae63-f0b136cc968f}
   Transition Trans_89: Id {5c8ec368-d265-4704-b238-a0e7fae312fe}
   Transition Trans_9: Id {19aed697-83cf-49ad-8f74-33fcabc9994e}
   Transition Trans_90: Id {549ff61b-e991-48a7-a0dd-7ab7863fb678}
   Transition Trans_91: Id {8779a092-aca4-4019-b1f3-a147d5c451c0}
   Transition Trans_92: Id {2a6521bf-6649-4010-912a-b9ef18a77915}
   Transition Trans_93: Id {3272d9dc-327c-4690-b0f1-e4c705aa3e6c}
   Transition Trans_94: Id {e0aac3cc-7470-4f83-a063-26d79d5b1755}
   Transition Trans_95: Id {bd63753f-86cd-4c09-b2e0-cd6fc7ffdc90}
   Transition Trans_96: Id {a7529c8d-217d-4d53-9229-2f2b5658353b}
   Transition Trans_97: Id {46072854-4d14-4957-9545-eac42c7c290d}
   Transition Trans_98: Id {902da588-ed42-446b-8e2f-6fc55a684d64}
   Transition Trans_99: Id {2125bfec-2247-4914-97bc-0569bc2ca9fe} *)
